    RC4_Receive_PDO_Mapping_Physical_outputs_60FE_01 : UDINT;
    RC4_Transmit_PDO_Mapping_StatusWord_6041_00 : UINT;
    RC4_Transmit_PDO_Mapping_Position_actual_value_6064_00 : DINT;
    RC4_Transmit_PDO_Mapping_Mode_of_operation_display_6061_00 : SINT;
    RC4_Transmit_PDO_Mapping_Following_error_actual_valu_60F4_00 : DINT;
    RC4_Transmit_PDO_Mapping_Torque_actual_value_6077_00 : INT;
    RC4_Transmit_PDO_Mapping_Digital_inputs_60FD_00 : UDINT;
    RC4_Transmit_PDO_Mapping_Error_code_603F_00 : UINT;
    RC5_Receive_PDO_Mapping_ControlWord_6040_00 : UINT;
    RC5_Receive_PDO_Mapping_Target_Position_607A_00 : DINT;
    RC5_Receive_PDO_Mapping_Mode_of_operation_6060_00 : SINT;
    RC5_Receive_PDO_Mapping_Profile_velocity_6081_00 : UDINT;
    RC5_Receive_PDO_Mapping_Profile_acceleration_6083_00 : UDINT;
    RC5_Receive_PDO_Mapping_Profile_deceleration_6084_00 : UDINT;
    RC5_Receive_PDO_Mapping_Physical_outputs_60FE_01 : UDINT;
    RC5_Transmit_PDO_Mapping_StatusWord_6041_00 : UINT;
    RC5_Transmit_PDO_Mapping_Position_actual_value_6064_00 : DINT;
    RC5_Transmit_PDO_Mapping_Mode_of_operation_display_6061_00 : SINT;
    RC5_Transmit_PDO_Mapping_Following_error_actual_valu_60F4_00 : DINT;
    RC5_Transmit_PDO_Mapping_Torque_actual_value_6077_00 : INT;
    RC5_Transmit_PDO_Mapping_Digital_inputs_60FD_00 : UDINT;
    RC5_Transmit_PDO_Mapping_Error_code_603F_00 : UINT;
    RC6_Receive_PDO_Mapping_ControlWord_6040_00 : UINT;
    RC6_Receive_PDO_Mapping_ControlWord_6040_00_1 : UINT;
    RC6_Receive_PDO_Mapping_Target_Position_607A_00 : DINT;
    RC6_Receive_PDO_Mapping_Mode_of_operation_6060_00 : SINT;
    RC6_Receive_PDO_Mapping_Profile_velocity_6081_00 : UDINT;
    RC6_Receive_PDO_Mapping_Profile_acceleration_6083_00 : UDINT;
    RC6_Receive_PDO_Mapping_Profile_deceleration_6084_00 : UDINT;
    RC6_Receive_PDO_Mapping_Physical_outputs_60FE_01 : UDINT;
    RC6_Transmit_PDO_Mapping_StatusWord_6041_00 : UINT;
    RC6_Transmit_PDO_Mapping_Position_actual_value_6064_00 : DINT;
    RC6_Transmit_PDO_Mapping_Mode_of_operation_display_6061_00 : SINT;
    RC6_Transmit_PDO_Mapping_Following_error_actual_valu_60F4_00 : DINT;
    RC6_Transmit_PDO_Mapping_Torque_actual_value_6077_00 : INT;
    RC6_Transmit_PDO_Mapping_Digital_inputs_60FD_00 : UDINT;
    RC6_Transmit_PDO_Mapping_Error_code_603F_00 : UINT;
    RCON1_OUT : ARRAY[1..6] OF ST_RCON_Direct_OUT_Axis;  (* RCON1 6軸分 PLC→RCON 指令（内部変数・通信変換は別途） *)
    RCON1_IN : ARRAY[1..6] OF ST_RCON_Direct_IN_Axis;  (* RCON1 6軸分 RCON→PLC 取得値・状態（内部変数・通信変換は別途） *)
    RCON1_SpeedUnit_mm_s : LREAL;  (* RCON1 速度の1カウント量mm/s。実機設定1.0または0.1を確認。未確認・0では使用しない。 *)
    RCON1_OUT_GwControl0Raw : UINT;  (* RCON1 PLC→RCON 【OUT00】共通 ゲートウェイ制御信号0（MON等）（未割付・直接数値指定の設計用） *)
    RCON1_OUT_GwControl1ReservedRaw : UINT;  (* RCON1 PLC→RCON 【OUT01】共通 ゲートウェイ制御信号1（予約・使用禁止）（未割付・直接数値指定の設計用） *)
    RCON1_OUT_ReservedOut02Raw : UINT;  (* RCON1 PLC→RCON 【OUT02】共通 共通予約領域（使用禁止・占有あり）（未割付・直接数値指定の設計用） *)
    RCON1_OUT_ReservedOut03Raw : UINT;  (* RCON1 PLC→RCON 【OUT03】共通 共通予約領域（使用禁止・占有あり）（未割付・直接数値指定の設計用） *)
    RCON1_OUT_ReservedOut04Raw : UINT;  (* RCON1 PLC→RCON 【OUT04】共通 共通予約領域（使用禁止・占有あり）（未割付・直接数値指定の設計用） *)
    RCON1_OUT_ReservedOut05Raw : UINT;  (* RCON1 PLC→RCON 【OUT05】共通 共通予約領域（使用禁止・占有あり）（未割付・直接数値指定の設計用） *)
    RCON1_OUT_ReservedOut06Raw : UINT;  (* RCON1 PLC→RCON 【OUT06】共通 共通予約領域（使用禁止・占有あり）（未割付・直接数値指定の設計用） *)
    RCON1_OUT_ReservedOut07Raw : UINT;  (* RCON1 PLC→RCON 【OUT07】共通 共通予約領域（使用禁止・占有あり）（未割付・直接数値指定の設計用） *)
    RCON1_OUT_Axis1_TargetPosLoRaw : UINT;  (* RCON1 PLC→RCON 【OUT08】1軸目（No.0） 目標位置 下位ワード（未割付・直接数値指定の設計用） *)
    RCON1_OUT_Axis1_TargetPosHiRaw : UINT;  (* RCON1 PLC→RCON 【OUT09】1軸目（No.0） 目標位置 上位ワード（未割付・直接数値指定の設計用） *)
    RCON1_OUT_Axis1_PositionBandLoRaw : UINT;  (* RCON1 PLC→RCON 【OUT10】1軸目（No.0） 位置決め幅 下位ワード（未割付・直接数値指定の設計用） *)
    RCON1_OUT_Axis1_PositionBandHiRaw : UINT;  (* RCON1 PLC→RCON 【OUT11】1軸目（No.0） 位置決め幅 上位ワード（未割付・直接数値指定の設計用） *)
    RCON1_OUT_Axis1_SpeedRaw : UINT;  (* RCON1 PLC→RCON 【OUT12】1軸目（No.0） 速度指令（未割付・直接数値指定の設計用） *)
    RCON1_OUT_Axis1_AccDecRaw : UINT;  (* RCON1 PLC→RCON 【OUT13】1軸目（No.0） 加減速度指令（加速・減速共通）（未割付・直接数値指定の設計用） *)
    RCON1_OUT_Axis1_PushLimitRaw : UINT;  (* RCON1 PLC→RCON 【OUT14】1軸目（No.0） 押付け電流制限値（未割付・直接数値指定の設計用） *)
    RCON1_OUT_Axis1_ControlRaw : UINT;  (* RCON1 PLC→RCON 【OUT15】1軸目（No.0） 軸制御信号（DSTR・SON等）（未割付・直接数値指定の設計用） *)
    RCON1_OUT_Axis2_TargetPosLoRaw : UINT;  (* RCON1 PLC→RCON 【OUT16】2軸目（No.1） 目標位置 下位ワード（未割付・直接数値指定の設計用） *)
    RCON1_OUT_Axis2_TargetPosHiRaw : UINT;  (* RCON1 PLC→RCON 【OUT17】2軸目（No.1） 目標位置 上位ワード（未割付・直接数値指定の設計用） *)
    RCON1_OUT_Axis2_PositionBandLoRaw : UINT;  (* RCON1 PLC→RCON 【OUT18】2軸目（No.1） 位置決め幅 下位ワード（未割付・直接数値指定の設計用） *)
    RCON1_OUT_Axis2_PositionBandHiRaw : UINT;  (* RCON1 PLC→RCON 【OUT19】2軸目（No.1） 位置決め幅 上位ワード（未割付・直接数値指定の設計用） *)
    RCON1_OUT_Axis2_SpeedRaw : UINT;  (* RCON1 PLC→RCON 【OUT20】2軸目（No.1） 速度指令（未割付・直接数値指定の設計用） *)
    RCON1_OUT_Axis2_AccDecRaw : UINT;  (* RCON1 PLC→RCON 【OUT21】2軸目（No.1） 加減速度指令（加速・減速共通）（未割付・直接数値指定の設計用） *)
    RCON1_OUT_Axis2_PushLimitRaw : UINT;  (* RCON1 PLC→RCON 【OUT22】2軸目（No.1） 押付け電流制限値（未割付・直接数値指定の設計用） *)
    RCON1_OUT_Axis2_ControlRaw : UINT;  (* RCON1 PLC→RCON 【OUT23】2軸目（No.1） 軸制御信号（DSTR・SON等）（未割付・直接数値指定の設計用） *)
    RCON1_OUT_Axis3_TargetPosLoRaw : UINT;  (* RCON1 PLC→RCON 【OUT24】3軸目（No.2） 目標位置 下位ワード（未割付・直接数値指定の設計用） *)
    RCON1_OUT_Axis3_TargetPosHiRaw : UINT;  (* RCON1 PLC→RCON 【OUT25】3軸目（No.2） 目標位置 上位ワード（未割付・直接数値指定の設計用） *)
    RCON1_OUT_Axis3_PositionBandLoRaw : UINT;  (* RCON1 PLC→RCON 【OUT26】3軸目（No.2） 位置決め幅 下位ワード（未割付・直接数値指定の設計用） *)
    RCON1_OUT_Axis3_PositionBandHiRaw : UINT;  (* RCON1 PLC→RCON 【OUT27】3軸目（No.2） 位置決め幅 上位ワード（未割付・直接数値指定の設計用） *)
    RCON1_OUT_Axis3_SpeedRaw : UINT;  (* RCON1 PLC→RCON 【OUT28】3軸目（No.2） 速度指令（未割付・直接数値指定の設計用） *)
    RCON1_OUT_Axis3_AccDecRaw : UINT;  (* RCON1 PLC→RCON 【OUT29】3軸目（No.2） 加減速度指令（加速・減速共通）（未割付・直接数値指定の設計用） *)
    RCON1_OUT_Axis3_PushLimitRaw : UINT;  (* RCON1 PLC→RCON 【OUT30】3軸目（No.2） 押付け電流制限値（未割付・直接数値指定の設計用） *)
    RCON1_OUT_Axis3_ControlRaw : UINT;  (* RCON1 PLC→RCON 【OUT31】3軸目（No.2） 軸制御信号（DSTR・SON等）（未割付・直接数値指定の設計用） *)
    RCON1_OUT_Axis4_TargetPosLoRaw : UINT;  (* RCON1 PLC→RCON 【OUT32】4軸目（No.3） 目標位置 下位ワード（未割付・直接数値指定の設計用） *)
    RCON1_OUT_Axis4_TargetPosHiRaw : UINT;  (* RCON1 PLC→RCON 【OUT33】4軸目（No.3） 目標位置 上位ワード（未割付・直接数値指定の設計用） *)
    RCON1_OUT_Axis4_PositionBandLoRaw : UINT;  (* RCON1 PLC→RCON 【OUT34】4軸目（No.3） 位置決め幅 下位ワード（未割付・直接数値指定の設計用） *)
    RCON1_OUT_Axis4_PositionBandHiRaw : UINT;  (* RCON1 PLC→RCON 【OUT35】4軸目（No.3） 位置決め幅 上位ワード（未割付・直接数値指定の設計用） *)
    RCON1_OUT_Axis4_SpeedRaw : UINT;  (* RCON1 PLC→RCON 【OUT36】4軸目（No.3） 速度指令（未割付・直接数値指定の設計用） *)
    RCON1_OUT_Axis4_AccDecRaw : UINT;  (* RCON1 PLC→RCON 【OUT37】4軸目（No.3） 加減速度指令（加速・減速共通）（未割付・直接数値指定の設計用） *)
    RCON1_OUT_Axis4_PushLimitRaw : UINT;  (* RCON1 PLC→RCON 【OUT38】4軸目（No.3） 押付け電流制限値（未割付・直接数値指定の設計用） *)
    RCON1_OUT_Axis4_ControlRaw : UINT;  (* RCON1 PLC→RCON 【OUT39】4軸目（No.3） 軸制御信号（DSTR・SON等）（未割付・直接数値指定の設計用） *)
    RCON1_OUT_Axis5_TargetPosLoRaw : UINT;  (* RCON1 PLC→RCON 【OUT40】5軸目（No.4） 目標位置 下位ワード（未割付・直接数値指定の設計用） *)
    RCON1_OUT_Axis5_TargetPosHiRaw : UINT;  (* RCON1 PLC→RCON 【OUT41】5軸目（No.4） 目標位置 上位ワード（未割付・直接数値指定の設計用） *)
    RCON1_OUT_Axis5_PositionBandLoRaw : UINT;  (* RCON1 PLC→RCON 【OUT42】5軸目（No.4） 位置決め幅 下位ワード（未割付・直接数値指定の設計用） *)
    RCON1_OUT_Axis5_PositionBandHiRaw : UINT;  (* RCON1 PLC→RCON 【OUT43】5軸目（No.4） 位置決め幅 上位ワード（未割付・直接数値指定の設計用） *)
    RCON1_OUT_Axis5_SpeedRaw : UINT;  (* RCON1 PLC→RCON 【OUT44】5軸目（No.4） 速度指令（未割付・直接数値指定の設計用） *)
    RCON1_OUT_Axis5_AccDecRaw : UINT;  (* RCON1 PLC→RCON 【OUT45】5軸目（No.4） 加減速度指令（加速・減速共通）（未割付・直接数値指定の設計用） *)
    RCON1_OUT_Axis5_PushLimitRaw : UINT;  (* RCON1 PLC→RCON 【OUT46】5軸目（No.4） 押付け電流制限値（未割付・直接数値指定の設計用） *)
    RCON1_OUT_Axis5_ControlRaw : UINT;  (* RCON1 PLC→RCON 【OUT47】5軸目（No.4） 軸制御信号（DSTR・SON等）（未割付・直接数値指定の設計用） *)
    RCON1_OUT_Axis6_TargetPosLoRaw : UINT;  (* RCON1 PLC→RCON 【OUT48】6軸目（No.5） 目標位置 下位ワード（未割付・直接数値指定の設計用） *)
    RCON1_OUT_Axis6_TargetPosHiRaw : UINT;  (* RCON1 PLC→RCON 【OUT49】6軸目（No.5） 目標位置 上位ワード（未割付・直接数値指定の設計用） *)
    RCON1_OUT_Axis6_PositionBandLoRaw : UINT;  (* RCON1 PLC→RCON 【OUT50】6軸目（No.5） 位置決め幅 下位ワード（未割付・直接数値指定の設計用） *)
    RCON1_OUT_Axis6_PositionBandHiRaw : UINT;  (* RCON1 PLC→RCON 【OUT51】6軸目（No.5） 位置決め幅 上位ワード（未割付・直接数値指定の設計用） *)
    RCON1_OUT_Axis6_SpeedRaw : UINT;  (* RCON1 PLC→RCON 【OUT52】6軸目（No.5） 速度指令（未割付・直接数値指定の設計用） *)
    RCON1_OUT_Axis6_AccDecRaw : UINT;  (* RCON1 PLC→RCON 【OUT53】6軸目（No.5） 加減速度指令（加速・減速共通）（未割付・直接数値指定の設計用） *)
    RCON1_OUT_Axis6_PushLimitRaw : UINT;  (* RCON1 PLC→RCON 【OUT54】6軸目（No.5） 押付け電流制限値（未割付・直接数値指定の設計用） *)
    RCON1_OUT_Axis6_ControlRaw : UINT;  (* RCON1 PLC→RCON 【OUT55】6軸目（No.5） 軸制御信号（DSTR・SON等）（未割付・直接数値指定の設計用） *)
    RCON1_IN_GwStatus0Raw : UINT;  (* RCON1 RCON→PLC 【IN00】共通 ゲートウェイ状態信号0（未割付・直接数値指定の設計用） *)
    RCON1_IN_AxisLinkStatusRaw : UINT;  (* RCON1 RCON→PLC 【IN01】共通 ゲートウェイ状態信号1（軸No.0～15リンク状態）（未割付・直接数値指定の設計用） *)
    RCON1_IN_PowerStatus0Raw : UINT;  (* RCON1 RCON→PLC 【IN02】共通 電源ユニット状態信号0（未割付・直接数値指定の設計用） *)
    RCON1_IN_PowerStatus1Raw : UINT;  (* RCON1 RCON→PLC 【IN03】共通 電源ユニット状態信号1（未割付・直接数値指定の設計用） *)
    RCON1_IN_PowerStatus2Raw : UINT;  (* RCON1 RCON→PLC 【IN04】共通 電源ユニット状態信号2（未割付・直接数値指定の設計用） *)
    RCON1_IN_PowerStatus3Raw : UINT;  (* RCON1 RCON→PLC 【IN05】共通 電源ユニット状態信号3（未割付・直接数値指定の設計用） *)
    RCON1_IN_PowerStatus4MaintenanceRaw : UINT;  (* RCON1 RCON→PLC 【IN06】共通 電源ユニット状態信号4／軽故障メンテナンス（設定依存）（未割付・直接数値指定の設計用） *)
    RCON1_IN_ReservedIn07Raw : UINT;  (* RCON1 RCON→PLC 【IN07】共通 共通予約領域（使用禁止・占有あり）（未割付・直接数値指定の設計用） *)
    RCON1_IN_Axis1_ActualPosLoRaw : UINT;  (* RCON1 RCON→PLC 【IN08】1軸目（No.0） 現在位置 下位ワード（未割付・直接数値指定の設計用） *)
    RCON1_IN_Axis1_ActualPosHiRaw : UINT;  (* RCON1 RCON→PLC 【IN09】1軸目（No.0） 現在位置 上位ワード（未割付・直接数値指定の設計用） *)
    RCON1_IN_Axis1_CurrentLoRaw : UINT;  (* RCON1 RCON→PLC 【IN10】1軸目（No.0） 現在電流 下位ワード（PCは指令電流）（未割付・直接数値指定の設計用） *)
    RCON1_IN_Axis1_CurrentHiRaw : UINT;  (* RCON1 RCON→PLC 【IN11】1軸目（No.0） 現在電流 上位ワード（PCは指令電流）（未割付・直接数値指定の設計用） *)
    RCON1_IN_Axis1_ActualSpeedRaw : UINT;  (* RCON1 RCON→PLC 【IN12】1軸目（No.0） 現在速度（負方向は2の補数）（未割付・直接数値指定の設計用） *)
    RCON1_IN_Axis1_ReservedInRaw : UINT;  (* RCON1 RCON→PLC 【IN13】1軸目（No.0） 予約領域（使用禁止）（未割付・直接数値指定の設計用） *)
    RCON1_IN_Axis1_AlarmCodeRaw : UINT;  (* RCON1 RCON→PLC 【IN14】1軸目（No.0） アラームコード（簡易コードではない）（未割付・直接数値指定の設計用） *)
    RCON1_IN_Axis1_StatusRaw : UINT;  (* RCON1 RCON→PLC 【IN15】1軸目（No.0） 軸状態信号（PEND・SV等）（未割付・直接数値指定の設計用） *)
    RCON1_IN_Axis2_ActualPosLoRaw : UINT;  (* RCON1 RCON→PLC 【IN16】2軸目（No.1） 現在位置 下位ワード（未割付・直接数値指定の設計用） *)
    RCON1_IN_Axis2_ActualPosHiRaw : UINT;  (* RCON1 RCON→PLC 【IN17】2軸目（No.1） 現在位置 上位ワード（未割付・直接数値指定の設計用） *)
    RCON1_IN_Axis2_CurrentLoRaw : UINT;  (* RCON1 RCON→PLC 【IN18】2軸目（No.1） 現在電流 下位ワード（PCは指令電流）（未割付・直接数値指定の設計用） *)
    RCON1_IN_Axis2_CurrentHiRaw : UINT;  (* RCON1 RCON→PLC 【IN19】2軸目（No.1） 現在電流 上位ワード（PCは指令電流）（未割付・直接数値指定の設計用） *)
    RCON1_IN_Axis2_ActualSpeedRaw : UINT;  (* RCON1 RCON→PLC 【IN20】2軸目（No.1） 現在速度（負方向は2の補数）（未割付・直接数値指定の設計用） *)
    RCON1_IN_Axis2_ReservedInRaw : UINT;  (* RCON1 RCON→PLC 【IN21】2軸目（No.1） 予約領域（使用禁止）（未割付・直接数値指定の設計用） *)
    RCON1_IN_Axis2_AlarmCodeRaw : UINT;  (* RCON1 RCON→PLC 【IN22】2軸目（No.1） アラームコード（簡易コードではない）（未割付・直接数値指定の設計用） *)
    RCON1_IN_Axis2_StatusRaw : UINT;  (* RCON1 RCON→PLC 【IN23】2軸目（No.1） 軸状態信号（PEND・SV等）（未割付・直接数値指定の設計用） *)
    RCON1_IN_Axis3_ActualPosLoRaw : UINT;  (* RCON1 RCON→PLC 【IN24】3軸目（No.2） 現在位置 下位ワード（未割付・直接数値指定の設計用） *)
    RCON1_IN_Axis3_ActualPosHiRaw : UINT;  (* RCON1 RCON→PLC 【IN25】3軸目（No.2） 現在位置 上位ワード（未割付・直接数値指定の設計用） *)
    RCON1_IN_Axis3_CurrentLoRaw : UINT;  (* RCON1 RCON→PLC 【IN26】3軸目（No.2） 現在電流 下位ワード（PCは指令電流）（未割付・直接数値指定の設計用） *)
    RCON1_IN_Axis3_CurrentHiRaw : UINT;  (* RCON1 RCON→PLC 【IN27】3軸目（No.2） 現在電流 上位ワード（PCは指令電流）（未割付・直接数値指定の設計用） *)
    RCON1_IN_Axis3_ActualSpeedRaw : UINT;  (* RCON1 RCON→PLC 【IN28】3軸目（No.2） 現在速度（負方向は2の補数）（未割付・直接数値指定の設計用） *)
    RCON1_IN_Axis3_ReservedInRaw : UINT;  (* RCON1 RCON→PLC 【IN29】3軸目（No.2） 予約領域（使用禁止）（未割付・直接数値指定の設計用） *)
    RCON1_IN_Axis3_AlarmCodeRaw : UINT;  (* RCON1 RCON→PLC 【IN30】3軸目（No.2） アラームコード（簡易コードではない）（未割付・直接数値指定の設計用） *)
    RCON1_IN_Axis3_StatusRaw : UINT;  (* RCON1 RCON→PLC 【IN31】3軸目（No.2） 軸状態信号（PEND・SV等）（未割付・直接数値指定の設計用） *)
    RCON1_IN_Axis4_ActualPosLoRaw : UINT;  (* RCON1 RCON→PLC 【IN32】4軸目（No.3） 現在位置 下位ワード（未割付・直接数値指定の設計用） *)
    RCON1_IN_Axis4_ActualPosHiRaw : UINT;  (* RCON1 RCON→PLC 【IN33】4軸目（No.3） 現在位置 上位ワード（未割付・直接数値指定の設計用） *)
    RCON1_IN_Axis4_CurrentLoRaw : UINT;  (* RCON1 RCON→PLC 【IN34】4軸目（No.3） 現在電流 下位ワード（PCは指令電流）（未割付・直接数値指定の設計用） *)
    RCON1_IN_Axis4_CurrentHiRaw : UINT;  (* RCON1 RCON→PLC 【IN35】4軸目（No.3） 現在電流 上位ワード（PCは指令電流）（未割付・直接数値指定の設計用） *)
    RCON1_IN_Axis4_ActualSpeedRaw : UINT;  (* RCON1 RCON→PLC 【IN36】4軸目（No.3） 現在速度（負方向は2の補数）（未割付・直接数値指定の設計用） *)
    RCON1_IN_Axis4_ReservedInRaw : UINT;  (* RCON1 RCON→PLC 【IN37】4軸目（No.3） 予約領域（使用禁止）（未割付・直接数値指定の設計用） *)
    RCON1_IN_Axis4_AlarmCodeRaw : UINT;  (* RCON1 RCON→PLC 【IN38】4軸目（No.3） アラームコード（簡易コードではない）（未割付・直接数値指定の設計用） *)
    RCON1_IN_Axis4_StatusRaw : UINT;  (* RCON1 RCON→PLC 【IN39】4軸目（No.3） 軸状態信号（PEND・SV等）（未割付・直接数値指定の設計用） *)
    RCON1_IN_Axis5_ActualPosLoRaw : UINT;  (* RCON1 RCON→PLC 【IN40】5軸目（No.4） 現在位置 下位ワード（未割付・直接数値指定の設計用） *)
    RCON1_IN_Axis5_ActualPosHiRaw : UINT;  (* RCON1 RCON→PLC 【IN41】5軸目（No.4） 現在位置 上位ワード（未割付・直接数値指定の設計用） *)
    RCON1_IN_Axis5_CurrentLoRaw : UINT;  (* RCON1 RCON→PLC 【IN42】5軸目（No.4） 現在電流 下位ワード（PCは指令電流）（未割付・直接数値指定の設計用） *)
    RCON1_IN_Axis5_CurrentHiRaw : UINT;  (* RCON1 RCON→PLC 【IN43】5軸目（No.4） 現在電流 上位ワード（PCは指令電流）（未割付・直接数値指定の設計用） *)
    RCON1_IN_Axis5_ActualSpeedRaw : UINT;  (* RCON1 RCON→PLC 【IN44】5軸目（No.4） 現在速度（負方向は2の補数）（未割付・直接数値指定の設計用） *)
    RCON1_IN_Axis5_ReservedInRaw : UINT;  (* RCON1 RCON→PLC 【IN45】5軸目（No.4） 予約領域（使用禁止）（未割付・直接数値指定の設計用） *)
    RCON1_IN_Axis5_AlarmCodeRaw : UINT;  (* RCON1 RCON→PLC 【IN46】5軸目（No.4） アラームコード（簡易コードではない）（未割付・直接数値指定の設計用） *)
    RCON1_IN_Axis5_StatusRaw : UINT;  (* RCON1 RCON→PLC 【IN47】5軸目（No.4） 軸状態信号（PEND・SV等）（未割付・直接数値指定の設計用） *)
    RCON1_IN_Axis6_ActualPosLoRaw : UINT;  (* RCON1 RCON→PLC 【IN48】6軸目（No.5） 現在位置 下位ワード（未割付・直接数値指定の設計用） *)
    RCON1_IN_Axis6_ActualPosHiRaw : UINT;  (* RCON1 RCON→PLC 【IN49】6軸目（No.5） 現在位置 上位ワード（未割付・直接数値指定の設計用） *)
    RCON1_IN_Axis6_CurrentLoRaw : UINT;  (* RCON1 RCON→PLC 【IN50】6軸目（No.5） 現在電流 下位ワード（PCは指令電流）（未割付・直接数値指定の設計用） *)
    RCON1_IN_Axis6_CurrentHiRaw : UINT;  (* RCON1 RCON→PLC 【IN51】6軸目（No.5） 現在電流 上位ワード（PCは指令電流）（未割付・直接数値指定の設計用） *)
    RCON1_IN_Axis6_ActualSpeedRaw : UINT;  (* RCON1 RCON→PLC 【IN52】6軸目（No.5） 現在速度（負方向は2の補数）（未割付・直接数値指定の設計用） *)
    RCON1_IN_Axis6_ReservedInRaw : UINT;  (* RCON1 RCON→PLC 【IN53】6軸目（No.5） 予約領域（使用禁止）（未割付・直接数値指定の設計用） *)
    RCON1_IN_Axis6_AlarmCodeRaw : UINT;  (* RCON1 RCON→PLC 【IN54】6軸目（No.5） アラームコード（簡易コードではない）（未割付・直接数値指定の設計用） *)
    RCON1_IN_Axis6_StatusRaw : UINT;  (* RCON1 RCON→PLC 【IN55】6軸目（No.5） 軸状態信号（PEND・SV等）（未割付・直接数値指定の設計用） *)
    RCON2_OUT : ARRAY[1..5] OF ST_RCON_Direct_OUT_Axis;  (* RCON2 5軸分 PLC→RCON 指令（内部変数・通信変換は別途） *)
    RCON2_IN : ARRAY[1..5] OF ST_RCON_Direct_IN_Axis;  (* RCON2 5軸分 RCON→PLC 取得値・状態（内部変数・通信変換は別途） *)
    RCON2_SpeedUnit_mm_s : LREAL;  (* RCON2 速度の1カウント量mm/s。実機設定1.0または0.1を確認。未確認・0では使用しない。 *)
    RCON2_OUT_GwControl0Raw : UINT;  (* RCON2 PLC→RCON 【OUT00】共通 ゲートウェイ制御信号0（MON等）（未割付・直接数値指定の設計用） *)
    RCON2_OUT_GwControl1ReservedRaw : UINT;  (* RCON2 PLC→RCON 【OUT01】共通 ゲートウェイ制御信号1（予約・使用禁止）（未割付・直接数値指定の設計用） *)
    RCON2_OUT_ReservedOut02Raw : UINT;  (* RCON2 PLC→RCON 【OUT02】共通 共通予約領域（使用禁止・占有あり）（未割付・直接数値指定の設計用） *)
    RCON2_OUT_ReservedOut03Raw : UINT;  (* RCON2 PLC→RCON 【OUT03】共通 共通予約領域（使用禁止・占有あり）（未割付・直接数値指定の設計用） *)
    RCON2_OUT_ReservedOut04Raw : UINT;  (* RCON2 PLC→RCON 【OUT04】共通 共通予約領域（使用禁止・占有あり）（未割付・直接数値指定の設計用） *)
    RCON2_OUT_ReservedOut05Raw : UINT;  (* RCON2 PLC→RCON 【OUT05】共通 共通予約領域（使用禁止・占有あり）（未割付・直接数値指定の設計用） *)
    RCON2_OUT_ReservedOut06Raw : UINT;  (* RCON2 PLC→RCON 【OUT06】共通 共通予約領域（使用禁止・占有あり）（未割付・直接数値指定の設計用） *)
    RCON2_OUT_ReservedOut07Raw : UINT;  (* RCON2 PLC→RCON 【OUT07】共通 共通予約領域（使用禁止・占有あり）（未割付・直接数値指定の設計用） *)
    RCON2_OUT_Axis1_TargetPosLoRaw : UINT;  (* RCON2 PLC→RCON 【OUT08】1軸目（No.0） 目標位置 下位ワード（未割付・直接数値指定の設計用） *)
    RCON2_OUT_Axis1_TargetPosHiRaw : UINT;  (* RCON2 PLC→RCON 【OUT09】1軸目（No.0） 目標位置 上位ワード（未割付・直接数値指定の設計用） *)
    RCON2_OUT_Axis1_PositionBandLoRaw : UINT;  (* RCON2 PLC→RCON 【OUT10】1軸目（No.0） 位置決め幅 下位ワード（未割付・直接数値指定の設計用） *)
    RCON2_OUT_Axis1_PositionBandHiRaw : UINT;  (* RCON2 PLC→RCON 【OUT11】1軸目（No.0） 位置決め幅 上位ワード（未割付・直接数値指定の設計用） *)
    RCON2_OUT_Axis1_SpeedRaw : UINT;  (* RCON2 PLC→RCON 【OUT12】1軸目（No.0） 速度指令（未割付・直接数値指定の設計用） *)
    RCON2_OUT_Axis1_AccDecRaw : UINT;  (* RCON2 PLC→RCON 【OUT13】1軸目（No.0） 加減速度指令（加速・減速共通）（未割付・直接数値指定の設計用） *)
    RCON2_OUT_Axis1_PushLimitRaw : UINT;  (* RCON2 PLC→RCON 【OUT14】1軸目（No.0） 押付け電流制限値（未割付・直接数値指定の設計用） *)
    RCON2_OUT_Axis1_ControlRaw : UINT;  (* RCON2 PLC→RCON 【OUT15】1軸目（No.0） 軸制御信号（DSTR・SON等）（未割付・直接数値指定の設計用） *)
    RCON2_OUT_Axis2_TargetPosLoRaw : UINT;  (* RCON2 PLC→RCON 【OUT16】2軸目（No.1） 目標位置 下位ワード（未割付・直接数値指定の設計用） *)
    RCON2_OUT_Axis2_TargetPosHiRaw : UINT;  (* RCON2 PLC→RCON 【OUT17】2軸目（No.1） 目標位置 上位ワード（未割付・直接数値指定の設計用） *)
    RCON2_OUT_Axis2_PositionBandLoRaw : UINT;  (* RCON2 PLC→RCON 【OUT18】2軸目（No.1） 位置決め幅 下位ワード（未割付・直接数値指定の設計用） *)
    RCON2_OUT_Axis2_PositionBandHiRaw : UINT;  (* RCON2 PLC→RCON 【OUT19】2軸目（No.1） 位置決め幅 上位ワード（未割付・直接数値指定の設計用） *)
    RCON2_OUT_Axis2_SpeedRaw : UINT;  (* RCON2 PLC→RCON 【OUT20】2軸目（No.1） 速度指令（未割付・直接数値指定の設計用） *)
    RCON2_OUT_Axis2_AccDecRaw : UINT;  (* RCON2 PLC→RCON 【OUT21】2軸目（No.1） 加減速度指令（加速・減速共通）（未割付・直接数値指定の設計用） *)
    RCON2_OUT_Axis2_PushLimitRaw : UINT;  (* RCON2 PLC→RCON 【OUT22】2軸目（No.1） 押付け電流制限値（未割付・直接数値指定の設計用） *)
    RCON2_OUT_Axis2_ControlRaw : UINT;  (* RCON2 PLC→RCON 【OUT23】2軸目（No.1） 軸制御信号（DSTR・SON等）（未割付・直接数値指定の設計用） *)
    RCON2_OUT_Axis3_TargetPosLoRaw : UINT;  (* RCON2 PLC→RCON 【OUT24】3軸目（No.2） 目標位置 下位ワード（未割付・直接数値指定の設計用） *)
    RCON2_OUT_Axis3_TargetPosHiRaw : UINT;  (* RCON2 PLC→RCON 【OUT25】3軸目（No.2） 目標位置 上位ワード（未割付・直接数値指定の設計用） *)
    RCON2_OUT_Axis3_PositionBandLoRaw : UINT;  (* RCON2 PLC→RCON 【OUT26】3軸目（No.2） 位置決め幅 下位ワード（未割付・直接数値指定の設計用） *)
    RCON2_OUT_Axis3_PositionBandHiRaw : UINT;  (* RCON2 PLC→RCON 【OUT27】3軸目（No.2） 位置決め幅 上位ワード（未割付・直接数値指定の設計用） *)
    RCON2_OUT_Axis3_SpeedRaw : UINT;  (* RCON2 PLC→RCON 【OUT28】3軸目（No.2） 速度指令（未割付・直接数値指定の設計用） *)
    RCON2_OUT_Axis3_AccDecRaw : UINT;  (* RCON2 PLC→RCON 【OUT29】3軸目（No.2） 加減速度指令（加速・減速共通）（未割付・直接数値指定の設計用） *)
    RCON2_OUT_Axis3_PushLimitRaw : UINT;  (* RCON2 PLC→RCON 【OUT30】3軸目（No.2） 押付け電流制限値（未割付・直接数値指定の設計用） *)
    RCON2_OUT_Axis3_ControlRaw : UINT;  (* RCON2 PLC→RCON 【OUT31】3軸目（No.2） 軸制御信号（DSTR・SON等）（未割付・直接数値指定の設計用） *)
    RCON2_OUT_Axis4_TargetPosLoRaw : UINT;  (* RCON2 PLC→RCON 【OUT32】4軸目（No.3） 目標位置 下位ワード（未割付・直接数値指定の設計用） *)
    RCON2_OUT_Axis4_TargetPosHiRaw : UINT;  (* RCON2 PLC→RCON 【OUT33】4軸目（No.3） 目標位置 上位ワード（未割付・直接数値指定の設計用） *)
    RCON2_OUT_Axis4_PositionBandLoRaw : UINT;  (* RCON2 PLC→RCON 【OUT34】4軸目（No.3） 位置決め幅 下位ワード（未割付・直接数値指定の設計用） *)
    RCON2_OUT_Axis4_PositionBandHiRaw : UINT;  (* RCON2 PLC→RCON 【OUT35】4軸目（No.3） 位置決め幅 上位ワード（未割付・直接数値指定の設計用） *)
    RCON2_OUT_Axis4_SpeedRaw : UINT;  (* RCON2 PLC→RCON 【OUT36】4軸目（No.3） 速度指令（未割付・直接数値指定の設計用） *)
    RCON2_OUT_Axis4_AccDecRaw : UINT;  (* RCON2 PLC→RCON 【OUT37】4軸目（No.3） 加減速度指令（加速・減速共通）（未割付・直接数値指定の設計用） *)
    RCON2_OUT_Axis4_PushLimitRaw : UINT;  (* RCON2 PLC→RCON 【OUT38】4軸目（No.3） 押付け電流制限値（未割付・直接数値指定の設計用） *)
    RCON2_OUT_Axis4_ControlRaw : UINT;  (* RCON2 PLC→RCON 【OUT39】4軸目（No.3） 軸制御信号（DSTR・SON等）（未割付・直接数値指定の設計用） *)
    RCON2_OUT_Axis5_TargetPosLoRaw : UINT;  (* RCON2 PLC→RCON 【OUT40】5軸目（No.4） 目標位置 下位ワード（未割付・直接数値指定の設計用） *)
    RCON2_OUT_Axis5_TargetPosHiRaw : UINT;  (* RCON2 PLC→RCON 【OUT41】5軸目（No.4） 目標位置 上位ワード（未割付・直接数値指定の設計用） *)
    RCON2_OUT_Axis5_PositionBandLoRaw : UINT;  (* RCON2 PLC→RCON 【OUT42】5軸目（No.4） 位置決め幅 下位ワード（未割付・直接数値指定の設計用） *)
    RCON2_OUT_Axis5_PositionBandHiRaw : UINT;  (* RCON2 PLC→RCON 【OUT43】5軸目（No.4） 位置決め幅 上位ワード（未割付・直接数値指定の設計用） *)
    RCON2_OUT_Axis5_SpeedRaw : UINT;  (* RCON2 PLC→RCON 【OUT44】5軸目（No.4） 速度指令（未割付・直接数値指定の設計用） *)
    RCON2_OUT_Axis5_AccDecRaw : UINT;  (* RCON2 PLC→RCON 【OUT45】5軸目（No.4） 加減速度指令（加速・減速共通）（未割付・直接数値指定の設計用） *)
    RCON2_OUT_Axis5_PushLimitRaw : UINT;  (* RCON2 PLC→RCON 【OUT46】5軸目（No.4） 押付け電流制限値（未割付・直接数値指定の設計用） *)
    RCON2_OUT_Axis5_ControlRaw : UINT;  (* RCON2 PLC→RCON 【OUT47】5軸目（No.4） 軸制御信号（DSTR・SON等）（未割付・直接数値指定の設計用） *)
    RCON2_IN_GwStatus0Raw : UINT;  (* RCON2 RCON→PLC 【IN00】共通 ゲートウェイ状態信号0（未割付・直接数値指定の設計用） *)
    RCON2_IN_AxisLinkStatusRaw : UINT;  (* RCON2 RCON→PLC 【IN01】共通 ゲートウェイ状態信号1（軸No.0～15リンク状態）（未割付・直接数値指定の設計用） *)
    RCON2_IN_PowerStatus0Raw : UINT;  (* RCON2 RCON→PLC 【IN02】共通 電源ユニット状態信号0（未割付・直接数値指定の設計用） *)
    RCON2_IN_PowerStatus1Raw : UINT;  (* RCON2 RCON→PLC 【IN03】共通 電源ユニット状態信号1（未割付・直接数値指定の設計用） *)
    RCON2_IN_PowerStatus2Raw : UINT;  (* RCON2 RCON→PLC 【IN04】共通 電源ユニット状態信号2（未割付・直接数値指定の設計用） *)
    RCON2_IN_PowerStatus3Raw : UINT;  (* RCON2 RCON→PLC 【IN05】共通 電源ユニット状態信号3（未割付・直接数値指定の設計用） *)
    RCON2_IN_PowerStatus4MaintenanceRaw : UINT;  (* RCON2 RCON→PLC 【IN06】共通 電源ユニット状態信号4／軽故障メンテナンス（設定依存）（未割付・直接数値指定の設計用） *)
    RCON2_IN_ReservedIn07Raw : UINT;  (* RCON2 RCON→PLC 【IN07】共通 共通予約領域（使用禁止・占有あり）（未割付・直接数値指定の設計用） *)
    RCON2_IN_Axis1_ActualPosLoRaw : UINT;  (* RCON2 RCON→PLC 【IN08】1軸目（No.0） 現在位置 下位ワード（未割付・直接数値指定の設計用） *)
    RCON2_IN_Axis1_ActualPosHiRaw : UINT;  (* RCON2 RCON→PLC 【IN09】1軸目（No.0） 現在位置 上位ワード（未割付・直接数値指定の設計用） *)
    RCON2_IN_Axis1_CurrentLoRaw : UINT;  (* RCON2 RCON→PLC 【IN10】1軸目（No.0） 現在電流 下位ワード（PCは指令電流）（未割付・直接数値指定の設計用） *)
    RCON2_IN_Axis1_CurrentHiRaw : UINT;  (* RCON2 RCON→PLC 【IN11】1軸目（No.0） 現在電流 上位ワード（PCは指令電流）（未割付・直接数値指定の設計用） *)
    RCON2_IN_Axis1_ActualSpeedRaw : UINT;  (* RCON2 RCON→PLC 【IN12】1軸目（No.0） 現在速度（負方向は2の補数）（未割付・直接数値指定の設計用） *)
    RCON2_IN_Axis1_ReservedInRaw : UINT;  (* RCON2 RCON→PLC 【IN13】1軸目（No.0） 予約領域（使用禁止）（未割付・直接数値指定の設計用） *)
    RCON2_IN_Axis1_AlarmCodeRaw : UINT;  (* RCON2 RCON→PLC 【IN14】1軸目（No.0） アラームコード（簡易コードではない）（未割付・直接数値指定の設計用） *)
    RCON2_IN_Axis1_StatusRaw : UINT;  (* RCON2 RCON→PLC 【IN15】1軸目（No.0） 軸状態信号（PEND・SV等）（未割付・直接数値指定の設計用） *)
    RCON2_IN_Axis2_ActualPosLoRaw : UINT;  (* RCON2 RCON→PLC 【IN16】2軸目（No.1） 現在位置 下位ワード（未割付・直接数値指定の設計用） *)
    RCON2_IN_Axis2_ActualPosHiRaw : UINT;  (* RCON2 RCON→PLC 【IN17】2軸目（No.1） 現在位置 上位ワード（未割付・直接数値指定の設計用） *)
    RCON2_IN_Axis2_CurrentLoRaw : UINT;  (* RCON2 RCON→PLC 【IN18】2軸目（No.1） 現在電流 下位ワード（PCは指令電流）（未割付・直接数値指定の設計用） *)
    RCON2_IN_Axis2_CurrentHiRaw : UINT;  (* RCON2 RCON→PLC 【IN19】2軸目（No.1） 現在電流 上位ワード（PCは指令電流）（未割付・直接数値指定の設計用） *)
    RCON2_IN_Axis2_ActualSpeedRaw : UINT;  (* RCON2 RCON→PLC 【IN20】2軸目（No.1） 現在速度（負方向は2の補数）（未割付・直接数値指定の設計用） *)
    RCON2_IN_Axis2_ReservedInRaw : UINT;  (* RCON2 RCON→PLC 【IN21】2軸目（No.1） 予約領域（使用禁止）（未割付・直接数値指定の設計用） *)
    RCON2_IN_Axis2_AlarmCodeRaw : UINT;  (* RCON2 RCON→PLC 【IN22】2軸目（No.1） アラームコード（簡易コードではない）（未割付・直接数値指定の設計用） *)
    RCON2_IN_Axis2_StatusRaw : UINT;  (* RCON2 RCON→PLC 【IN23】2軸目（No.1） 軸状態信号（PEND・SV等）（未割付・直接数値指定の設計用） *)
    RCON2_IN_Axis3_ActualPosLoRaw : UINT;  (* RCON2 RCON→PLC 【IN24】3軸目（No.2） 現在位置 下位ワード（未割付・直接数値指定の設計用） *)
    RCON2_IN_Axis3_ActualPosHiRaw : UINT;  (* RCON2 RCON→PLC 【IN25】3軸目（No.2） 現在位置 上位ワード（未割付・直接数値指定の設計用） *)
    RCON2_IN_Axis3_CurrentLoRaw : UINT;  (* RCON2 RCON→PLC 【IN26】3軸目（No.2） 現在電流 下位ワード（PCは指令電流）（未割付・直接数値指定の設計用） *)
    RCON2_IN_Axis3_CurrentHiRaw : UINT;  (* RCON2 RCON→PLC 【IN27】3軸目（No.2） 現在電流 上位ワード（PCは指令電流）（未割付・直接数値指定の設計用） *)
    RCON2_IN_Axis3_ActualSpeedRaw : UINT;  (* RCON2 RCON→PLC 【IN28】3軸目（No.2） 現在速度（負方向は2の補数）（未割付・直接数値指定の設計用） *)
    RCON2_IN_Axis3_ReservedInRaw : UINT;  (* RCON2 RCON→PLC 【IN29】3軸目（No.2） 予約領域（使用禁止）（未割付・直接数値指定の設計用） *)
    RCON2_IN_Axis3_AlarmCodeRaw : UINT;  (* RCON2 RCON→PLC 【IN30】3軸目（No.2） アラームコード（簡易コードではない）（未割付・直接数値指定の設計用） *)
    RCON2_IN_Axis3_StatusRaw : UINT;  (* RCON2 RCON→PLC 【IN31】3軸目（No.2） 軸状態信号（PEND・SV等）（未割付・直接数値指定の設計用） *)
    RCON2_IN_Axis4_ActualPosLoRaw : UINT;  (* RCON2 RCON→PLC 【IN32】4軸目（No.3） 現在位置 下位ワード（未割付・直接数値指定の設計用） *)
    RCON2_IN_Axis4_ActualPosHiRaw : UINT;  (* RCON2 RCON→PLC 【IN33】4軸目（No.3） 現在位置 上位ワード（未割付・直接数値指定の設計用） *)
    RCON2_IN_Axis4_CurrentLoRaw : UINT;  (* RCON2 RCON→PLC 【IN34】4軸目（No.3） 現在電流 下位ワード（PCは指令電流）（未割付・直接数値指定の設計用） *)
    RCON2_IN_Axis4_CurrentHiRaw : UINT;  (* RCON2 RCON→PLC 【IN35】4軸目（No.3） 現在電流 上位ワード（PCは指令電流）（未割付・直接数値指定の設計用） *)
    RCON2_IN_Axis4_ActualSpeedRaw : UINT;  (* RCON2 RCON→PLC 【IN36】4軸目（No.3） 現在速度（負方向は2の補数）（未割付・直接数値指定の設計用） *)
    RCON2_IN_Axis4_ReservedInRaw : UINT;  (* RCON2 RCON→PLC 【IN37】4軸目（No.3） 予約領域（使用禁止）（未割付・直接数値指定の設計用） *)
    RCON2_IN_Axis4_AlarmCodeRaw : UINT;  (* RCON2 RCON→PLC 【IN38】4軸目（No.3） アラームコード（簡易コードではない）（未割付・直接数値指定の設計用） *)
    RCON2_IN_Axis4_StatusRaw : UINT;  (* RCON2 RCON→PLC 【IN39】4軸目（No.3） 軸状態信号（PEND・SV等）（未割付・直接数値指定の設計用） *)
    RCON2_IN_Axis5_ActualPosLoRaw : UINT;  (* RCON2 RCON→PLC 【IN40】5軸目（No.4） 現在位置 下位ワード（未割付・直接数値指定の設計用） *)
    RCON2_IN_Axis5_ActualPosHiRaw : UINT;  (* RCON2 RCON→PLC 【IN41】5軸目（No.4） 現在位置 上位ワード（未割付・直接数値指定の設計用） *)
    RCON2_IN_Axis5_CurrentLoRaw : UINT;  (* RCON2 RCON→PLC 【IN42】5軸目（No.4） 現在電流 下位ワード（PCは指令電流）（未割付・直接数値指定の設計用） *)
    RCON2_IN_Axis5_CurrentHiRaw : UINT;  (* RCON2 RCON→PLC 【IN43】5軸目（No.4） 現在電流 上位ワード（PCは指令電流）（未割付・直接数値指定の設計用） *)
    RCON2_IN_Axis5_ActualSpeedRaw : UINT;  (* RCON2 RCON→PLC 【IN44】5軸目（No.4） 現在速度（負方向は2の補数）（未割付・直接数値指定の設計用） *)
    RCON2_IN_Axis5_ReservedInRaw : UINT;  (* RCON2 RCON→PLC 【IN45】5軸目（No.4） 予約領域（使用禁止）（未割付・直接数値指定の設計用） *)
    RCON2_IN_Axis5_AlarmCodeRaw : UINT;  (* RCON2 RCON→PLC 【IN46】5軸目（No.4） アラームコード（簡易コードではない）（未割付・直接数値指定の設計用） *)
    RCON2_IN_Axis5_StatusRaw : UINT;  (* RCON2 RCON→PLC 【IN47】5軸目（No.4） 軸状態信号（PEND・SV等）（未割付・直接数値指定の設計用） *)
    E005_Out_OUT00_2003_01 : UINT;
    E005_Out_OUT01_2003_02 : UINT;
    E005_Out_OUT02_2003_03 : UINT;
    E005_Out_OUT03_2003_04 : UINT;
    E005_Out_OUT04_2003_05 : UINT;
    E005_Out_OUT05_2003_06 : UINT;
    E005_Out_OUT06_2003_07 : UINT;
    E005_Out_OUT07_2003_08 : UINT;
    E005_Out_OUT08_2003_09 : UINT;
    E005_Out_OUT09_2003_0A : UINT;
    E005_Out_OUT10_2003_0B : UINT;
    E005_Out_OUT11_2003_0C : UINT;
    E005_Out_OUT12_2003_0D : UINT;
    E005_Out_OUT13_2003_0E : UINT;
    E005_Out_OUT14_2003_0F : UINT;
    E005_Out_OUT15_2003_10 : UINT;
    E005_Out_OUT16_2003_11 : UINT;
    E005_Out_OUT17_2003_12 : UINT;
    E005_Out_OUT18_2003_13 : UINT;
    E005_Out_OUT19_2003_14 : UINT;
    E005_Out_OUT20_2003_15 : UINT;
    E005_Out_OUT21_2003_16 : UINT;
    E005_Out_OUT22_2003_17 : UINT;
    E005_Out_OUT23_2003_18 : UINT;
    E005_Out_OUT24_2003_19 : UINT;
    E005_Out_OUT25_2003_1A : UINT;
    E005_Out_OUT26_2003_1B : UINT;
    E005_Out_OUT27_2003_1C : UINT;
    E005_Out_OUT28_2003_1D : UINT;
    E005_Out_OUT29_2003_1E : UINT;
    E005_Out_OUT30_2003_1F : UINT;
    E005_Out_OUT31_2003_20 : UINT;
    E005_Out_OUT32_2003_21 : UINT;
    E005_Out_OUT33_2003_22 : UINT;
    E005_Out_OUT34_2003_23 : UINT;
    E005_Out_OUT35_2003_24 : UINT;
    E005_Out_OUT36_2003_25 : UINT;
    E005_Out_OUT37_2003_26 : UINT;
    E005_Out_OUT38_2003_27 : UINT;
    E005_Out_OUT39_2003_28 : UINT;
    E005_Out_OUT40_2003_29 : UINT;
    E005_Out_OUT41_2003_2A : UINT;
    E005_Out_OUT42_2003_2B : UINT;
    E005_Out_OUT43_2003_2C : UINT;
    E005_Out_OUT44_2003_2D : UINT;
    E005_Out_OUT45_2003_2E : UINT;
    E005_Out_OUT46_2003_2F : UINT;
    E005_Out_OUT47_2003_30 : UINT;
    E005_Out_OUT48_2003_31 : UINT;
    E005_Out_OUT49_2003_32 : UINT;
    E005_Out_OUT50_2003_33 : UINT;
    E005_Out_OUT51_2003_34 : UINT;
    E005_Out_OUT52_2003_35 : UINT;
    E005_Out_OUT53_2003_36 : UINT;
    E005_Out_OUT54_2003_37 : UINT;
    E005_Out_OUT55_2003_38 : UINT;
    E005_Out_OUT56_2003_39 : UINT;
    E005_Out_OUT57_2003_3A : UINT;
    E005_Out_OUT58_2003_3B : UINT;
    E005_Out_OUT59_2003_3C : UINT;
    E005_Out_OUT60_2003_3D : UINT;
    E005_Out_OUT61_2003_3E : UINT;
    E005_Out_OUT62_2003_3F : UINT;
    E005_Out_OUT63_2003_40 : UINT;
    E005_Out_OUT64_2003_41 : UINT;
    E005_Out_OUT65_2003_42 : UINT;
    E005_Out_OUT66_2003_43 : UINT;
    E005_Out_OUT67_2003_44 : UINT;
    E005_Out_OUT68_2003_45 : UINT;
    E005_Out_OUT69_2003_46 : UINT;
    E005_Out_OUT70_2003_47 : UINT;
    E005_Out_OUT71_2003_48 : UINT;
    E005_In_IN00_2004_01 : UINT;
    E005_In_IN01_2004_02 : UINT;
    E005_In_IN02_2004_03 : UINT;
    E005_In_IN03_2004_04 : UINT;
    E005_In_IN04_2004_05 : UINT;
    E005_In_IN05_2004_06 : UINT;
    E005_In_IN06_2004_07 : UINT;
    E005_In_IN07_2004_08 : UINT;
    E005_In_IN08_2004_09 : UINT;
    E005_In_IN09_2004_0A : UINT;
    E005_In_IN10_2004_0B : UINT;
    E005_In_IN11_2004_0C : UINT;
    E005_In_IN12_2004_0D : UINT;
    E005_In_IN13_2004_0E : UINT;
    E005_In_IN14_2004_0F : UINT;
    E005_In_IN15_2004_10 : UINT;
    E005_In_IN16_2004_11 : UINT;
    E005_In_IN17_2004_12 : UINT;
    E005_In_IN18_2004_13 : UINT;
    E005_In_IN19_2004_14 : UINT;
    E005_In_IN20_2004_15 : UINT;
    E005_In_IN21_2004_16 : UINT;
    E005_In_IN22_2004_17 : UINT;
    E005_In_IN23_2004_18 : UINT;
    E005_In_IN24_2004_19 : UINT;
    E005_In_IN25_2004_1A : UINT;
    E005_In_IN26_2004_1B : UINT;
    E005_In_IN27_2004_1C : UINT;
    E005_In_IN28_2004_1D : UINT;
    E005_In_IN29_2004_1E : UINT;
    E005_In_IN30_2004_1F : UINT;
    E005_In_IN31_2004_20 : UINT;
    E005_In_IN32_2004_21 : UINT;
    E005_In_IN33_2004_22 : UINT;
    E005_In_IN34_2004_23 : UINT;
    E005_In_IN35_2004_24 : UINT;
    E005_In_IN36_2004_25 : UINT;
    E005_In_IN37_2004_26 : UINT;
    E005_In_IN38_2004_27 : UINT;
    E005_In_IN39_2004_28 : UINT;
    E005_In_IN40_2004_29 : UINT;
    E005_In_IN41_2004_2A : UINT;
    E005_In_IN42_2004_2B : UINT;
    E005_In_IN43_2004_2C : UINT;
    E005_In_IN44_2004_2D : UINT;
    E005_In_IN45_2004_2E : UINT;
    E005_In_IN46_2004_2F : UINT;
    E005_In_IN47_2004_30 : UINT;
    E005_In_IN48_2004_31 : UINT;
    E005_In_IN49_2004_32 : UINT;
    E005_In_IN50_2004_33 : UINT;
    E005_In_IN51_2004_34 : UINT;
    E005_In_IN52_2004_35 : UINT;
    E005_In_IN53_2004_36 : UINT;
    E005_In_IN54_2004_37 : UINT;
    E005_In_IN55_2004_38 : UINT;
    E005_In_IN56_2004_39 : UINT;
    E005_In_IN57_2004_3A : UINT;
    E005_In_IN58_2004_3B : UINT;
    E005_In_IN59_2004_3C : UINT;
    E005_In_IN60_2004_3D : UINT;
    E005_In_IN61_2004_3E : UINT;
    E005_In_IN62_2004_3F : UINT;
    E005_In_IN63_2004_40 : UINT;
    E005_In_IN64_2004_41 : UINT;
    E005_In_IN65_2004_42 : UINT;
    E005_In_IN66_2004_43 : UINT;
    E005_In_IN67_2004_44 : UINT;
    E005_In_IN68_2004_45 : UINT;
    E005_In_IN69_2004_46 : UINT;
    E005_In_IN70_2004_47 : UINT;
    E005_In_IN71_2004_48 : UINT;
    E005_Out_OUT00_2003_01_1 : UINT;  (* RCON2（Node5） PLC→RCON 【OUT00】共通 ゲートウェイ制御信号0（MON等）; at ECAT://node#5/Out_OUT00_2003_01 *)
    E005_Out_OUT01_2003_02_1 : UINT;  (* RCON2（Node5） PLC→RCON 【OUT01】共通 ゲートウェイ制御信号1（予約・使用禁止）／今回書込まない; at ECAT://node#5/Out_OUT01_2003_02 *)
    E005_Out_OUT02_2003_03_1 : UINT;  (* RCON2（Node5） PLC→RCON 【OUT02】共通 共通予約領域（使用禁止・占有あり）／今回書込まない; at ECAT://node#5/Out_OUT02_2003_03 *)
    E005_Out_OUT03_2003_04_1 : UINT;  (* RCON2（Node5） PLC→RCON 【OUT03】共通 共通予約領域（使用禁止・占有あり）／今回書込まない; at ECAT://node#5/Out_OUT03_2003_04 *)
    E005_Out_OUT04_2003_05_1 : UINT;  (* RCON2（Node5） PLC→RCON 【OUT04】共通 共通予約領域（使用禁止・占有あり）／今回書込まない; at ECAT://node#5/Out_OUT04_2003_05 *)
    E005_Out_OUT05_2003_06_1 : UINT;  (* RCON2（Node5） PLC→RCON 【OUT05】共通 共通予約領域（使用禁止・占有あり）／今回書込まない; at ECAT://node#5/Out_OUT05_2003_06 *)
    E005_Out_OUT06_2003_07_1 : UINT;  (* RCON2（Node5） PLC→RCON 【OUT06】共通 共通予約領域（使用禁止・占有あり）／今回書込まない; at ECAT://node#5/Out_OUT06_2003_07 *)
    E005_Out_OUT07_2003_08_1 : UINT;  (* RCON2（Node5） PLC→RCON 【OUT07】共通 共通予約領域（使用禁止・占有あり）／今回書込まない; at ECAT://node#5/Out_OUT07_2003_08 *)
    E005_Out_OUT08_2003_09_1 : UINT;  (* RCON2（Node5） PLC→RCON 【OUT08】1軸目（No.0） 目標位置 下位ワード; at ECAT://node#5/Out_OUT08_2003_09 *)
    E005_Out_OUT09_2003_0A_1 : UINT;  (* RCON2（Node5） PLC→RCON 【OUT09】1軸目（No.0） 目標位置 上位ワード; at ECAT://node#5/Out_OUT09_2003_0A *)
    E005_Out_OUT10_2003_0B_1 : UINT;  (* RCON2（Node5） PLC→RCON 【OUT10】1軸目（No.0） 位置決め幅 下位ワード; at ECAT://node#5/Out_OUT10_2003_0B *)
    E005_Out_OUT11_2003_0C_1 : UINT;  (* RCON2（Node5） PLC→RCON 【OUT11】1軸目（No.0） 位置決め幅 上位ワード; at ECAT://node#5/Out_OUT11_2003_0C *)
    E005_Out_OUT12_2003_0D_1 : UINT;  (* RCON2（Node5） PLC→RCON 【OUT12】1軸目（No.0） 速度指令; at ECAT://node#5/Out_OUT12_2003_0D *)
    E005_Out_OUT13_2003_0E_1 : UINT;  (* RCON2（Node5） PLC→RCON 【OUT13】1軸目（No.0） 加減速度指令（加速・減速共通）; at ECAT://node#5/Out_OUT13_2003_0E *)
    E005_Out_OUT14_2003_0F_1 : UINT;  (* RCON2（Node5） PLC→RCON 【OUT14】1軸目（No.0） 押付け電流制限値; at ECAT://node#5/Out_OUT14_2003_0F *)
    E005_Out_OUT15_2003_10_1 : UINT;  (* RCON2（Node5） PLC→RCON 【OUT15】1軸目（No.0） 軸制御信号（DSTR・SON等）; at ECAT://node#5/Out_OUT15_2003_10 *)
    E005_Out_OUT16_2003_11_1 : UINT;  (* RCON2（Node5） PLC→RCON 【OUT16】2軸目（No.1） 目標位置 下位ワード; at ECAT://node#5/Out_OUT16_2003_11 *)
    E005_Out_OUT17_2003_12_1 : UINT;  (* RCON2（Node5） PLC→RCON 【OUT17】2軸目（No.1） 目標位置 上位ワード; at ECAT://node#5/Out_OUT17_2003_12 *)
    E005_Out_OUT18_2003_13_1 : UINT;  (* RCON2（Node5） PLC→RCON 【OUT18】2軸目（No.1） 位置決め幅 下位ワード; at ECAT://node#5/Out_OUT18_2003_13 *)
    E005_Out_OUT19_2003_14_1 : UINT;  (* RCON2（Node5） PLC→RCON 【OUT19】2軸目（No.1） 位置決め幅 上位ワード; at ECAT://node#5/Out_OUT19_2003_14 *)
    E005_Out_OUT20_2003_15_1 : UINT;  (* RCON2（Node5） PLC→RCON 【OUT20】2軸目（No.1） 速度指令; at ECAT://node#5/Out_OUT20_2003_15 *)
    E005_Out_OUT21_2003_16_1 : UINT;  (* RCON2（Node5） PLC→RCON 【OUT21】2軸目（No.1） 加減速度指令（加速・減速共通）; at ECAT://node#5/Out_OUT21_2003_16 *)
    E005_Out_OUT22_2003_17_1 : UINT;  (* RCON2（Node5） PLC→RCON 【OUT22】2軸目（No.1） 押付け電流制限値; at ECAT://node#5/Out_OUT22_2003_17 *)
    E005_Out_OUT23_2003_18_1 : UINT;  (* RCON2（Node5） PLC→RCON 【OUT23】2軸目（No.1） 軸制御信号（DSTR・SON等）; at ECAT://node#5/Out_OUT23_2003_18 *)
    E005_Out_OUT24_2003_19_1 : UINT;  (* RCON2（Node5） PLC→RCON 【OUT24】3軸目（No.2） 目標位置 下位ワード; at ECAT://node#5/Out_OUT24_2003_19 *)
    E005_Out_OUT25_2003_1A_1 : UINT;  (* RCON2（Node5） PLC→RCON 【OUT25】3軸目（No.2） 目標位置 上位ワード; at ECAT://node#5/Out_OUT25_2003_1A *)
    E005_Out_OUT26_2003_1B_1 : UINT;  (* RCON2（Node5） PLC→RCON 【OUT26】3軸目（No.2） 位置決め幅 下位ワード; at ECAT://node#5/Out_OUT26_2003_1B *)
    E005_Out_OUT27_2003_1C_1 : UINT;  (* RCON2（Node5） PLC→RCON 【OUT27】3軸目（No.2） 位置決め幅 上位ワード; at ECAT://node#5/Out_OUT27_2003_1C *)
    E005_Out_OUT28_2003_1D_1 : UINT;  (* RCON2（Node5） PLC→RCON 【OUT28】3軸目（No.2） 速度指令; at ECAT://node#5/Out_OUT28_2003_1D *)
    E005_Out_OUT29_2003_1E_1 : UINT;  (* RCON2（Node5） PLC→RCON 【OUT29】3軸目（No.2） 加減速度指令（加速・減速共通）; at ECAT://node#5/Out_OUT29_2003_1E *)
    E005_Out_OUT30_2003_1F_1 : UINT;  (* RCON2（Node5） PLC→RCON 【OUT30】3軸目（No.2） 押付け電流制限値; at ECAT://node#5/Out_OUT30_2003_1F *)
    E005_Out_OUT31_2003_20_1 : UINT;  (* RCON2（Node5） PLC→RCON 【OUT31】3軸目（No.2） 軸制御信号（DSTR・SON等）; at ECAT://node#5/Out_OUT31_2003_20 *)
    E005_Out_OUT32_2003_21_1 : UINT;  (* RCON2（Node5） PLC→RCON 【OUT32】4軸目（No.3） 目標位置 下位ワード; at ECAT://node#5/Out_OUT32_2003_21 *)
    E005_Out_OUT33_2003_22_1 : UINT;  (* RCON2（Node5） PLC→RCON 【OUT33】4軸目（No.3） 目標位置 上位ワード; at ECAT://node#5/Out_OUT33_2003_22 *)
    E005_Out_OUT34_2003_23_1 : UINT;  (* RCON2（Node5） PLC→RCON 【OUT34】4軸目（No.3） 位置決め幅 下位ワード; at ECAT://node#5/Out_OUT34_2003_23 *)
    E005_Out_OUT35_2003_24_1 : UINT;  (* RCON2（Node5） PLC→RCON 【OUT35】4軸目（No.3） 位置決め幅 上位ワード; at ECAT://node#5/Out_OUT35_2003_24 *)
    E005_Out_OUT36_2003_25_1 : UINT;  (* RCON2（Node5） PLC→RCON 【OUT36】4軸目（No.3） 速度指令; at ECAT://node#5/Out_OUT36_2003_25 *)
    E005_Out_OUT37_2003_26_1 : UINT;  (* RCON2（Node5） PLC→RCON 【OUT37】4軸目（No.3） 加減速度指令（加速・減速共通）; at ECAT://node#5/Out_OUT37_2003_26 *)
    E005_Out_OUT38_2003_27_1 : UINT;  (* RCON2（Node5） PLC→RCON 【OUT38】4軸目（No.3） 押付け電流制限値; at ECAT://node#5/Out_OUT38_2003_27 *)
    E005_Out_OUT39_2003_28_1 : UINT;  (* RCON2（Node5） PLC→RCON 【OUT39】4軸目（No.3） 軸制御信号（DSTR・SON等）; at ECAT://node#5/Out_OUT39_2003_28 *)
    E005_Out_OUT40_2003_29_1 : UINT;  (* RCON2（Node5） PLC→RCON 【OUT40】5軸目（No.4） 目標位置 下位ワード; at ECAT://node#5/Out_OUT40_2003_29 *)
    E005_Out_OUT41_2003_2A_1 : UINT;  (* RCON2（Node5） PLC→RCON 【OUT41】5軸目（No.4） 目標位置 上位ワード; at ECAT://node#5/Out_OUT41_2003_2A *)
    E005_Out_OUT42_2003_2B_1 : UINT;  (* RCON2（Node5） PLC→RCON 【OUT42】5軸目（No.4） 位置決め幅 下位ワード; at ECAT://node#5/Out_OUT42_2003_2B *)
    E005_Out_OUT43_2003_2C_1 : UINT;  (* RCON2（Node5） PLC→RCON 【OUT43】5軸目（No.4） 位置決め幅 上位ワード; at ECAT://node#5/Out_OUT43_2003_2C *)
    E005_Out_OUT44_2003_2D_1 : UINT;  (* RCON2（Node5） PLC→RCON 【OUT44】5軸目（No.4） 速度指令; at ECAT://node#5/Out_OUT44_2003_2D *)
    E005_Out_OUT45_2003_2E_1 : UINT;  (* RCON2（Node5） PLC→RCON 【OUT45】5軸目（No.4） 加減速度指令（加速・減速共通）; at ECAT://node#5/Out_OUT45_2003_2E *)
    E005_Out_OUT46_2003_2F_1 : UINT;  (* RCON2（Node5） PLC→RCON 【OUT46】5軸目（No.4） 押付け電流制限値; at ECAT://node#5/Out_OUT46_2003_2F *)
    E005_Out_OUT47_2003_30_1 : UINT;  (* RCON2（Node5） PLC→RCON 【OUT47】5軸目（No.4） 軸制御信号（DSTR・SON等）; at ECAT://node#5/Out_OUT47_2003_30 *)
    E005_Out_OUT48_2003_31_1 : UINT;  (* RCON2（Node5） 【OUT48】用途未確認領域。今回の軸データ変換では未使用。／今回書込まない; at ECAT://node#5/Out_OUT48_2003_31 *)
    E005_Out_OUT49_2003_32_1 : UINT;  (* RCON2（Node5） 【OUT49】用途未確認領域。今回の軸データ変換では未使用。／今回書込まない; at ECAT://node#5/Out_OUT49_2003_32 *)
    E005_Out_OUT50_2003_33_1 : UINT;  (* RCON2（Node5） 【OUT50】用途未確認領域。今回の軸データ変換では未使用。／今回書込まない; at ECAT://node#5/Out_OUT50_2003_33 *)
    E005_Out_OUT51_2003_34_1 : UINT;  (* RCON2（Node5） 【OUT51】用途未確認領域。今回の軸データ変換では未使用。／今回書込まない; at ECAT://node#5/Out_OUT51_2003_34 *)
    E005_Out_OUT52_2003_35_1 : UINT;  (* RCON2（Node5） 【OUT52】用途未確認領域。今回の軸データ変換では未使用。／今回書込まない; at ECAT://node#5/Out_OUT52_2003_35 *)
    E005_Out_OUT53_2003_36_1 : UINT;  (* RCON2（Node5） 【OUT53】用途未確認領域。今回の軸データ変換では未使用。／今回書込まない; at ECAT://node#5/Out_OUT53_2003_36 *)
    E005_Out_OUT54_2003_37_1 : UINT;  (* RCON2（Node5） 【OUT54】用途未確認領域。今回の軸データ変換では未使用。／今回書込まない; at ECAT://node#5/Out_OUT54_2003_37 *)
    E005_Out_OUT55_2003_38_1 : UINT;  (* RCON2（Node5） 【OUT55】用途未確認領域。今回の軸データ変換では未使用。／今回書込まない; at ECAT://node#5/Out_OUT55_2003_38 *)
    E005_In_IN00_2004_01_1 : UINT;  (* RCON2（Node5） RCON→PLC 【IN00】共通 ゲートウェイ状態信号0; at ECAT://node#5/In_IN00_2004_01 *)
    E005_In_IN01_2004_02_1 : UINT;  (* RCON2（Node5） RCON→PLC 【IN01】共通 ゲートウェイ状態信号1（軸No.0～15リンク状態）; at ECAT://node#5/In_IN01_2004_02 *)
    E005_In_IN02_2004_03_1 : UINT;  (* RCON2（Node5） RCON→PLC 【IN02】共通 電源ユニット状態信号0; at ECAT://node#5/In_IN02_2004_03 *)
    E005_In_IN03_2004_04_1 : UINT;  (* RCON2（Node5） RCON→PLC 【IN03】共通 電源ユニット状態信号1; at ECAT://node#5/In_IN03_2004_04 *)
    E005_In_IN04_2004_05_1 : UINT;  (* RCON2（Node5） RCON→PLC 【IN04】共通 電源ユニット状態信号2; at ECAT://node#5/In_IN04_2004_05 *)
    E005_In_IN05_2004_06_1 : UINT;  (* RCON2（Node5） RCON→PLC 【IN05】共通 電源ユニット状態信号3; at ECAT://node#5/In_IN05_2004_06 *)
    E005_In_IN06_2004_07_1 : UINT;  (* RCON2（Node5） RCON→PLC 【IN06】共通 電源ユニット状態信号4／軽故障メンテナンス（設定依存）; at ECAT://node#5/In_IN06_2004_07 *)
    E005_In_IN07_2004_08_1 : UINT;  (* RCON2（Node5） RCON→PLC 【IN07】共通 共通予約領域（使用禁止・占有あり）; at ECAT://node#5/In_IN07_2004_08 *)
    E005_In_IN08_2004_09_1 : UINT;  (* RCON2（Node5） RCON→PLC 【IN08】1軸目（No.0） 現在位置 下位ワード; at ECAT://node#5/In_IN08_2004_09 *)
    E005_In_IN09_2004_0A_1 : UINT;  (* RCON2（Node5） RCON→PLC 【IN09】1軸目（No.0） 現在位置 上位ワード; at ECAT://node#5/In_IN09_2004_0A *)
    E005_In_IN10_2004_0B_1 : UINT;  (* RCON2（Node5） RCON→PLC 【IN10】1軸目（No.0） 現在電流 下位ワード（PCは指令電流）; at ECAT://node#5/In_IN10_2004_0B *)
    E005_In_IN11_2004_0C_1 : UINT;  (* RCON2（Node5） RCON→PLC 【IN11】1軸目（No.0） 現在電流 上位ワード（PCは指令電流）; at ECAT://node#5/In_IN11_2004_0C *)
    E005_In_IN12_2004_0D_1 : UINT;  (* RCON2（Node5） RCON→PLC 【IN12】1軸目（No.0） 現在速度（負方向は2の補数）; at ECAT://node#5/In_IN12_2004_0D *)
    E005_In_IN13_2004_0E_1 : UINT;  (* RCON2（Node5） RCON→PLC 【IN13】1軸目（No.0） 予約領域（使用禁止）; at ECAT://node#5/In_IN13_2004_0E *)
    E005_In_IN14_2004_0F_1 : UINT;  (* RCON2（Node5） RCON→PLC 【IN14】1軸目（No.0） アラームコード（簡易コードではない）; at ECAT://node#5/In_IN14_2004_0F *)
    E005_In_IN15_2004_10_1 : UINT;  (* RCON2（Node5） RCON→PLC 【IN15】1軸目（No.0） 軸状態信号（PEND・SV等）; at ECAT://node#5/In_IN15_2004_10 *)
    E005_In_IN16_2004_11_1 : UINT;  (* RCON2（Node5） RCON→PLC 【IN16】2軸目（No.1） 現在位置 下位ワード; at ECAT://node#5/In_IN16_2004_11 *)
    E005_In_IN17_2004_12_1 : UINT;  (* RCON2（Node5） RCON→PLC 【IN17】2軸目（No.1） 現在位置 上位ワード; at ECAT://node#5/In_IN17_2004_12 *)
    E005_In_IN18_2004_13_1 : UINT;  (* RCON2（Node5） RCON→PLC 【IN18】2軸目（No.1） 現在電流 下位ワード（PCは指令電流）; at ECAT://node#5/In_IN18_2004_13 *)
    E005_In_IN19_2004_14_1 : UINT;  (* RCON2（Node5） RCON→PLC 【IN19】2軸目（No.1） 現在電流 上位ワード（PCは指令電流）; at ECAT://node#5/In_IN19_2004_14 *)
    E005_In_IN20_2004_15_1 : UINT;  (* RCON2（Node5） RCON→PLC 【IN20】2軸目（No.1） 現在速度（負方向は2の補数）; at ECAT://node#5/In_IN20_2004_15 *)
    E005_In_IN21_2004_16_1 : UINT;  (* RCON2（Node5） RCON→PLC 【IN21】2軸目（No.1） 予約領域（使用禁止）; at ECAT://node#5/In_IN21_2004_16 *)
    E005_In_IN22_2004_17_1 : UINT;  (* RCON2（Node5） RCON→PLC 【IN22】2軸目（No.1） アラームコード（簡易コードではない）; at ECAT://node#5/In_IN22_2004_17 *)
    E005_In_IN23_2004_18_1 : UINT;  (* RCON2（Node5） RCON→PLC 【IN23】2軸目（No.1） 軸状態信号（PEND・SV等）; at ECAT://node#5/In_IN23_2004_18 *)
    E005_In_IN24_2004_19_1 : UINT;  (* RCON2（Node5） RCON→PLC 【IN24】3軸目（No.2） 現在位置 下位ワード; at ECAT://node#5/In_IN24_2004_19 *)
    E005_In_IN25_2004_1A_1 : UINT;  (* RCON2（Node5） RCON→PLC 【IN25】3軸目（No.2） 現在位置 上位ワード; at ECAT://node#5/In_IN25_2004_1A *)
    E005_In_IN26_2004_1B_1 : UINT;  (* RCON2（Node5） RCON→PLC 【IN26】3軸目（No.2） 現在電流 下位ワード（PCは指令電流）; at ECAT://node#5/In_IN26_2004_1B *)
    E005_In_IN27_2004_1C_1 : UINT;  (* RCON2（Node5） RCON→PLC 【IN27】3軸目（No.2） 現在電流 上位ワード（PCは指令電流）; at ECAT://node#5/In_IN27_2004_1C *)
    E005_In_IN28_2004_1D_1 : UINT;  (* RCON2（Node5） RCON→PLC 【IN28】3軸目（No.2） 現在速度（負方向は2の補数）; at ECAT://node#5/In_IN28_2004_1D *)
    E005_In_IN29_2004_1E_1 : UINT;  (* RCON2（Node5） RCON→PLC 【IN29】3軸目（No.2） 予約領域（使用禁止）; at ECAT://node#5/In_IN29_2004_1E *)
    E005_In_IN30_2004_1F_1 : UINT;  (* RCON2（Node5） RCON→PLC 【IN30】3軸目（No.2） アラームコード（簡易コードではない）; at ECAT://node#5/In_IN30_2004_1F *)
    E005_In_IN31_2004_20_1 : UINT;  (* RCON2（Node5） RCON→PLC 【IN31】3軸目（No.2） 軸状態信号（PEND・SV等）; at ECAT://node#5/In_IN31_2004_20 *)
    E005_In_IN32_2004_21_1 : UINT;  (* RCON2（Node5） RCON→PLC 【IN32】4軸目（No.3） 現在位置 下位ワード; at ECAT://node#5/In_IN32_2004_21 *)
    E005_In_IN33_2004_22_1 : UINT;  (* RCON2（Node5） RCON→PLC 【IN33】4軸目（No.3） 現在位置 上位ワード; at ECAT://node#5/In_IN33_2004_22 *)
    E005_In_IN34_2004_23_1 : UINT;  (* RCON2（Node5） RCON→PLC 【IN34】4軸目（No.3） 現在電流 下位ワード（PCは指令電流）; at ECAT://node#5/In_IN34_2004_23 *)
    E005_In_IN35_2004_24_1 : UINT;  (* RCON2（Node5） RCON→PLC 【IN35】4軸目（No.3） 現在電流 上位ワード（PCは指令電流）; at ECAT://node#5/In_IN35_2004_24 *)
    E005_In_IN36_2004_25_1 : UINT;  (* RCON2（Node5） RCON→PLC 【IN36】4軸目（No.3） 現在速度（負方向は2の補数）; at ECAT://node#5/In_IN36_2004_25 *)
    E005_In_IN37_2004_26_1 : UINT;  (* RCON2（Node5） RCON→PLC 【IN37】4軸目（No.3） 予約領域（使用禁止）; at ECAT://node#5/In_IN37_2004_26 *)
    E005_In_IN38_2004_27_1 : UINT;  (* RCON2（Node5） RCON→PLC 【IN38】4軸目（No.3） アラームコード（簡易コードではない）; at ECAT://node#5/In_IN38_2004_27 *)
    E005_In_IN39_2004_28_1 : UINT;  (* RCON2（Node5） RCON→PLC 【IN39】4軸目（No.3） 軸状態信号（PEND・SV等）; at ECAT://node#5/In_IN39_2004_28 *)
    E005_In_IN40_2004_29_1 : UINT;  (* RCON2（Node5） RCON→PLC 【IN40】5軸目（No.4） 現在位置 下位ワード; at ECAT://node#5/In_IN40_2004_29 *)
    E005_In_IN41_2004_2A_1 : UINT;  (* RCON2（Node5） RCON→PLC 【IN41】5軸目（No.4） 現在位置 上位ワード; at ECAT://node#5/In_IN41_2004_2A *)
    E005_In_IN42_2004_2B_1 : UINT;  (* RCON2（Node5） RCON→PLC 【IN42】5軸目（No.4） 現在電流 下位ワード（PCは指令電流）; at ECAT://node#5/In_IN42_2004_2B *)
    E005_In_IN43_2004_2C_1 : UINT;  (* RCON2（Node5） RCON→PLC 【IN43】5軸目（No.4） 現在電流 上位ワード（PCは指令電流）; at ECAT://node#5/In_IN43_2004_2C *)
    E005_In_IN44_2004_2D_1 : UINT;  (* RCON2（Node5） RCON→PLC 【IN44】5軸目（No.4） 現在速度（負方向は2の補数）; at ECAT://node#5/In_IN44_2004_2D *)
    E005_In_IN45_2004_2E_1 : UINT;  (* RCON2（Node5） RCON→PLC 【IN45】5軸目（No.4） 予約領域（使用禁止）; at ECAT://node#5/In_IN45_2004_2E *)
    E005_In_IN46_2004_2F_1 : UINT;  (* RCON2（Node5） RCON→PLC 【IN46】5軸目（No.4） アラームコード（簡易コードではない）; at ECAT://node#5/In_IN46_2004_2F *)
    E005_In_IN47_2004_30_1 : UINT;  (* RCON2（Node5） RCON→PLC 【IN47】5軸目（No.4） 軸状態信号（PEND・SV等）; at ECAT://node#5/In_IN47_2004_30 *)
    E005_In_IN48_2004_31_1 : UINT;  (* RCON2（Node5） 【IN48】用途未確認領域。今回の軸データ変換では未使用。; at ECAT://node#5/In_IN48_2004_31 *)
    E005_In_IN49_2004_32_1 : UINT;  (* RCON2（Node5） 【IN49】用途未確認領域。今回の軸データ変換では未使用。; at ECAT://node#5/In_IN49_2004_32 *)
    E005_In_IN50_2004_33_1 : UINT;  (* RCON2（Node5） 【IN50】用途未確認領域。今回の軸データ変換では未使用。; at ECAT://node#5/In_IN50_2004_33 *)
    E005_In_IN51_2004_34_1 : UINT;  (* RCON2（Node5） 【IN51】用途未確認領域。今回の軸データ変換では未使用。; at ECAT://node#5/In_IN51_2004_34 *)
    E005_In_IN52_2004_35_1 : UINT;  (* RCON2（Node5） 【IN52】用途未確認領域。今回の軸データ変換では未使用。; at ECAT://node#5/In_IN52_2004_35 *)
    E005_In_IN53_2004_36_1 : UINT;  (* RCON2（Node5） 【IN53】用途未確認領域。今回の軸データ変換では未使用。; at ECAT://node#5/In_IN53_2004_36 *)
    E005_In_IN54_2004_37_1 : UINT;  (* RCON2（Node5） 【IN54】用途未確認領域。今回の軸データ変換では未使用。; at ECAT://node#5/In_IN54_2004_37 *)
    E005_In_IN55_2004_38_1 : UINT;  (* RCON2（Node5） 【IN55】用途未確認領域。今回の軸データ変換では未使用。; at ECAT://node#5/In_IN55_2004_38 *)
    E001_Out_OUT00_2003_01 : UINT;  (* RCON1（Node1） PLC→RCON 【OUT00】共通 ゲートウェイ制御信号0（MON等）; at ECAT://node#1/Out_OUT00_2003_01 *)
    E001_Out_OUT01_2003_02 : UINT;  (* RCON1（Node1） PLC→RCON 【OUT01】共通 ゲートウェイ制御信号1（予約・使用禁止）／今回書込まない; at ECAT://node#1/Out_OUT01_2003_02 *)
    E001_Out_OUT02_2003_03 : UINT;  (* RCON1（Node1） PLC→RCON 【OUT02】共通 共通予約領域（使用禁止・占有あり）／今回書込まない; at ECAT://node#1/Out_OUT02_2003_03 *)
    E001_Out_OUT03_2003_04 : UINT;  (* RCON1（Node1） PLC→RCON 【OUT03】共通 共通予約領域（使用禁止・占有あり）／今回書込まない; at ECAT://node#1/Out_OUT03_2003_04 *)
    E001_Out_OUT04_2003_05 : UINT;  (* RCON1（Node1） PLC→RCON 【OUT04】共通 共通予約領域（使用禁止・占有あり）／今回書込まない; at ECAT://node#1/Out_OUT04_2003_05 *)
    E001_Out_OUT05_2003_06 : UINT;  (* RCON1（Node1） PLC→RCON 【OUT05】共通 共通予約領域（使用禁止・占有あり）／今回書込まない; at ECAT://node#1/Out_OUT05_2003_06 *)
    E001_Out_OUT06_2003_07 : UINT;  (* RCON1（Node1） PLC→RCON 【OUT06】共通 共通予約領域（使用禁止・占有あり）／今回書込まない; at ECAT://node#1/Out_OUT06_2003_07 *)
    E001_Out_OUT07_2003_08 : UINT;  (* RCON1（Node1） PLC→RCON 【OUT07】共通 共通予約領域（使用禁止・占有あり）／今回書込まない; at ECAT://node#1/Out_OUT07_2003_08 *)
    E001_Out_OUT08_2003_09 : UINT;  (* RCON1（Node1） PLC→RCON 【OUT08】1軸目（No.0） 目標位置 下位ワード; at ECAT://node#1/Out_OUT08_2003_09 *)
    E001_Out_OUT09_2003_0A : UINT;  (* RCON1（Node1） PLC→RCON 【OUT09】1軸目（No.0） 目標位置 上位ワード; at ECAT://node#1/Out_OUT09_2003_0A *)
    E001_Out_OUT10_2003_0B : UINT;  (* RCON1（Node1） PLC→RCON 【OUT10】1軸目（No.0） 位置決め幅 下位ワード; at ECAT://node#1/Out_OUT10_2003_0B *)
    E001_Out_OUT11_2003_0C : UINT;  (* RCON1（Node1） PLC→RCON 【OUT11】1軸目（No.0） 位置決め幅 上位ワード; at ECAT://node#1/Out_OUT11_2003_0C *)
    E001_Out_OUT12_2003_0D : UINT;  (* RCON1（Node1） PLC→RCON 【OUT12】1軸目（No.0） 速度指令; at ECAT://node#1/Out_OUT12_2003_0D *)
    E001_Out_OUT13_2003_0E : UINT;  (* RCON1（Node1） PLC→RCON 【OUT13】1軸目（No.0） 加減速度指令（加速・減速共通）; at ECAT://node#1/Out_OUT13_2003_0E *)
    E001_Out_OUT14_2003_0F : UINT;  (* RCON1（Node1） PLC→RCON 【OUT14】1軸目（No.0） 押付け電流制限値; at ECAT://node#1/Out_OUT14_2003_0F *)
    E001_Out_OUT15_2003_10 : UINT;  (* RCON1（Node1） PLC→RCON 【OUT15】1軸目（No.0） 軸制御信号（DSTR・SON等）; at ECAT://node#1/Out_OUT15_2003_10 *)
    E001_Out_OUT16_2003_11 : UINT;  (* RCON1（Node1） PLC→RCON 【OUT16】2軸目（No.1） 目標位置 下位ワード; at ECAT://node#1/Out_OUT16_2003_11 *)
    E001_Out_OUT17_2003_12 : UINT;  (* RCON1（Node1） PLC→RCON 【OUT17】2軸目（No.1） 目標位置 上位ワード; at ECAT://node#1/Out_OUT17_2003_12 *)
    E001_Out_OUT18_2003_13 : UINT;  (* RCON1（Node1） PLC→RCON 【OUT18】2軸目（No.1） 位置決め幅 下位ワード; at ECAT://node#1/Out_OUT18_2003_13 *)
    E001_Out_OUT19_2003_14 : UINT;  (* RCON1（Node1） PLC→RCON 【OUT19】2軸目（No.1） 位置決め幅 上位ワード; at ECAT://node#1/Out_OUT19_2003_14 *)
    E001_Out_OUT20_2003_15 : UINT;  (* RCON1（Node1） PLC→RCON 【OUT20】2軸目（No.1） 速度指令; at ECAT://node#1/Out_OUT20_2003_15 *)
    E001_Out_OUT21_2003_16 : UINT;  (* RCON1（Node1） PLC→RCON 【OUT21】2軸目（No.1） 加減速度指令（加速・減速共通）; at ECAT://node#1/Out_OUT21_2003_16 *)
    E001_Out_OUT22_2003_17 : UINT;  (* RCON1（Node1） PLC→RCON 【OUT22】2軸目（No.1） 押付け電流制限値; at ECAT://node#1/Out_OUT22_2003_17 *)
    E001_Out_OUT23_2003_18 : UINT;  (* RCON1（Node1） PLC→RCON 【OUT23】2軸目（No.1） 軸制御信号（DSTR・SON等）; at ECAT://node#1/Out_OUT23_2003_18 *)
    E001_Out_OUT24_2003_19 : UINT;  (* RCON1（Node1） PLC→RCON 【OUT24】3軸目（No.2） 目標位置 下位ワード; at ECAT://node#1/Out_OUT24_2003_19 *)
    E001_Out_OUT25_2003_1A : UINT;  (* RCON1（Node1） PLC→RCON 【OUT25】3軸目（No.2） 目標位置 上位ワード; at ECAT://node#1/Out_OUT25_2003_1A *)
    E001_Out_OUT26_2003_1B : UINT;  (* RCON1（Node1） PLC→RCON 【OUT26】3軸目（No.2） 位置決め幅 下位ワード; at ECAT://node#1/Out_OUT26_2003_1B *)
    E001_Out_OUT27_2003_1C : UINT;  (* RCON1（Node1） PLC→RCON 【OUT27】3軸目（No.2） 位置決め幅 上位ワード; at ECAT://node#1/Out_OUT27_2003_1C *)
    E001_Out_OUT28_2003_1D : UINT;  (* RCON1（Node1） PLC→RCON 【OUT28】3軸目（No.2） 速度指令; at ECAT://node#1/Out_OUT28_2003_1D *)
    E001_Out_OUT29_2003_1E : UINT;  (* RCON1（Node1） PLC→RCON 【OUT29】3軸目（No.2） 加減速度指令（加速・減速共通）; at ECAT://node#1/Out_OUT29_2003_1E *)
    E001_Out_OUT30_2003_1F : UINT;  (* RCON1（Node1） PLC→RCON 【OUT30】3軸目（No.2） 押付け電流制限値; at ECAT://node#1/Out_OUT30_2003_1F *)
    E001_Out_OUT31_2003_20 : UINT;  (* RCON1（Node1） PLC→RCON 【OUT31】3軸目（No.2） 軸制御信号（DSTR・SON等）; at ECAT://node#1/Out_OUT31_2003_20 *)
    E001_Out_OUT32_2003_21 : UINT;  (* RCON1（Node1） PLC→RCON 【OUT32】4軸目（No.3） 目標位置 下位ワード; at ECAT://node#1/Out_OUT32_2003_21 *)
    E001_Out_OUT33_2003_22 : UINT;  (* RCON1（Node1） PLC→RCON 【OUT33】4軸目（No.3） 目標位置 上位ワード; at ECAT://node#1/Out_OUT33_2003_22 *)
    E001_Out_OUT34_2003_23 : UINT;  (* RCON1（Node1） PLC→RCON 【OUT34】4軸目（No.3） 位置決め幅 下位ワード; at ECAT://node#1/Out_OUT34_2003_23 *)
    E001_Out_OUT35_2003_24 : UINT;  (* RCON1（Node1） PLC→RCON 【OUT35】4軸目（No.3） 位置決め幅 上位ワード; at ECAT://node#1/Out_OUT35_2003_24 *)
    E001_Out_OUT36_2003_25 : UINT;  (* RCON1（Node1） PLC→RCON 【OUT36】4軸目（No.3） 速度指令; at ECAT://node#1/Out_OUT36_2003_25 *)
    E001_Out_OUT37_2003_26 : UINT;  (* RCON1（Node1） PLC→RCON 【OUT37】4軸目（No.3） 加減速度指令（加速・減速共通）; at ECAT://node#1/Out_OUT37_2003_26 *)
    E001_Out_OUT38_2003_27 : UINT;  (* RCON1（Node1） PLC→RCON 【OUT38】4軸目（No.3） 押付け電流制限値; at ECAT://node#1/Out_OUT38_2003_27 *)
    E001_Out_OUT39_2003_28 : UINT;  (* RCON1（Node1） PLC→RCON 【OUT39】4軸目（No.3） 軸制御信号（DSTR・SON等）; at ECAT://node#1/Out_OUT39_2003_28 *)
    E001_Out_OUT40_2003_29 : UINT;  (* RCON1（Node1） PLC→RCON 【OUT40】5軸目（No.4） 目標位置 下位ワード; at ECAT://node#1/Out_OUT40_2003_29 *)
    E001_Out_OUT41_2003_2A : UINT;  (* RCON1（Node1） PLC→RCON 【OUT41】5軸目（No.4） 目標位置 上位ワード; at ECAT://node#1/Out_OUT41_2003_2A *)
    E001_Out_OUT42_2003_2B : UINT;  (* RCON1（Node1） PLC→RCON 【OUT42】5軸目（No.4） 位置決め幅 下位ワード; at ECAT://node#1/Out_OUT42_2003_2B *)
    E001_Out_OUT43_2003_2C : UINT;  (* RCON1（Node1） PLC→RCON 【OUT43】5軸目（No.4） 位置決め幅 上位ワード; at ECAT://node#1/Out_OUT43_2003_2C *)
    E001_Out_OUT44_2003_2D : UINT;  (* RCON1（Node1） PLC→RCON 【OUT44】5軸目（No.4） 速度指令; at ECAT://node#1/Out_OUT44_2003_2D *)
    E001_Out_OUT45_2003_2E : UINT;  (* RCON1（Node1） PLC→RCON 【OUT45】5軸目（No.4） 加減速度指令（加速・減速共通）; at ECAT://node#1/Out_OUT45_2003_2E *)
    E001_Out_OUT46_2003_2F : UINT;  (* RCON1（Node1） PLC→RCON 【OUT46】5軸目（No.4） 押付け電流制限値; at ECAT://node#1/Out_OUT46_2003_2F *)
    E001_Out_OUT47_2003_30 : UINT;  (* RCON1（Node1） PLC→RCON 【OUT47】5軸目（No.4） 軸制御信号（DSTR・SON等）; at ECAT://node#1/Out_OUT47_2003_30 *)
    E001_Out_OUT48_2003_31 : UINT;  (* RCON1（Node1） PLC→RCON 【OUT48】6軸目（No.5） 目標位置 下位ワード; at ECAT://node#1/Out_OUT48_2003_31 *)
    E001_Out_OUT49_2003_32 : UINT;  (* RCON1（Node1） PLC→RCON 【OUT49】6軸目（No.5） 目標位置 上位ワード; at ECAT://node#1/Out_OUT49_2003_32 *)
    E001_Out_OUT50_2003_33 : UINT;  (* RCON1（Node1） PLC→RCON 【OUT50】6軸目（No.5） 位置決め幅 下位ワード; at ECAT://node#1/Out_OUT50_2003_33 *)
    E001_Out_OUT51_2003_34 : UINT;  (* RCON1（Node1） PLC→RCON 【OUT51】6軸目（No.5） 位置決め幅 上位ワード; at ECAT://node#1/Out_OUT51_2003_34 *)
    E001_Out_OUT52_2003_35 : UINT;  (* RCON1（Node1） PLC→RCON 【OUT52】6軸目（No.5） 速度指令; at ECAT://node#1/Out_OUT52_2003_35 *)
    E001_Out_OUT53_2003_36 : UINT;  (* RCON1（Node1） PLC→RCON 【OUT53】6軸目（No.5） 加減速度指令（加速・減速共通）; at ECAT://node#1/Out_OUT53_2003_36 *)
    E001_Out_OUT54_2003_37 : UINT;  (* RCON1（Node1） PLC→RCON 【OUT54】6軸目（No.5） 押付け電流制限値; at ECAT://node#1/Out_OUT54_2003_37 *)
    E001_Out_OUT55_2003_38 : UINT;  (* RCON1（Node1） PLC→RCON 【OUT55】6軸目（No.5） 軸制御信号（DSTR・SON等）; at ECAT://node#1/Out_OUT55_2003_38 *)
    E001_Out_OUT56_2003_39 : UINT;  (* RCON1（Node1） 【OUT56】用途未確認領域。今回の軸データ変換では未使用。／今回書込まない; at ECAT://node#1/Out_OUT56_2003_39 *)
    E001_Out_OUT57_2003_3A : UINT;  (* RCON1（Node1） 【OUT57】用途未確認領域。今回の軸データ変換では未使用。／今回書込まない; at ECAT://node#1/Out_OUT57_2003_3A *)
    E001_Out_OUT58_2003_3B : UINT;  (* RCON1（Node1） 【OUT58】用途未確認領域。今回の軸データ変換では未使用。／今回書込まない; at ECAT://node#1/Out_OUT58_2003_3B *)
    E001_Out_OUT59_2003_3C : UINT;  (* RCON1（Node1） 【OUT59】用途未確認領域。今回の軸データ変換では未使用。／今回書込まない; at ECAT://node#1/Out_OUT59_2003_3C *)
    E001_Out_OUT60_2003_3D : UINT;  (* RCON1（Node1） 【OUT60】用途未確認領域。今回の軸データ変換では未使用。／今回書込まない; at ECAT://node#1/Out_OUT60_2003_3D *)
    E001_Out_OUT61_2003_3E : UINT;  (* RCON1（Node1） 【OUT61】用途未確認領域。今回の軸データ変換では未使用。／今回書込まない; at ECAT://node#1/Out_OUT61_2003_3E *)
    E001_Out_OUT62_2003_3F : UINT;  (* RCON1（Node1） 【OUT62】用途未確認領域。今回の軸データ変換では未使用。／今回書込まない; at ECAT://node#1/Out_OUT62_2003_3F *)
    E001_Out_OUT63_2003_40 : UINT;  (* RCON1（Node1） 【OUT63】用途未確認領域。今回の軸データ変換では未使用。／今回書込まない; at ECAT://node#1/Out_OUT63_2003_40 *)
    E001_Out_OUT64_2003_41 : UINT;  (* RCON1（Node1） 【OUT64】用途未確認領域。今回の軸データ変換では未使用。／今回書込まない; at ECAT://node#1/Out_OUT64_2003_41 *)
    E001_Out_OUT65_2003_42 : UINT;  (* RCON1（Node1） 【OUT65】用途未確認領域。今回の軸データ変換では未使用。／今回書込まない; at ECAT://node#1/Out_OUT65_2003_42 *)
    E001_Out_OUT66_2003_43 : UINT;  (* RCON1（Node1） 【OUT66】用途未確認領域。今回の軸データ変換では未使用。／今回書込まない; at ECAT://node#1/Out_OUT66_2003_43 *)
    E001_Out_OUT67_2003_44 : UINT;  (* RCON1（Node1） 【OUT67】用途未確認領域。今回の軸データ変換では未使用。／今回書込まない; at ECAT://node#1/Out_OUT67_2003_44 *)
    E001_Out_OUT68_2003_45 : UINT;  (* RCON1（Node1） 【OUT68】用途未確認領域。今回の軸データ変換では未使用。／今回書込まない; at ECAT://node#1/Out_OUT68_2003_45 *)
    E001_Out_OUT69_2003_46 : UINT;  (* RCON1（Node1） 【OUT69】用途未確認領域。今回の軸データ変換では未使用。／今回書込まない; at ECAT://node#1/Out_OUT69_2003_46 *)
    E001_Out_OUT70_2003_47 : UINT;  (* RCON1（Node1） 【OUT70】用途未確認領域。今回の軸データ変換では未使用。／今回書込まない; at ECAT://node#1/Out_OUT70_2003_47 *)
    E001_Out_OUT71_2003_48 : UINT;  (* RCON1（Node1） 【OUT71】用途未確認領域。今回の軸データ変換では未使用。／今回書込まない; at ECAT://node#1/Out_OUT71_2003_48 *)
    E001_In_IN00_2004_01 : UINT;  (* RCON1（Node1） RCON→PLC 【IN00】共通 ゲートウェイ状態信号0; at ECAT://node#1/In_IN00_2004_01 *)
    E001_In_IN01_2004_02 : UINT;  (* RCON1（Node1） RCON→PLC 【IN01】共通 ゲートウェイ状態信号1（軸No.0～15リンク状態）; at ECAT://node#1/In_IN01_2004_02 *)
    E001_In_IN02_2004_03 : UINT;  (* RCON1（Node1） RCON→PLC 【IN02】共通 電源ユニット状態信号0; at ECAT://node#1/In_IN02_2004_03 *)
    E001_In_IN03_2004_04 : UINT;  (* RCON1（Node1） RCON→PLC 【IN03】共通 電源ユニット状態信号1; at ECAT://node#1/In_IN03_2004_04 *)
    E001_In_IN04_2004_05 : UINT;  (* RCON1（Node1） RCON→PLC 【IN04】共通 電源ユニット状態信号2; at ECAT://node#1/In_IN04_2004_05 *)
    E001_In_IN05_2004_06 : UINT;  (* RCON1（Node1） RCON→PLC 【IN05】共通 電源ユニット状態信号3; at ECAT://node#1/In_IN05_2004_06 *)
    E001_In_IN06_2004_07 : UINT;  (* RCON1（Node1） RCON→PLC 【IN06】共通 電源ユニット状態信号4／軽故障メンテナンス（設定依存）; at ECAT://node#1/In_IN06_2004_07 *)
    E001_In_IN07_2004_08 : UINT;  (* RCON1（Node1） RCON→PLC 【IN07】共通 共通予約領域（使用禁止・占有あり）; at ECAT://node#1/In_IN07_2004_08 *)
    E001_In_IN08_2004_09 : UINT;  (* RCON1（Node1） RCON→PLC 【IN08】1軸目（No.0） 現在位置 下位ワード; at ECAT://node#1/In_IN08_2004_09 *)
    E001_In_IN09_2004_0A : UINT;  (* RCON1（Node1） RCON→PLC 【IN09】1軸目（No.0） 現在位置 上位ワード; at ECAT://node#1/In_IN09_2004_0A *)
    E001_In_IN10_2004_0B : UINT;  (* RCON1（Node1） RCON→PLC 【IN10】1軸目（No.0） 現在電流 下位ワード（PCは指令電流）; at ECAT://node#1/In_IN10_2004_0B *)
    E001_In_IN11_2004_0C : UINT;  (* RCON1（Node1） RCON→PLC 【IN11】1軸目（No.0） 現在電流 上位ワード（PCは指令電流）; at ECAT://node#1/In_IN11_2004_0C *)
    E001_In_IN12_2004_0D : UINT;  (* RCON1（Node1） RCON→PLC 【IN12】1軸目（No.0） 現在速度（負方向は2の補数）; at ECAT://node#1/In_IN12_2004_0D *)
    E001_In_IN13_2004_0E : UINT;  (* RCON1（Node1） RCON→PLC 【IN13】1軸目（No.0） 予約領域（使用禁止）; at ECAT://node#1/In_IN13_2004_0E *)
    E001_In_IN14_2004_0F : UINT;  (* RCON1（Node1） RCON→PLC 【IN14】1軸目（No.0） アラームコード（簡易コードではない）; at ECAT://node#1/In_IN14_2004_0F *)
    E001_In_IN15_2004_10 : UINT;  (* RCON1（Node1） RCON→PLC 【IN15】1軸目（No.0） 軸状態信号（PEND・SV等）; at ECAT://node#1/In_IN15_2004_10 *)
    E001_In_IN16_2004_11 : UINT;  (* RCON1（Node1） RCON→PLC 【IN16】2軸目（No.1） 現在位置 下位ワード; at ECAT://node#1/In_IN16_2004_11 *)
    E001_In_IN17_2004_12 : UINT;  (* RCON1（Node1） RCON→PLC 【IN17】2軸目（No.1） 現在位置 上位ワード; at ECAT://node#1/In_IN17_2004_12 *)
    E001_In_IN18_2004_13 : UINT;  (* RCON1（Node1） RCON→PLC 【IN18】2軸目（No.1） 現在電流 下位ワード（PCは指令電流）; at ECAT://node#1/In_IN18_2004_13 *)
    E001_In_IN19_2004_14 : UINT;  (* RCON1（Node1） RCON→PLC 【IN19】2軸目（No.1） 現在電流 上位ワード（PCは指令電流）; at ECAT://node#1/In_IN19_2004_14 *)
    E001_In_IN20_2004_15 : UINT;  (* RCON1（Node1） RCON→PLC 【IN20】2軸目（No.1） 現在速度（負方向は2の補数）; at ECAT://node#1/In_IN20_2004_15 *)
    E001_In_IN21_2004_16 : UINT;  (* RCON1（Node1） RCON→PLC 【IN21】2軸目（No.1） 予約領域（使用禁止）; at ECAT://node#1/In_IN21_2004_16 *)
    E001_In_IN22_2004_17 : UINT;  (* RCON1（Node1） RCON→PLC 【IN22】2軸目（No.1） アラームコード（簡易コードではない）; at ECAT://node#1/In_IN22_2004_17 *)
    E001_In_IN23_2004_18 : UINT;  (* RCON1（Node1） RCON→PLC 【IN23】2軸目（No.1） 軸状態信号（PEND・SV等）; at ECAT://node#1/In_IN23_2004_18 *)
    E001_In_IN24_2004_19 : UINT;  (* RCON1（Node1） RCON→PLC 【IN24】3軸目（No.2） 現在位置 下位ワード; at ECAT://node#1/In_IN24_2004_19 *)
    E001_In_IN25_2004_1A : UINT;  (* RCON1（Node1） RCON→PLC 【IN25】3軸目（No.2） 現在位置 上位ワード; at ECAT://node#1/In_IN25_2004_1A *)
    E001_In_IN26_2004_1B : UINT;  (* RCON1（Node1） RCON→PLC 【IN26】3軸目（No.2） 現在電流 下位ワード（PCは指令電流）; at ECAT://node#1/In_IN26_2004_1B *)
    E001_In_IN27_2004_1C : UINT;  (* RCON1（Node1） RCON→PLC 【IN27】3軸目（No.2） 現在電流 上位ワード（PCは指令電流）; at ECAT://node#1/In_IN27_2004_1C *)
    E001_In_IN28_2004_1D : UINT;  (* RCON1（Node1） RCON→PLC 【IN28】3軸目（No.2） 現在速度（負方向は2の補数）; at ECAT://node#1/In_IN28_2004_1D *)
    E001_In_IN29_2004_1E : UINT;  (* RCON1（Node1） RCON→PLC 【IN29】3軸目（No.2） 予約領域（使用禁止）; at ECAT://node#1/In_IN29_2004_1E *)
    E001_In_IN30_2004_1F : UINT;  (* RCON1（Node1） RCON→PLC 【IN30】3軸目（No.2） アラームコード（簡易コードではない）; at ECAT://node#1/In_IN30_2004_1F *)
    E001_In_IN31_2004_20 : UINT;  (* RCON1（Node1） RCON→PLC 【IN31】3軸目（No.2） 軸状態信号（PEND・SV等）; at ECAT://node#1/In_IN31_2004_20 *)
    E001_In_IN32_2004_21 : UINT;  (* RCON1（Node1） RCON→PLC 【IN32】4軸目（No.3） 現在位置 下位ワード; at ECAT://node#1/In_IN32_2004_21 *)
    E001_In_IN33_2004_22 : UINT;  (* RCON1（Node1） RCON→PLC 【IN33】4軸目（No.3） 現在位置 上位ワード; at ECAT://node#1/In_IN33_2004_22 *)
    E001_In_IN34_2004_23 : UINT;  (* RCON1（Node1） RCON→PLC 【IN34】4軸目（No.3） 現在電流 下位ワード（PCは指令電流）; at ECAT://node#1/In_IN34_2004_23 *)
    E001_In_IN35_2004_24 : UINT;  (* RCON1（Node1） RCON→PLC 【IN35】4軸目（No.3） 現在電流 上位ワード（PCは指令電流）; at ECAT://node#1/In_IN35_2004_24 *)
    E001_In_IN36_2004_25 : UINT;  (* RCON1（Node1） RCON→PLC 【IN36】4軸目（No.3） 現在速度（負方向は2の補数）; at ECAT://node#1/In_IN36_2004_25 *)
    E001_In_IN37_2004_26 : UINT;  (* RCON1（Node1） RCON→PLC 【IN37】4軸目（No.3） 予約領域（使用禁止）; at ECAT://node#1/In_IN37_2004_26 *)
    E001_In_IN38_2004_27 : UINT;  (* RCON1（Node1） RCON→PLC 【IN38】4軸目（No.3） アラームコード（簡易コードではない）; at ECAT://node#1/In_IN38_2004_27 *)
    E001_In_IN39_2004_28 : UINT;  (* RCON1（Node1） RCON→PLC 【IN39】4軸目（No.3） 軸状態信号（PEND・SV等）; at ECAT://node#1/In_IN39_2004_28 *)
    E001_In_IN40_2004_29 : UINT;  (* RCON1（Node1） RCON→PLC 【IN40】5軸目（No.4） 現在位置 下位ワード; at ECAT://node#1/In_IN40_2004_29 *)
    E001_In_IN41_2004_2A : UINT;  (* RCON1（Node1） RCON→PLC 【IN41】5軸目（No.4） 現在位置 上位ワード; at ECAT://node#1/In_IN41_2004_2A *)
    E001_In_IN42_2004_2B : UINT;  (* RCON1（Node1） RCON→PLC 【IN42】5軸目（No.4） 現在電流 下位ワード（PCは指令電流）; at ECAT://node#1/In_IN42_2004_2B *)
    E001_In_IN43_2004_2C : UINT;  (* RCON1（Node1） RCON→PLC 【IN43】5軸目（No.4） 現在電流 上位ワード（PCは指令電流）; at ECAT://node#1/In_IN43_2004_2C *)
    E001_In_IN44_2004_2D : UINT;  (* RCON1（Node1） RCON→PLC 【IN44】5軸目（No.4） 現在速度（負方向は2の補数）; at ECAT://node#1/In_IN44_2004_2D *)
    E001_In_IN45_2004_2E : UINT;  (* RCON1（Node1） RCON→PLC 【IN45】5軸目（No.4） 予約領域（使用禁止）; at ECAT://node#1/In_IN45_2004_2E *)
    E001_In_IN46_2004_2F : UINT;  (* RCON1（Node1） RCON→PLC 【IN46】5軸目（No.4） アラームコード（簡易コードではない）; at ECAT://node#1/In_IN46_2004_2F *)
    E001_In_IN47_2004_30 : UINT;  (* RCON1（Node1） RCON→PLC 【IN47】5軸目（No.4） 軸状態信号（PEND・SV等）; at ECAT://node#1/In_IN47_2004_30 *)
    E001_In_IN48_2004_31 : UINT;  (* RCON1（Node1） RCON→PLC 【IN48】6軸目（No.5） 現在位置 下位ワード; at ECAT://node#1/In_IN48_2004_31 *)
    E001_In_IN49_2004_32 : UINT;  (* RCON1（Node1） RCON→PLC 【IN49】6軸目（No.5） 現在位置 上位ワード; at ECAT://node#1/In_IN49_2004_32 *)
    E001_In_IN50_2004_33 : UINT;  (* RCON1（Node1） RCON→PLC 【IN50】6軸目（No.5） 現在電流 下位ワード（PCは指令電流）; at ECAT://node#1/In_IN50_2004_33 *)
    E001_In_IN51_2004_34 : UINT;  (* RCON1（Node1） RCON→PLC 【IN51】6軸目（No.5） 現在電流 上位ワード（PCは指令電流）; at ECAT://node#1/In_IN51_2004_34 *)
    E001_In_IN52_2004_35 : UINT;  (* RCON1（Node1） RCON→PLC 【IN52】6軸目（No.5） 現在速度（負方向は2の補数）; at ECAT://node#1/In_IN52_2004_35 *)
    E001_In_IN53_2004_36 : UINT;  (* RCON1（Node1） RCON→PLC 【IN53】6軸目（No.5） 予約領域（使用禁止）; at ECAT://node#1/In_IN53_2004_36 *)
    E001_In_IN54_2004_37 : UINT;  (* RCON1（Node1） RCON→PLC 【IN54】6軸目（No.5） アラームコード（簡易コードではない）; at ECAT://node#1/In_IN54_2004_37 *)
    E001_In_IN55_2004_38 : UINT;  (* RCON1（Node1） RCON→PLC 【IN55】6軸目（No.5） 軸状態信号（PEND・SV等）; at ECAT://node#1/In_IN55_2004_38 *)
    E001_In_IN56_2004_39 : UINT;  (* RCON1（Node1） 【IN56】用途未確認領域。今回の軸データ変換では未使用。; at ECAT://node#1/In_IN56_2004_39 *)
    E001_In_IN57_2004_3A : UINT;  (* RCON1（Node1） 【IN57】用途未確認領域。今回の軸データ変換では未使用。; at ECAT://node#1/In_IN57_2004_3A *)
    E001_In_IN58_2004_3B : UINT;  (* RCON1（Node1） 【IN58】用途未確認領域。今回の軸データ変換では未使用。; at ECAT://node#1/In_IN58_2004_3B *)
    E001_In_IN59_2004_3C : UINT;  (* RCON1（Node1） 【IN59】用途未確認領域。今回の軸データ変換では未使用。; at ECAT://node#1/In_IN59_2004_3C *)
    E001_In_IN60_2004_3D : UINT;  (* RCON1（Node1） 【IN60】用途未確認領域。今回の軸データ変換では未使用。; at ECAT://node#1/In_IN60_2004_3D *)
    E001_In_IN61_2004_3E : UINT;  (* RCON1（Node1） 【IN61】用途未確認領域。今回の軸データ変換では未使用。; at ECAT://node#1/In_IN61_2004_3E *)
    E001_In_IN62_2004_3F : UINT;  (* RCON1（Node1） 【IN62】用途未確認領域。今回の軸データ変換では未使用。; at ECAT://node#1/In_IN62_2004_3F *)
    E001_In_IN63_2004_40 : UINT;  (* RCON1（Node1） 【IN63】用途未確認領域。今回の軸データ変換では未使用。; at ECAT://node#1/In_IN63_2004_40 *)
    E001_In_IN64_2004_41 : UINT;  (* RCON1（Node1） 【IN64】用途未確認領域。今回の軸データ変換では未使用。; at ECAT://node#1/In_IN64_2004_41 *)
    E001_In_IN65_2004_42 : UINT;  (* RCON1（Node1） 【IN65】用途未確認領域。今回の軸データ変換では未使用。; at ECAT://node#1/In_IN65_2004_42 *)
    E001_In_IN66_2004_43 : UINT;  (* RCON1（Node1） 【IN66】用途未確認領域。今回の軸データ変換では未使用。; at ECAT://node#1/In_IN66_2004_43 *)
    E001_In_IN67_2004_44 : UINT;  (* RCON1（Node1） 【IN67】用途未確認領域。今回の軸データ変換では未使用。; at ECAT://node#1/In_IN67_2004_44 *)
    E001_In_IN68_2004_45 : UINT;  (* RCON1（Node1） 【IN68】用途未確認領域。今回の軸データ変換では未使用。; at ECAT://node#1/In_IN68_2004_45 *)
    E001_In_IN69_2004_46 : UINT;  (* RCON1（Node1） 【IN69】用途未確認領域。今回の軸データ変換では未使用。; at ECAT://node#1/In_IN69_2004_46 *)
    E001_In_IN70_2004_47 : UINT;  (* RCON1（Node1） 【IN70】用途未確認領域。今回の軸データ変換では未使用。; at ECAT://node#1/In_IN70_2004_47 *)
    E001_In_IN71_2004_48 : UINT;  (* RCON1（Node1） 【IN71】用途未確認領域。今回の軸データ変換では未使用。; at ECAT://node#1/In_IN71_2004_48 *)
    RCON1_RxRaw : ARRAY[0..71] OF UINT;  (* RCON1：E001入力を読取った通信値。書換えない。 *)
    RCON1_RxWord : ARRAY[0..71] OF WORD;  (* RCON1：バイト順を正規化した論理入力ワード。 *)
    RCON1_TxWord : ARRAY[0..55] OF WORD;  (* RCON1：内部値から作成した論理出力ワード。 *)
    RCON1_TxUInt : ARRAY[0..55] OF UINT;  (* RCON1：バイト順を適用した送信候補。実I/Oそのものではない。 *)
    RCON1_LayoutConfirmed : BOOL;  (* RCON1：初期FALSE。全6軸直接数値指定・共通8W・軸順・占有を確認して設定。 *)
    RCON1_ByteOrderConfirmed : BOOL;  (* RCON1：初期FALSE。既知の位置とbitでワード順・バイト順を確認して設定。 *)
    RCON1_SwapBytes : BOOL;  (* RCON1：初期FALSEは仮値。1ワード内のバイト交換が必要か実機で確認。 *)
    RCON1_CommOK : BOOL;  (* RCON1：初期FALSE。CPUの実EtherCAT通信状態から別途作成。TRUE固定禁止。 *)
    RCON1_GwMON_Request : BOOL;  (* RCON1：初期FALSE。ゲートウェイMON要求。論理b15。安全停止ではない。 *)
    RCON1_GwRTE_Request : BOOL;  (* RCON1：初期FALSE。ゲートウェイ通信異常ラッチ解除要求。論理b13。 *)
    RCON1_GwRun : BOOL;  (* RCON1：入力：ゲートウェイ正常動作中RUN。 *)
    RCON1_GwControllerCommLatch : BOOL;  (* RCON1：入力：運転中ERR-C保持LERC。 *)
    RCON1_GwAxisCommError : BOOL;  (* RCON1：入力：ゲートウェイと軸の通信異常ERRT。 *)
    RCON1_GwManual : BOOL;  (* RCON1：入力：MANUスイッチ選択MOD。 *)
    RCON1_GwHeavyAlarm : BOOL;  (* RCON1：入力：再起動が必要なゲートウェイ異常ALMH。 *)
    RCON1_GwLightAlarm : BOOL;  (* RCON1：入力：ゲートウェイ軽微異常ALML。 *)
    RCON1_GwSystemStop : BOOL;  (* RCON1：入力：システムSTOP入力による停止状態SEMG。安全回路の代用不可。 *)
    RCON1_GwAlarmCode : UINT;  (* RCON1：入力：ゲートウェイALMCの下位8bit。軸AlarmCodeとは別。 *)
    RCON1_AxisLinked : ARRAY[1..6] OF BOOL;  (* RCON1：入力：軸No.0～5のリンク状態。 *)
    RCON1_PowerStateRaw : ARRAY[0..4] OF WORD;  (* RCON1：入力IN02～06の正規化済み生ワード。詳細意味は構成依存。 *)
    RCON1_EncodeOK : ARRAY[1..6] OF BOOL;  (* RCON1：通信形式へ数値変換できたか。安全・運転許可ではない。 *)
    RCON1_EncodeError : ARRAY[1..6] OF UINT;  (* RCON1：変換エラー番号。0正常、1単位、2位置、3幅、4速度、5加減速、6押付け、7両方向ジョグ。 *)
    RCON1_WriteEnable : BOOL;  (* RCON1：初期FALSE。実出力への書込みを許可。OFFは出力更新保留であり停止ではない。 *)
    RCON1_GwApply : BOOL;  (* RCON1：初期FALSE。共通MON/RTEワードを書込む。 *)
    RCON1_AxisApply : ARRAY[1..6] OF BOOL;  (* RCON1：初期FALSE。指定軸の8ワードを書込む。OFFは停止ではない。 *)
    RCON1_MotionPermit : ARRAY[1..6] OF BOOL;  (* RCON1：初期FALSE。機械範囲・安全・運転条件から別途作成する運転許可。単純TRUE固定禁止。 *)
    RCON1_GwWritten : BOOL;  (* RCON1：共通出力へ代入したサイクルのみTRUE。RCON受付の意味ではない。 *)
    RCON1_AxisWritten : ARRAY[1..6] OF BOOL;  (* RCON1：各軸出力へ代入したサイクルのみTRUE。RCON受付・完了ではない。 *)
    RCON2_RxRaw : ARRAY[0..47] OF UINT;  (* RCON2：E005（末尾_1）入力を読取った通信値。書換えない。 *)
    RCON2_RxWord : ARRAY[0..47] OF WORD;  (* RCON2：バイト順を正規化した論理入力ワード。 *)
    RCON2_TxWord : ARRAY[0..47] OF WORD;  (* RCON2：内部値から作成した論理出力ワード。 *)
    RCON2_TxUInt : ARRAY[0..47] OF UINT;  (* RCON2：バイト順を適用した送信候補。実I/Oそのものではない。 *)
    RCON2_LayoutConfirmed : BOOL;  (* RCON2：初期FALSE。全5軸直接数値指定・共通8W・軸順・占有を確認して設定。 *)
    RCON2_ByteOrderConfirmed : BOOL;  (* RCON2：初期FALSE。既知の位置とbitでワード順・バイト順を確認して設定。 *)
    RCON2_SwapBytes : BOOL;  (* RCON2：初期FALSEは仮値。1ワード内のバイト交換が必要か実機で確認。 *)
    RCON2_CommOK : BOOL;  (* RCON2：初期FALSE。CPUの実EtherCAT通信状態から別途作成。TRUE固定禁止。 *)
    RCON2_GwMON_Request : BOOL;  (* RCON2：初期FALSE。ゲートウェイMON要求。論理b15。安全停止ではない。 *)
    RCON2_GwRTE_Request : BOOL;  (* RCON2：初期FALSE。ゲートウェイ通信異常ラッチ解除要求。論理b13。 *)
    RCON2_GwRun : BOOL;  (* RCON2：入力：ゲートウェイ正常動作中RUN。 *)
    RCON2_GwControllerCommLatch : BOOL;  (* RCON2：入力：運転中ERR-C保持LERC。 *)
    RCON2_GwAxisCommError : BOOL;  (* RCON2：入力：ゲートウェイと軸の通信異常ERRT。 *)
    RCON2_GwManual : BOOL;  (* RCON2：入力：MANUスイッチ選択MOD。 *)
    RCON2_GwHeavyAlarm : BOOL;  (* RCON2：入力：再起動が必要なゲートウェイ異常ALMH。 *)
    RCON2_GwLightAlarm : BOOL;  (* RCON2：入力：ゲートウェイ軽微異常ALML。 *)
    RCON2_GwSystemStop : BOOL;  (* RCON2：入力：システムSTOP入力による停止状態SEMG。安全回路の代用不可。 *)
    RCON2_GwAlarmCode : UINT;  (* RCON2：入力：ゲートウェイALMCの下位8bit。軸AlarmCodeとは別。 *)
    RCON2_AxisLinked : ARRAY[1..5] OF BOOL;  (* RCON2：入力：軸No.0～4のリンク状態。 *)
    RCON2_PowerStateRaw : ARRAY[0..4] OF WORD;  (* RCON2：入力IN02～06の正規化済み生ワード。詳細意味は構成依存。 *)
    RCON2_EncodeOK : ARRAY[1..5] OF BOOL;  (* RCON2：通信形式へ数値変換できたか。安全・運転許可ではない。 *)
    RCON2_EncodeError : ARRAY[1..5] OF UINT;  (* RCON2：変換エラー番号。0正常、1単位、2位置、3幅、4速度、5加減速、6押付け、7両方向ジョグ。 *)
    RCON2_WriteEnable : BOOL;  (* RCON2：初期FALSE。実出力への書込みを許可。OFFは出力更新保留であり停止ではない。 *)
    RCON2_GwApply : BOOL;  (* RCON2：初期FALSE。共通MON/RTEワードを書込む。 *)
    RCON2_AxisApply : ARRAY[1..5] OF BOOL;  (* RCON2：初期FALSE。指定軸の8ワードを書込む。OFFは停止ではない。 *)
    RCON2_MotionPermit : ARRAY[1..5] OF BOOL;  (* RCON2：初期FALSE。機械範囲・安全・運転条件から別途作成する運転許可。単純TRUE固定禁止。 *)
    RCON2_GwWritten : BOOL;  (* RCON2：共通出力へ代入したサイクルのみTRUE。RCON受付の意味ではない。 *)
    RCON2_AxisWritten : ARRAY[1..5] OF BOOL;  (* RCON2：各軸出力へ代入したサイクルのみTRUE。RCON受付・完了ではない。 *)
END_VAR

PROGRAM ModeManagement_モード管理
VAR
    Setting_M : BOOL;
    Manual_M : BOOL;
    Auto_M : BOOL;
    Dummy_M : BOOL;
    Inital_M : BOOL;
    Output_Error_M : ARRAY[0..99] OF Bool;
    Index_Error_001 : DINT;
    Index_B_001 : DINT;
    Index_Share_001 : DINT;
    Error_TON : ARRAY[0..99] OF TON;
    Error_M : ARRAY[0..99] OF Bool;  (* エラー：; [1] シリンダ; [2] コンベア＆ドアセンサ; [3] FH; [4] A(左側)検査コンベア ワーク不一致 *)
    Error_TOF : ARRAY[0..99] OF TOF;
    AutoMode_A_M : ARRAY[0..99] OF Bool;
END_VAR
VAR_EXTERNAL
    Output_A_Error_M : ARRAY[0..99] OF Bool;
    Output_A_Restart_M : ARRAY[0..99] OF Bool;
    In_Sw_RESET : BOOL;
    In_Sw_START : BOOL;
    ManualMode : BOOL;
    M9999 : BOOL;
    Output_B_Error_M : ARRAY[0..99] OF Bool;  (* B(右側)シリンダエラー *)
    Output_B_Restart_M : ARRAY[0..99] OF Bool;  (* B(右側)シリンダ再開： *)
    Output_Share_Error_M : ARRAY[0..99] OF Bool;
    Output_Share_Restart_M : ARRAY[0..99] OF Bool;
    TimerQ_In_Sen_Accum_CV_A_Full : BOOL;
    Out_TDC_Stop : BOOL;
    In_Sen_Unl_Conv_A_Pass : BOOL;
    In_Sen_Accum_CV_A_Full : BOOL;
    In_Sen_Unl_Conv_B_Pass : BOOL;
    Pause : ARRAY[0..99] OF Bool;
    AutoMode : BOOL;
    In_Sen_DOOR_01 : BOOL;
    In_Sen_DOOR_02 : BOOL;
    In_Sen_DOOR_03 : BOOL;
    In_Sen_DOOR_04 : BOOL;
    In_Sen_DOOR_05 : BOOL;
    In_Sen_DOOR_06 : BOOL;
    In_Sw_EMS1 : BOOL;
    In_Sw_EMS2 : BOOL;
    In_Sw_EMS3 : BOOL;
    In_Sen_AIR１_Pressure_01 : BOOL;
    In_Sen_AIR１_Pressure_02 : BOOL;
    In_Sen_AIR１_Pressure_03 : BOOL;
    TEST_M : ARRAY[0..99] OF Bool;
    ST0_Sup_Start : BOOL;  (* ST0_動作開始 *)
    Out_CYw_Sply_Pick_A_H_Auto : ARRAY[0..10] OF Bool;
    Out_CYw_Sply_Pick_A_H_Done : BOOL;
    Out_CYw_Sply_Slide_A_H_Auto : ARRAY[0..10] OF Bool;
    Out_CYw_Sply_Slide_A_H_Done : BOOL;
    Out_CYw_Sup_Chuck_A_Cl_H_Auto : ARRAY[0..10] OF Bool;
    Out_CYw_Sup_Chuck_A_Cl_H_Done : BOOL;
    In_Sen_Accum_CV_A_Arrival : BOOL;
    In_Sen_Work_A_Pos_00 : BOOL;
    Out_CYw_Sply_Pick_A_F_Auto : ARRAY[0..10] OF Bool;
    Out_CYw_Sply_Pick_A_F_Done : BOOL;
    Out_CYw_Sup_Chuck_A_Cl_F_Auto : ARRAY[0..10] OF Bool;
    Out_CYw_Sup_Chuck_A_Cl_F_Done : BOOL;
    Out_CYw_Sply_Slide_A_F_Auto : ARRAY[0..10] OF Bool;
    Out_CYw_Sply_Slide_A_F_Done : BOOL;
    Ins_A_Cv_Error : BOOL;
    Station_A_Data : ARRAY[0..8] OF sData;
    Ins_A_Cv_M : ARRAY[0..99] OF Bool;
    HMI_MessageNo : ARRAY[0..9] OF UINT;
    FH_5552_10_A_Auto : BOOL;
    In_Sen_Accum_CV_B_Full : BOOL;
    FH_Line3_Error_Status_1 : BOOL;
    FH_Line0_Error_Status_1 : BOOL;
    FH_Line1_Error_Status_1 : BOOL;
    FH_Line2_Error_Status_1 : BOOL;
    FH_Line0_Error_Clear_1 : BOOL;
    FH_Line1_Error_Clear_1 : BOOL;
    FH_Line2_Error_Clear_1 : BOOL;
    FH_Line3_Error_Clear_1 : BOOL;
    Ins_A_Next_Cycle : BOOL;
    OriginDone : BOOL;  (* 原点復帰完了 *)
    DummyDone : BOOL;  (* ダミーチェック完了 *)
    HMI_CurrentPage : STRING[256];
    Ins_A_End : BOOL;
    Auto_A_Start : BOOL;  (* 自動運転 開始 *)
    Auto_Ready : BOOL;  (* 自動運転可能 *)
    ST0_A_Sup_Busy : BOOL;
    ST1_A_Ca1_Busy : BOOL;
END_VAR
VAR
    _e1 : R_TRIG;
    _p2 : BOOL;
    _e3 : R_TRIG;
    _e4 : R_TRIG;
    _e5 : R_TRIG;
    _e6 : R_TRIG;
    _e7 : R_TRIG;
    _e8 : R_TRIG;
    _e9 : R_TRIG;
    _e10 : R_TRIG;
    _e11 : R_TRIG;
    _p12 : BOOL;
    _p13 : BOOL;
    _e14 : R_TRIG;
    _p15 : BOOL;
    _e16 : R_TRIG;
    _e17 : R_TRIG;
    _e18 : R_TRIG;
    _e19 : R_TRIG;
    _e20 : R_TRIG;
    _e21 : R_TRIG;
    _e22 : R_TRIG;
    _p23 : BOOL;
END_VAR

(* Section Initial_初期化処理: ladder, written here as Structured Text *)

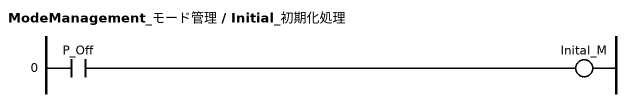
(* Rung 0 *)
Inital_M := P_Off;

(* Section DummyCheck_ダミーチェック: ladder, written here as Structured Text *)

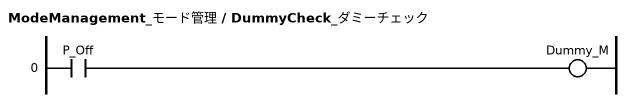
(* Rung 0 *)
Dummy_M := P_Off;

(* Section AutoMode_自動運転: ladder, written here as Structured Text *)

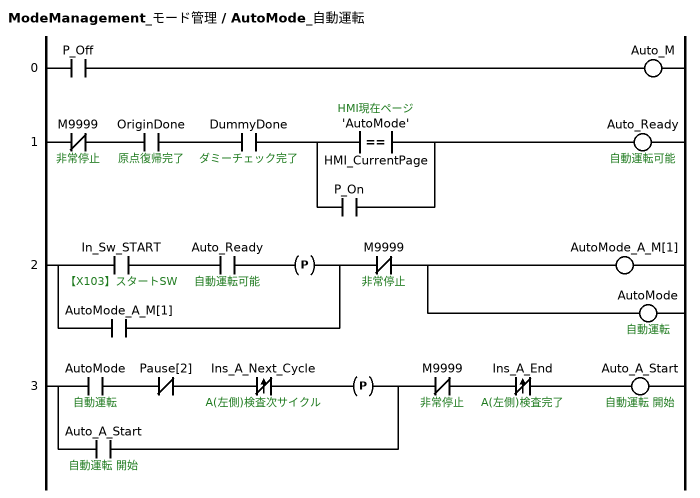
(* Rung 0 *)
Auto_M := P_Off;
(* Rung 1 *)
Auto_Ready := NOT M9999 AND OriginDone AND DummyDone AND (('AutoMode' = HMI_CurrentPage) OR P_On);
(* Rung 2 *)
_e1(CLK := In_Sw_START AND Auto_Ready);
_p2 := (_e1.Q OR AutoMode_A_M[1]) AND NOT M9999;
AutoMode_A_M[1] := _p2;
AutoMode := _p2;
(* Rung 3 *)
_e3(CLK := Ins_A_Next_Cycle);
_e4(CLK := AutoMode AND NOT Pause[2] AND NOT _e3.Q);
_e5(CLK := Ins_A_End);
Auto_A_Start := (_e4.Q OR Auto_A_Start) AND NOT M9999 AND NOT _e5.Q;

(* Section Manual_手動運転: ladder, written here as Structured Text *)

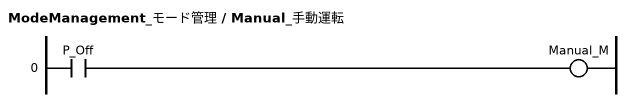
(* Rung 0 *)
Manual_M := P_Off;

(* Section Setting_設定: ladder, written here as Structured Text *)

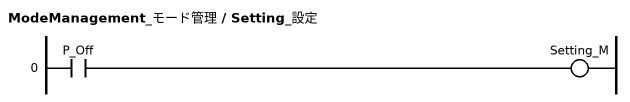
(* Rung 0 *)
Setting_M := P_Off;

(* Section Error_エラー処理: ladder, written here as Structured Text *)

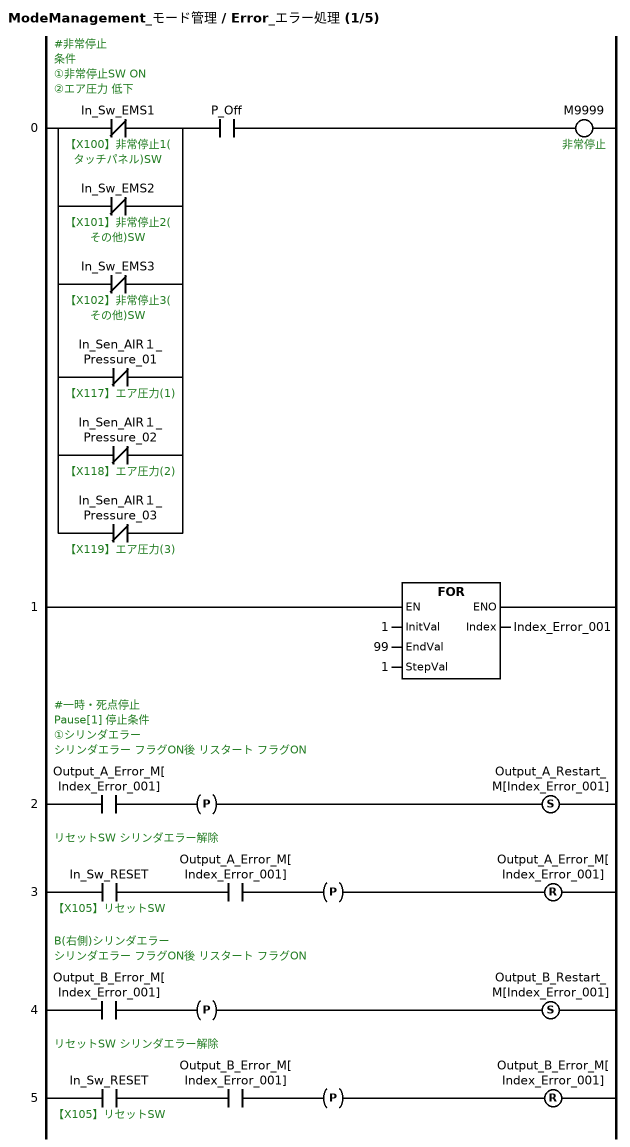
(* Rung 0: #非常停止 / 条件 / ①非常停止SW ON / ②エア圧力 低下 *)
M9999 := (NOT In_Sw_EMS1 OR NOT In_Sw_EMS2 OR NOT In_Sw_EMS3 OR NOT In_Sen_AIR１_Pressure_01 OR NOT In_Sen_AIR１_Pressure_02 OR NOT In_Sen_AIR１_Pressure_03) AND P_Off;
(* Rung 1 *)
Index_Error_001 := FOR(InitVal := 1, EndVal := 99, StepVal := 1);
(* Rung 2: #一時・死点停止 / Pause[1] 停止条件 / ①シリンダエラー / シリンダエラー フラグON後 リスタート フラグON *)
_e6(CLK := Output_A_Error_M[Index_Error_001]);
IF _e6.Q THEN Output_A_Restart_M[Index_Error_001] := TRUE; END_IF;
(* Rung 3: リセットSW シリンダエラー解除 *)
_e7(CLK := In_Sw_RESET AND Output_A_Error_M[Index_Error_001]);
IF _e7.Q THEN Output_A_Error_M[Index_Error_001] := FALSE; END_IF;
(* Rung 4: B(右側)シリンダエラー / シリンダエラー フラグON後 リスタート フラグON *)
_e8(CLK := Output_B_Error_M[Index_Error_001]);
IF _e8.Q THEN Output_B_Restart_M[Index_Error_001] := TRUE; END_IF;
(* Rung 5: リセットSW シリンダエラー解除 *)
_e9(CLK := In_Sw_RESET AND Output_B_Error_M[Index_Error_001]);
IF _e9.Q THEN Output_B_Error_M[Index_Error_001] := FALSE; END_IF;

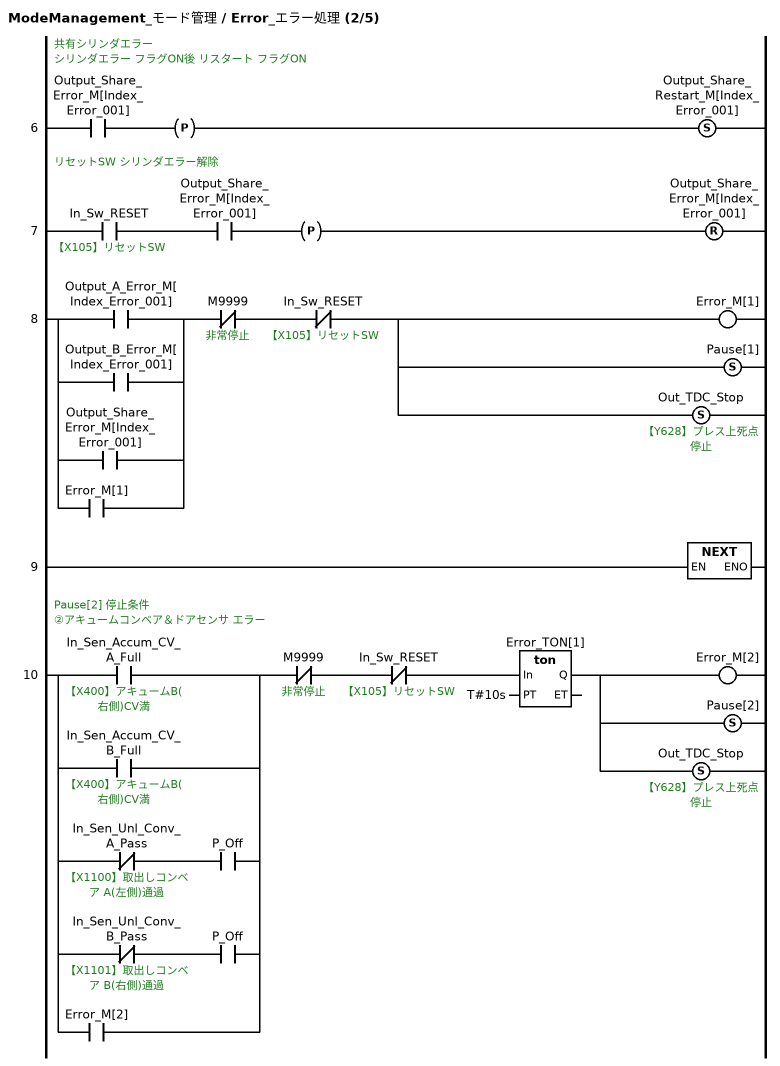
(* Rung 6: 共有シリンダエラー / シリンダエラー フラグON後 リスタート フラグON *)
_e10(CLK := Output_Share_Error_M[Index_Error_001]);
IF _e10.Q THEN Output_Share_Restart_M[Index_Error_001] := TRUE; END_IF;
(* Rung 7: リセットSW シリンダエラー解除 *)
_e11(CLK := In_Sw_RESET AND Output_Share_Error_M[Index_Error_001]);
IF _e11.Q THEN Output_Share_Error_M[Index_Error_001] := FALSE; END_IF;
(* Rung 8 *)
_p12 := (Output_A_Error_M[Index_Error_001] OR Output_B_Error_M[Index_Error_001] OR Output_Share_Error_M[Index_Error_001] OR Error_M[1]) AND NOT M9999 AND NOT In_Sw_RESET;
Error_M[1] := _p12;
IF _p12 THEN
    Pause[1] := TRUE;
    Out_TDC_Stop := TRUE;
END_IF;
(* Rung 9 *)
NEXT();
(* Rung 10: Pause[2] 停止条件 / ②アキュームコンベア＆ドアセンサ エラー *)
Error_TON[1](In := (In_Sen_Accum_CV_A_Full OR In_Sen_Accum_CV_B_Full OR (NOT In_Sen_Unl_Conv_A_Pass AND P_Off) OR (NOT In_Sen_Unl_Conv_B_Pass AND P_Off) OR Error_M[2]) AND NOT M9999 AND NOT In_Sw_RESET, PT := T#10s);
Error_M[2] := Error_TON[1].Q;
IF Error_TON[1].Q THEN
    Pause[2] := TRUE;
    Out_TDC_Stop := TRUE;
END_IF;

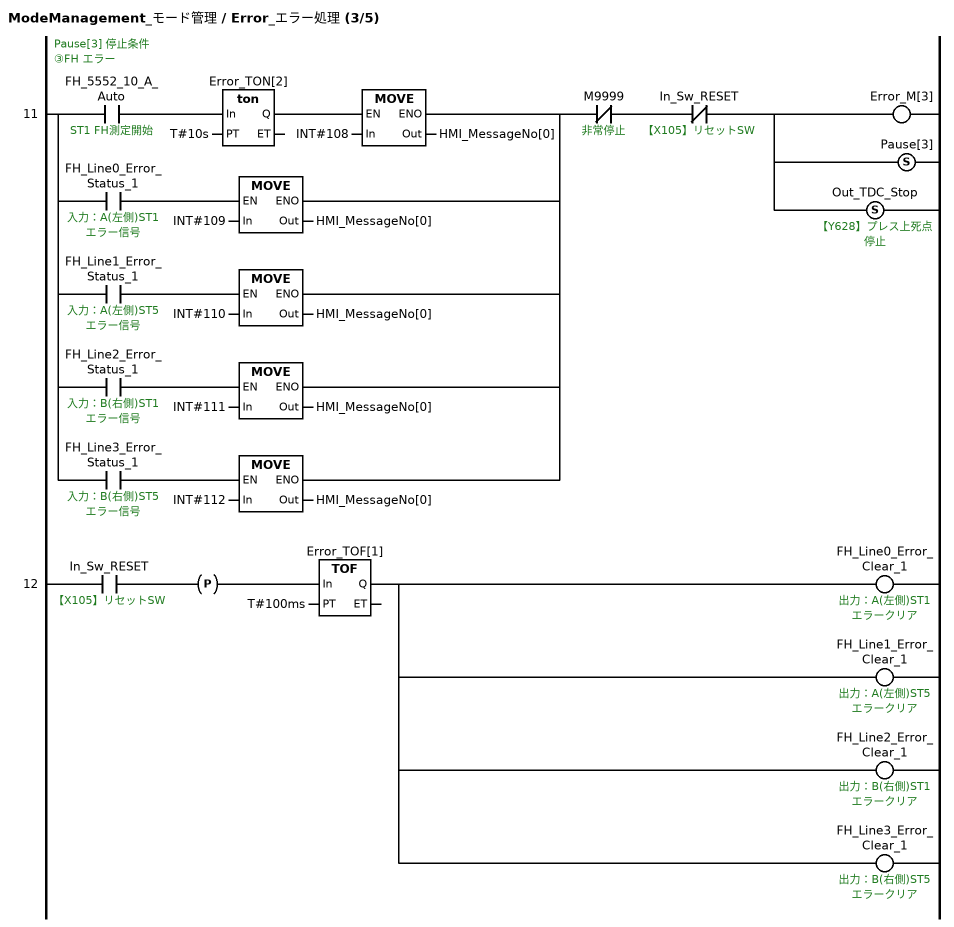
(* Rung 11: Pause[3] 停止条件 / ③FH エラー *)
Error_TON[2](In := FH_5552_10_A_Auto, PT := T#10s);
IF Error_TON[2].Q THEN HMI_MessageNo[0] := INT#108; END_IF;
IF FH_Line0_Error_Status_1 THEN HMI_MessageNo[0] := INT#109; END_IF;
IF FH_Line1_Error_Status_1 THEN HMI_MessageNo[0] := INT#110; END_IF;
IF FH_Line2_Error_Status_1 THEN HMI_MessageNo[0] := INT#111; END_IF;
IF FH_Line3_Error_Status_1 THEN HMI_MessageNo[0] := INT#112; END_IF;
_p13 := (Error_TON[2].Q OR FH_Line0_Error_Status_1 OR FH_Line1_Error_Status_1 OR FH_Line2_Error_Status_1 OR FH_Line3_Error_Status_1) AND NOT M9999 AND NOT In_Sw_RESET;
Error_M[3] := _p13;
IF _p13 THEN
    Pause[3] := TRUE;
    Out_TDC_Stop := TRUE;
END_IF;
(* Rung 12 *)
_e14(CLK := In_Sw_RESET);
Error_TOF[1](In := _e14.Q, PT := T#100ms);
FH_Line0_Error_Clear_1 := Error_TOF[1].Q;
FH_Line1_Error_Clear_1 := Error_TOF[1].Q;
FH_Line2_Error_Clear_1 := Error_TOF[1].Q;
FH_Line3_Error_Clear_1 := Error_TOF[1].Q;

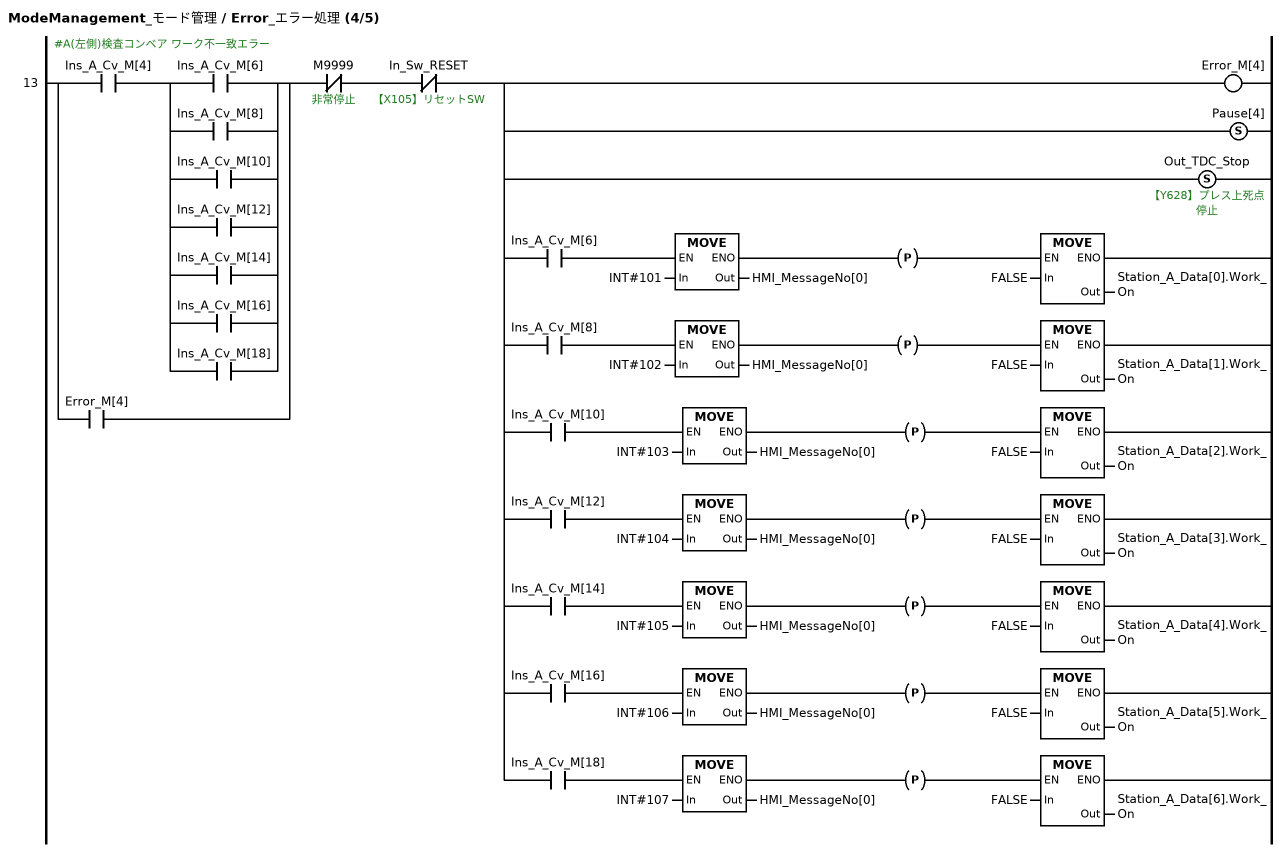
(* Rung 13: #A(左側)検査コンベア ワーク不一致エラー *)
_p15 := ((Ins_A_Cv_M[4] AND (Ins_A_Cv_M[6] OR Ins_A_Cv_M[8] OR Ins_A_Cv_M[10] OR Ins_A_Cv_M[12] OR Ins_A_Cv_M[14] OR Ins_A_Cv_M[16] OR Ins_A_Cv_M[18])) OR Error_M[4]) AND NOT M9999 AND NOT In_Sw_RESET;
Error_M[4] := _p15;
IF _p15 THEN
    Pause[4] := TRUE;
    Out_TDC_Stop := TRUE;
END_IF;
IF _p15 AND Ins_A_Cv_M[6] THEN HMI_MessageNo[0] := INT#101; END_IF;
_e16(CLK := _p15 AND Ins_A_Cv_M[6]);
IF _e16.Q THEN Station_A_Data[0].Work_On := FALSE; END_IF;
IF _p15 AND Ins_A_Cv_M[8] THEN HMI_MessageNo[0] := INT#102; END_IF;
_e17(CLK := _p15 AND Ins_A_Cv_M[8]);
IF _e17.Q THEN Station_A_Data[1].Work_On := FALSE; END_IF;
IF _p15 AND Ins_A_Cv_M[10] THEN HMI_MessageNo[0] := INT#103; END_IF;
_e18(CLK := _p15 AND Ins_A_Cv_M[10]);
IF _e18.Q THEN Station_A_Data[2].Work_On := FALSE; END_IF;
IF _p15 AND Ins_A_Cv_M[12] THEN HMI_MessageNo[0] := INT#104; END_IF;
_e19(CLK := _p15 AND Ins_A_Cv_M[12]);
IF _e19.Q THEN Station_A_Data[3].Work_On := FALSE; END_IF;
IF _p15 AND Ins_A_Cv_M[14] THEN HMI_MessageNo[0] := INT#105; END_IF;
_e20(CLK := _p15 AND Ins_A_Cv_M[14]);
IF _e20.Q THEN Station_A_Data[4].Work_On := FALSE; END_IF;
IF _p15 AND Ins_A_Cv_M[16] THEN HMI_MessageNo[0] := INT#106; END_IF;
_e21(CLK := _p15 AND Ins_A_Cv_M[16]);
IF _e21.Q THEN Station_A_Data[5].Work_On := FALSE; END_IF;
IF _p15 AND Ins_A_Cv_M[18] THEN HMI_MessageNo[0] := INT#107; END_IF;
_e22(CLK := _p15 AND Ins_A_Cv_M[18]);
IF _e22.Q THEN Station_A_Data[6].Work_On := FALSE; END_IF;

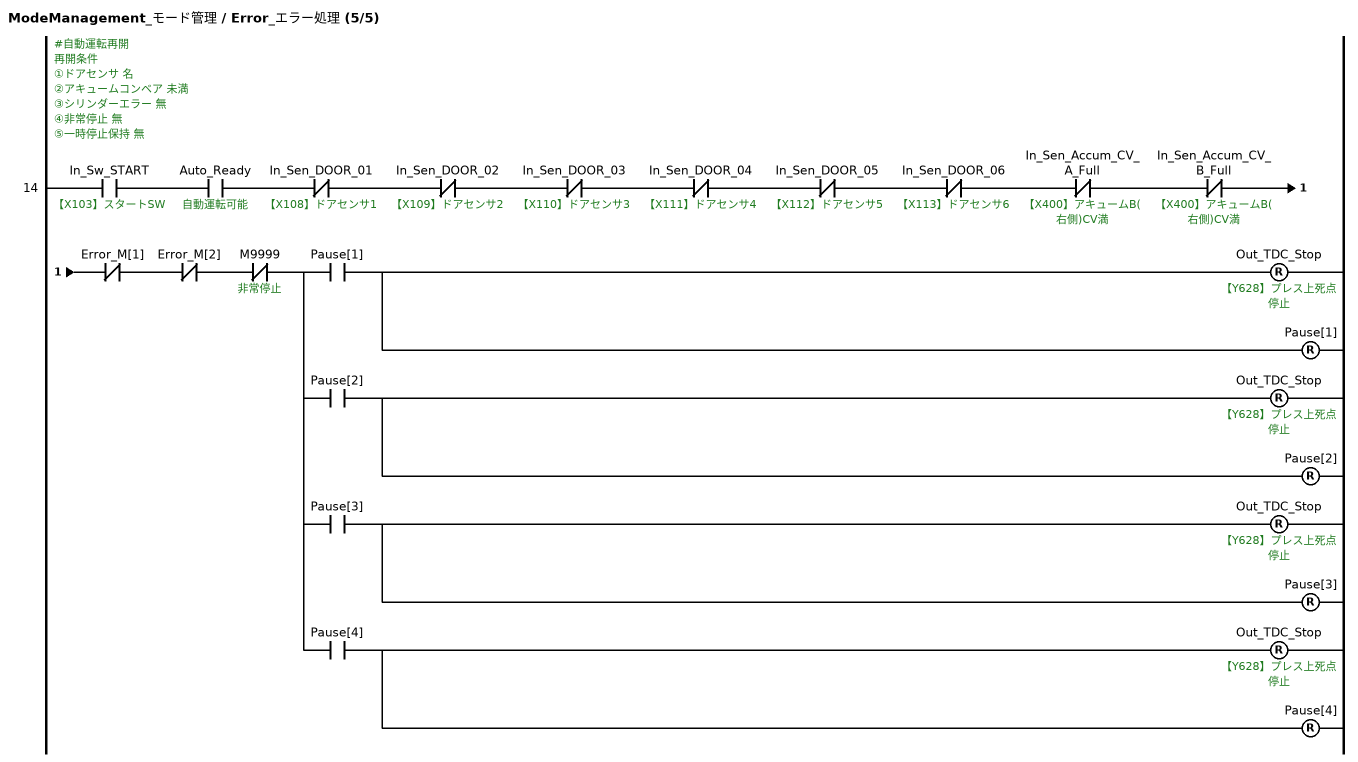
(* Rung 14: #自動運転再開 / 再開条件 / ①ドアセンサ 名 / ②アキュームコンベア 未満 / ③シリンダーエラー 無 / ④非常停止 無 / ⑤一時停止保持 無 *)
_p23 := In_Sw_START AND Auto_Ready AND NOT In_Sen_DOOR_01 AND NOT In_Sen_DOOR_02 AND NOT In_Sen_DOOR_03 AND NOT In_Sen_DOOR_04 AND NOT In_Sen_DOOR_05 AND NOT In_Sen_DOOR_06 AND NOT In_Sen_Accum_CV_A_Full AND NOT In_Sen_Accum_CV_B_Full AND NOT Error_M[1] AND NOT Error_M[2] AND NOT M9999;
IF _p23 AND Pause[1] THEN
    Out_TDC_Stop := FALSE;
    Pause[1] := FALSE;
END_IF;
IF _p23 AND Pause[2] THEN
    Out_TDC_Stop := FALSE;
    Pause[2] := FALSE;
END_IF;
IF _p23 AND Pause[3] THEN
    Out_TDC_Stop := FALSE;
    Pause[3] := FALSE;
END_IF;
IF _p23 AND Pause[4] THEN
    Out_TDC_Stop := FALSE;
    Pause[4] := FALSE;
END_IF;
END_PROGRAM

PROGRAM Movements_動作
VAR
    Mo_M : BOOL;
    ST0_A_Sup_M : ARRAY[0..99] OF Bool;  (* [4] 原点位置移動完了 *)
    ST1_Ins_Cv_Rdy : BOOL;
    ST2_Ins_Cv_Rdy : BOOL;
    ST3_Ins_Cv_Rdy : BOOL;
    ST4_Ins_Cv_Rdy : BOOL;
    ST5_Ins_Cv_Rdy : BOOL;
    ST6_Ins_Cv_Rdy : BOOL;
    ST7_Ins_Cv_Rdy : BOOL;
    Ins_A_Cv_T : ARRAY[0..99] OF TON;
    ST1_A_Ca1_Rdy : BOOL;
    ST1_A_Ca1_M : ARRAY[0..99] OF Bool;  (* [6] ST1 FH測定開始; [3] ワーク有無 判定; [1] ST1 A カメラ1 検査開始; [4] ST1 A ワーク有; [5] ST1 A ワーク無; [2] 【Y720】位置1A(左側)ストッパー 戻 *)
    ST2_A_Hgt_M : ARRAY[0..99] OF Bool;  (* [4] 【Y721】位置2A(左側)ストッパー戻; [6] ST1 A ワーク有; [7] ST1 A ワーク無; [5] ワーク有無 判定; [8] 【Y703】高さ検査A(左側)持上行; [9] 【Y701】高さ検査A(左側)押え行; [10] 高さ検査A(左側)OK判定; [11] 高さ検査A(左側)NG判定; [2] 【Y701】高さ検査A(左側)押え行 *)
    ST3_A_Dis1_M : ARRAY[0..99] OF Bool;
    GT2_A_Inspection_GetTime : DATE_AND_TIME;
    GT2_A_Inspection_GetTime_ST : STRING[256];
    GT2_A_Inspection_GetTime_ST_Del : STRING[20];
END_VAR
VAR_EXTERNAL
    ST0_Sup_Start : BOOL;  (* ST0_動作開始 *)
    M9999 : BOOL;
    Out_CYw_Sply_Pick_A_H_Auto : ARRAY[0..10] OF Bool;
    Out_CYw_Sply_Pick_A_H_Done : BOOL;
    Out_CYw_Sply_Slide_A_H_Auto : ARRAY[0..10] OF Bool;
    Out_CYw_Sply_Slide_A_H_Done : BOOL;
    Out_CYw_Sup_Chuck_A_Cl_H_Auto : ARRAY[0..10] OF Bool;
    Out_CYw_Sup_Chuck_A_Cl_H_Done : BOOL;
    In_Sen_Accum_CV_A_Arrival : BOOL;
    In_Sen_Work_A_Pos_00 : BOOL;
    Out_CYw_Sply_Pick_A_F_Auto : ARRAY[0..10] OF Bool;
    Out_CYw_Sply_Pick_A_F_Done : BOOL;
    Out_CYw_Sup_Chuck_A_Cl_F_Auto : ARRAY[0..10] OF Bool;
    Out_CYw_Sup_Chuck_A_Cl_F_Done : BOOL;
    Out_CYw_Sply_Slide_A_F_Auto : ARRAY[0..10] OF Bool;
    Out_CYw_Sply_Slide_A_F_Done : BOOL;
    Station_A_Data : ARRAY[0..8] OF sData;
    Cv_A_Data : ARRAY[0..8] OF sData;
    ST0_A_Sup_End : BOOL;  (* ST0 検査コンベア運転可 *)
    Out_CYS_Pos_01_Stopper_B_H_Auto : ARRAY[0..10] OF Bool;
    Out_CYS_Pos_02_Stopper_B_H_Auto : ARRAY[0..10] OF Bool;
    Out_CYS_Pos_03_Stopper_B_H_Auto : ARRAY[0..10] OF Bool;
    Out_CYS_Pos_04_Stopper_B_H_Auto : ARRAY[0..10] OF Bool;
    Out_CYS_Pos_05_Stopper_B_H_Auto : ARRAY[0..10] OF Bool;
    Out_CYS_Pos_06_Stopper_B_H_Auto : ARRAY[0..10] OF Bool;
    TimerQ_In_SenCY_Pos_01_Stopper_A_H : BOOL;
    TimerQ_In_SenCY_Pos_02_Stopper_A_H : BOOL;
    TimerQ_In_SenCY_Pos_03_Stopper_A_H : BOOL;
    TimerQ_In_SenCY_Pos_04_Stopper_A_H : BOOL;
    TimerQ_In_SenCY_Pos_05_Stopper_A_H : BOOL;
    TimerQ_In_SenCY_Pos_06_Stopper_A_H : BOOL;
    Out_Insp_Cv_A_Run_Auto : ARRAY[0..10] OF Bool;
    TimerQ_In_Sen_Work_A_Pos_01 : BOOL;
    TimerQ_In_Sen_Work_A_Pos_02 : BOOL;
    Pause : ARRAY[0..99] OF Bool;
    TimerQ_In_Sen_Work_A_Pos_03 : BOOL;
    TimerQ_In_Sen_Work_A_Pos_04 : BOOL;
    TimerQ_In_Sen_Work_A_Pos_05 : BOOL;
    TimerQ_In_Sen_Work_A_Pos_06 : BOOL;
    TimerQ_In_Sen_Work_A_Pos_07 : BOOL;
    Out_CYS_Pos_01_Stopper_A_H_Auto : ARRAY[0..10] OF Bool;
    Out_CYS_Pos_02_Stopper_A_H_Auto : ARRAY[0..10] OF Bool;
    Out_CYS_Pos_03_Stopper_A_H_Auto : ARRAY[0..10] OF Bool;
    Out_CYS_Pos_04_Stopper_A_H_Auto : ARRAY[0..10] OF Bool;
    Out_CYS_Pos_05_Stopper_A_H_Auto : ARRAY[0..10] OF Bool;
    Out_CYS_Pos_06_Stopper_A_H_Auto : ARRAY[0..10] OF Bool;
    Ins_A_Cv_M : ARRAY[0..99] OF Bool;
    Ins_A_Cv_Error : BOOL;  (* 検査コンベア ワーク不一致エラー *)
    TimerQ_In_Sen_Work_A_Pos_00 : BOOL;
    Out_CYS_Pos_01_Stopper_A_F_Auto : ARRAY[0..10] OF Bool;
    Out_CYS_Pos_02_Stopper_A_F_Auto : ARRAY[0..10] OF Bool;
    Out_CYS_Pos_03_Stopper_A_F_Auto : ARRAY[0..10] OF Bool;
    Out_CYS_Pos_04_Stopper_A_F_Auto : ARRAY[0..10] OF Bool;
    Out_CYS_Pos_05_Stopper_A_F_Auto : ARRAY[0..10] OF Bool;
    Out_CYS_Pos_06_Stopper_A_F_Auto : ARRAY[0..10] OF Bool;
    Ins_A_Next_Cycle : BOOL;  (* A(左側)検査コンベア 動作完了 *)
    ST0_A_Sup_Busy : BOOL;  (* ST0 稼働中 *)
    Ins_A_End : BOOL;  (* 検査完了 コンベア運転可能 *)
    Auto_A_Start : BOOL;
    Out_CYS_Pos_01_Stopper_A_H_Done : BOOL;
    FH_5552_10_A_Auto : BOOL;
    FH_A_ST1_Done : BOOL;
    ST1_A_Ca1_Busy : BOOL;  (* ST1 A検査中 *)
    ST1_A_Ca1_End : BOOL;  (* ST1 A 動作完了 *)
    ST2_A_Hgt_Busy : BOOL;  (* ST2 A 動作中 *)
    Out_CYw_HgtInsp_Clp_A_H_Auto : ARRAY[0..10] OF Bool;
    Out_CYw_HgtInsp_Clp_A_H_Done : BOOL;
    Out_CYw_HgtInsp_Lf_A_H_Auto : ARRAY[0..10] OF Bool;
    Out_CYw_HgtInsp_Lf_A_H_Done : BOOL;
    Out_CYS_Pos_02_Stopper_A_H_Done : BOOL;
    Out_CYw_HgtInsp_Clp_A_F_Auto : ARRAY[0..10] OF Bool;
    Out_CYw_HgtInsp_Clp_A_F_Done : BOOL;
    Out_CYw_HgtInsp_Lf_A_F_Auto : ARRAY[0..10] OF Bool;
    Out_CYw_HgtInsp_Lf_A_F_Done : BOOL;
    DLEP1_GT2_A_Auto : BOOL;
    Hgt_A_ComputedValueData : LREAL;
    Hight_LowerLimit : LREAL;  (* 高さ検査 下限値 *)
    Hight_UpperLimit : LREAL;  (* 高さ検査 上限値 *)
    ST2_A_Hgt_End : BOOL;  (* 高さ検査完了 *)
    ST3_A_Dis1_Busy : BOOL;  (* ST3 A 動作中 *)
    Out_CYw_NG1_Srt_A_H_Auto : ARRAY[0..10] OF Bool;
    Out_CYw_NG1_Srt_A_H_Done : BOOL;
    Out_CYw_Swv_01_Pick_A_H_Auto : ARRAY[0..10] OF Bool;
    Out_CYw_Swv_01_Pick_A_H_Done : BOOL;
    Out_CYw_NG1_Pick_A_H_Auto : ARRAY[0..10] OF Bool;
    Out_CYw_NG1_Pick_A_H_Done : BOOL;
    Out_CYw_NG1_Chk_A_H_Auto : ARRAY[0..10] OF Bool;
    Out_CYw_NG1_Chk_A_H_Done : BOOL;
END_VAR
VAR
    _e1 : R_TRIG;
    _p2 : BOOL;
    _e3 : R_TRIG;
    _e4 : R_TRIG;
    _p5 : BOOL;
    _e6 : R_TRIG;
    _e7 : R_TRIG;
    _p8 : BOOL;
    _p9 : BOOL;
    _p10 : BOOL;
    _p11 : BOOL;
    _p12 : BOOL;
    _p13 : BOOL;
    _p14 : BOOL;
    _p15 : BOOL;
    _e16 : R_TRIG;
    _p17 : BOOL;
    _p18 : BOOL;
    _p19 : BOOL;
    _p20 : BOOL;
    _p21 : BOOL;
    _p22 : BOOL;
    _p23 : BOOL;
    _p24 : BOOL;
    _p25 : BOOL;
    _p26 : BOOL;
    _p27 : BOOL;
    _p28 : BOOL;
    _e29 : R_TRIG;
    _p30 : BOOL;
    _p31 : BOOL;
    _p32 : BOOL;
    _p33 : BOOL;
    _p34 : BOOL;
    _p35 : BOOL;
    _p36 : BOOL;
    _p37 : BOOL;
    _p38 : BOOL;
    _p39 : BOOL;
    _p40 : BOOL;
    _p41 : BOOL;
    _p42 : BOOL;
END_VAR

(* Section Ins_A_Cv_左検査Cv: ladder, written here as Structured Text *)

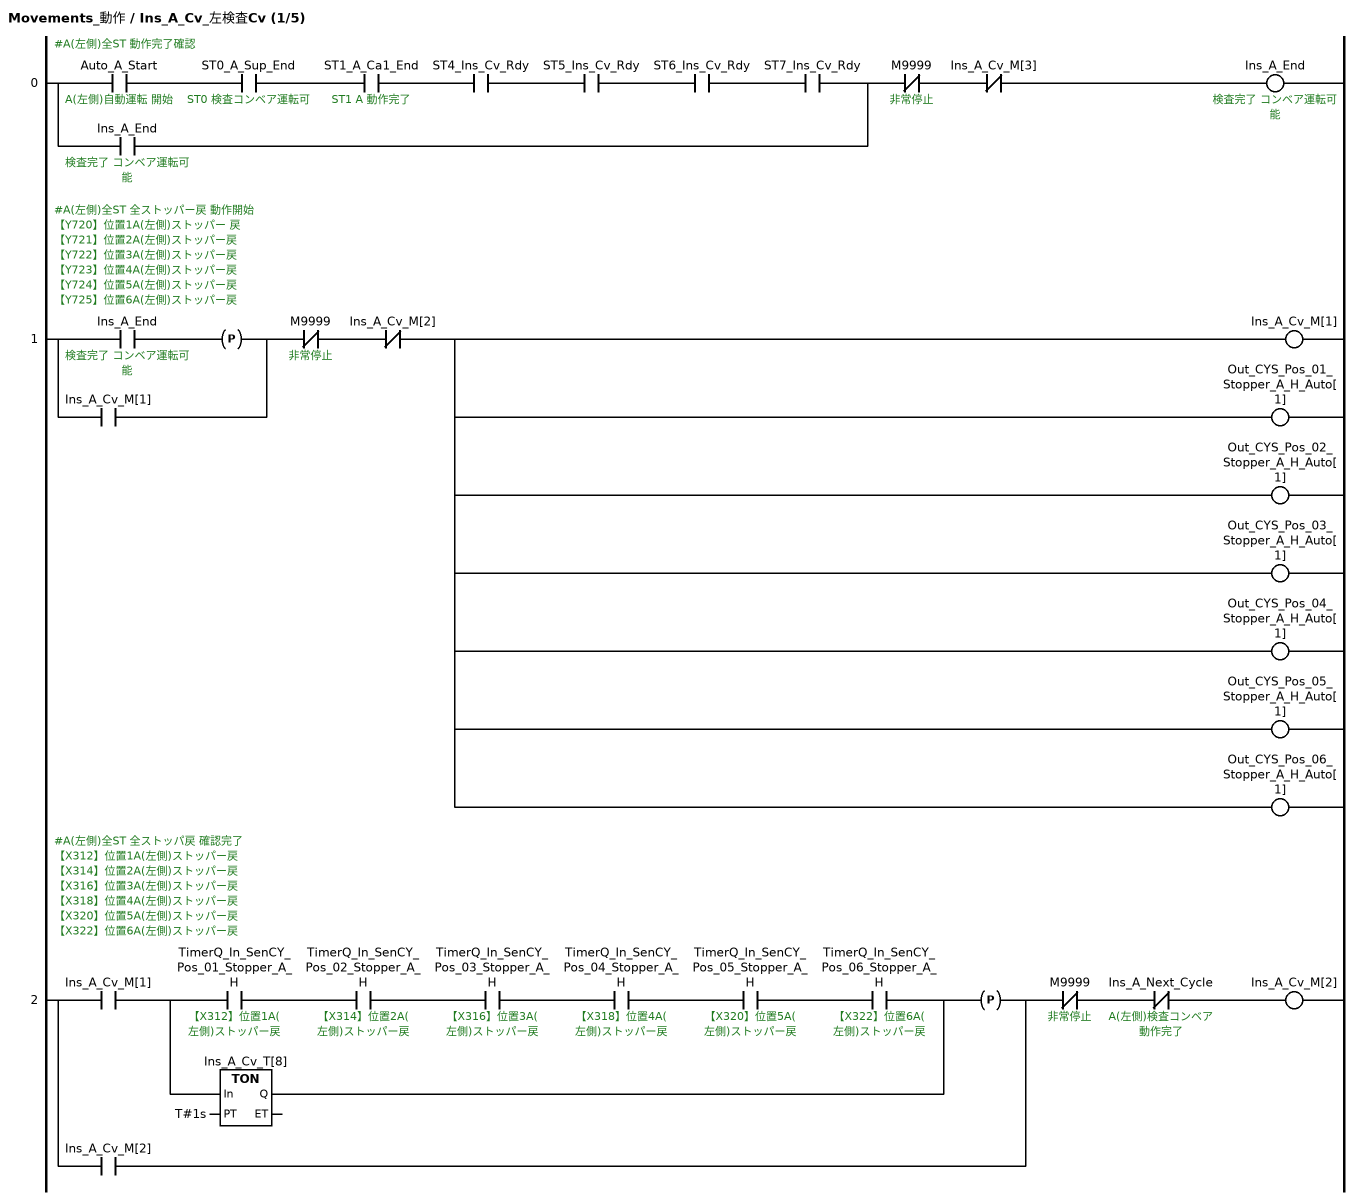
(* Rung 0: #A(左側)全ST 動作完了確認 *)
Ins_A_End := ((Auto_A_Start AND ST0_A_Sup_End AND ST1_A_Ca1_End AND ST4_Ins_Cv_Rdy AND ST5_Ins_Cv_Rdy AND ST6_Ins_Cv_Rdy AND ST7_Ins_Cv_Rdy) OR Ins_A_End) AND NOT M9999 AND NOT Ins_A_Cv_M[3];
(* Rung 1: #A(左側)全ST 全ストッパー戻 動作開始 / 【Y720】位置1A(左側)ストッパー 戻 / 【Y721】位置2A(左側)ストッパー戻 / 【Y722】位置3A(左側)ストッパー戻 / 【Y723】位置4A(左側)ストッパー戻 / 【Y724】位置5A(左側)ストッパー戻 / 【Y725】位置6A(左側)ストッパー戻 *)
_e1(CLK := Ins_A_End);
_p2 := (_e1.Q OR Ins_A_Cv_M[1]) AND NOT M9999 AND NOT Ins_A_Cv_M[2];
Ins_A_Cv_M[1] := _p2;
Out_CYS_Pos_01_Stopper_A_H_Auto[1] := _p2;
Out_CYS_Pos_02_Stopper_A_H_Auto[1] := _p2;
Out_CYS_Pos_03_Stopper_A_H_Auto[1] := _p2;
Out_CYS_Pos_04_Stopper_A_H_Auto[1] := _p2;
Out_CYS_Pos_05_Stopper_A_H_Auto[1] := _p2;
Out_CYS_Pos_06_Stopper_A_H_Auto[1] := _p2;
(* Rung 2: #A(左側)全ST 全ストッパ戻 確認完了 / 【X312】位置1A(左側)ストッパー戻 / 【X314】位置2A(左側)ストッパー戻 / 【X316】位置3A(左側)ストッパー戻 / 【X318】位置4A(左側)ストッパー戻 / 【X320】位置5A(左側)ストッパー戻 / 【X322】位置6A(左側)ストッパー戻 *)
Ins_A_Cv_T[8](In := Ins_A_Cv_M[1], PT := T#1s);
_e3(CLK := (Ins_A_Cv_M[1] AND TimerQ_In_SenCY_Pos_01_Stopper_A_H AND TimerQ_In_SenCY_Pos_02_Stopper_A_H AND TimerQ_In_SenCY_Pos_03_Stopper_A_H AND TimerQ_In_SenCY_Pos_04_Stopper_A_H AND TimerQ_In_SenCY_Pos_05_Stopper_A_H AND TimerQ_In_SenCY_Pos_06_Stopper_A_H) OR Ins_A_Cv_T[8].Q);
Ins_A_Cv_M[2] := (_e3.Q OR Ins_A_Cv_M[2]) AND NOT M9999 AND NOT Ins_A_Next_Cycle;

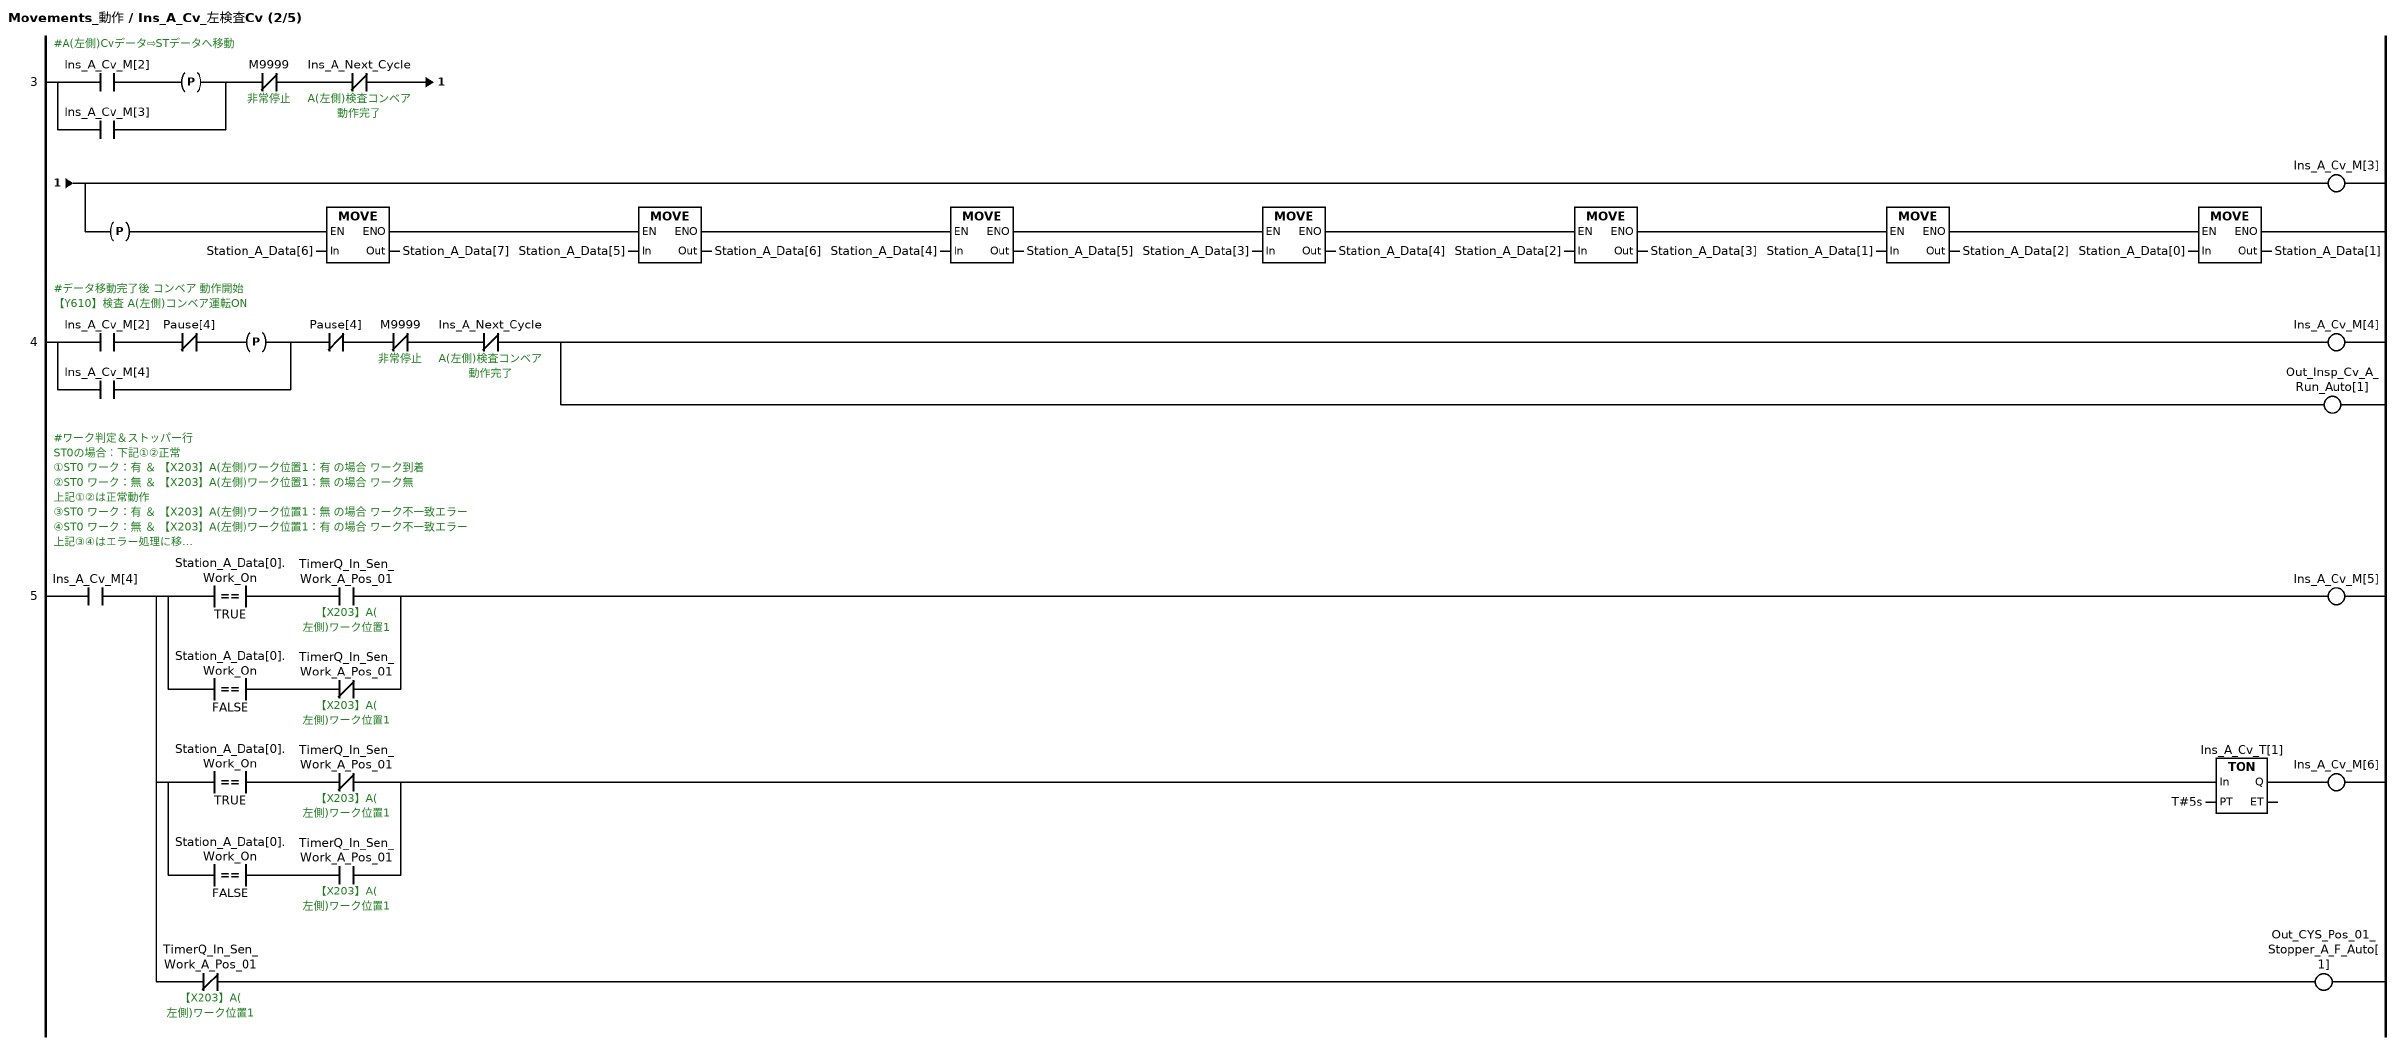
(* Rung 3: #A(左側)Cvデータ⇨STデータへ移動 *)
_e4(CLK := Ins_A_Cv_M[2]);
_p5 := (_e4.Q OR Ins_A_Cv_M[3]) AND NOT M9999 AND NOT Ins_A_Next_Cycle;
Ins_A_Cv_M[3] := _p5;
_e6(CLK := _p5);
IF _e6.Q THEN
    Station_A_Data[7] := Station_A_Data[6];
    Station_A_Data[6] := Station_A_Data[5];
    Station_A_Data[5] := Station_A_Data[4];
    Station_A_Data[4] := Station_A_Data[3];
    Station_A_Data[3] := Station_A_Data[2];
    Station_A_Data[2] := Station_A_Data[1];
    Station_A_Data[1] := Station_A_Data[0];
END_IF;
(* Rung 4: #データ移動完了後 コンベア 動作開始 / 【Y610】検査 A(左側)コンベア運転ON *)
_e7(CLK := Ins_A_Cv_M[2] AND NOT Pause[4]);
_p8 := (_e7.Q OR Ins_A_Cv_M[4]) AND NOT Pause[4] AND NOT M9999 AND NOT Ins_A_Next_Cycle;
Ins_A_Cv_M[4] := _p8;
Out_Insp_Cv_A_Run_Auto[1] := _p8;
(* Rung 5: #ワーク判定＆ストッパー行 / ST0の場合：下記①②正常 / ①ST0 ワーク：有 ＆ 【X203】A(左側)ワーク位置1：有 の場合 ワーク到着 / ②ST0 ワーク：無 ＆ 【X203】A(左側)ワーク位置1：無 の場合 ワーク無 / 上記①②は正常動作 / ③ST0 ワーク：有 ＆ 【X203】A(左側)ワーク位置1：無 の場合 ワーク不一致エラー / ④ST0 ワーク：無 ＆ 【X203】A(左側)ワーク位置1：有 の場合 ワーク不一致エラー / 上記③④はエラー処理に移動 / ⑤【X203】A(左側)ワーク位置1：無 の場合 / 【Y720】位置1A(左側)ストッパー 行 *)
_p9 := Ins_A_Cv_M[4];
Ins_A_Cv_M[5] := Ins_A_Cv_M[4] AND (((Station_A_Data[0].Work_On = TRUE) AND TimerQ_In_Sen_Work_A_Pos_01) OR ((Station_A_Data[0].Work_On = FALSE) AND NOT TimerQ_In_Sen_Work_A_Pos_01));
Ins_A_Cv_T[1](In := _p9 AND (((Station_A_Data[0].Work_On = TRUE) AND NOT TimerQ_In_Sen_Work_A_Pos_01) OR ((Station_A_Data[0].Work_On = FALSE) AND TimerQ_In_Sen_Work_A_Pos_01)), PT := T#5s);
Ins_A_Cv_M[6] := Ins_A_Cv_T[1].Q;
Out_CYS_Pos_01_Stopper_A_F_Auto[1] := _p9 AND NOT TimerQ_In_Sen_Work_A_Pos_01;

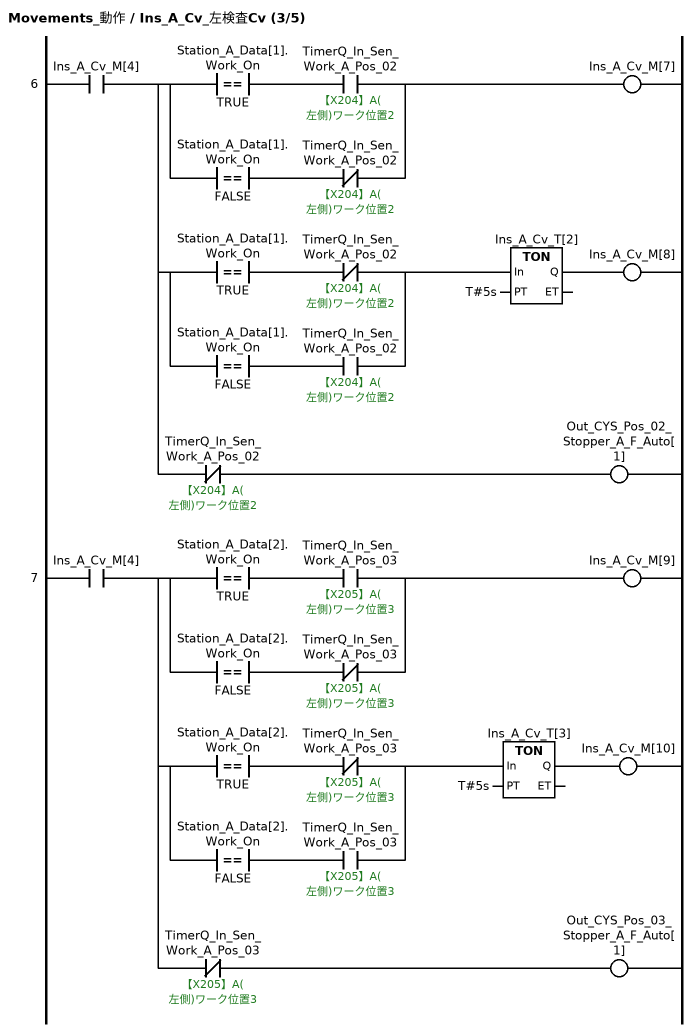
(* Rung 6 *)
_p10 := Ins_A_Cv_M[4];
Ins_A_Cv_M[7] := Ins_A_Cv_M[4] AND (((Station_A_Data[1].Work_On = TRUE) AND TimerQ_In_Sen_Work_A_Pos_02) OR ((Station_A_Data[1].Work_On = FALSE) AND NOT TimerQ_In_Sen_Work_A_Pos_02));
Ins_A_Cv_T[2](In := _p10 AND (((Station_A_Data[1].Work_On = TRUE) AND NOT TimerQ_In_Sen_Work_A_Pos_02) OR ((Station_A_Data[1].Work_On = FALSE) AND TimerQ_In_Sen_Work_A_Pos_02)), PT := T#5s);
Ins_A_Cv_M[8] := Ins_A_Cv_T[2].Q;
Out_CYS_Pos_02_Stopper_A_F_Auto[1] := _p10 AND NOT TimerQ_In_Sen_Work_A_Pos_02;
(* Rung 7 *)
_p11 := Ins_A_Cv_M[4];
Ins_A_Cv_M[9] := Ins_A_Cv_M[4] AND (((Station_A_Data[2].Work_On = TRUE) AND TimerQ_In_Sen_Work_A_Pos_03) OR ((Station_A_Data[2].Work_On = FALSE) AND NOT TimerQ_In_Sen_Work_A_Pos_03));
Ins_A_Cv_T[3](In := _p11 AND (((Station_A_Data[2].Work_On = TRUE) AND NOT TimerQ_In_Sen_Work_A_Pos_03) OR ((Station_A_Data[2].Work_On = FALSE) AND TimerQ_In_Sen_Work_A_Pos_03)), PT := T#5s);
Ins_A_Cv_M[10] := Ins_A_Cv_T[3].Q;
Out_CYS_Pos_03_Stopper_A_F_Auto[1] := _p11 AND NOT TimerQ_In_Sen_Work_A_Pos_03;

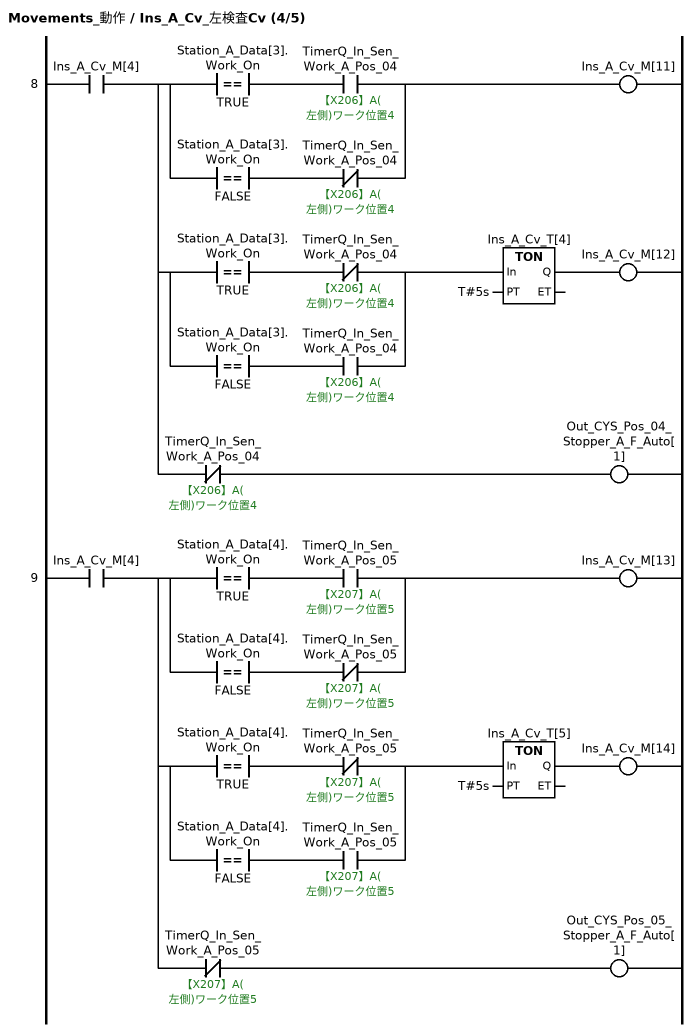
(* Rung 8 *)
_p12 := Ins_A_Cv_M[4];
Ins_A_Cv_M[11] := Ins_A_Cv_M[4] AND (((Station_A_Data[3].Work_On = TRUE) AND TimerQ_In_Sen_Work_A_Pos_04) OR ((Station_A_Data[3].Work_On = FALSE) AND NOT TimerQ_In_Sen_Work_A_Pos_04));
Ins_A_Cv_T[4](In := _p12 AND (((Station_A_Data[3].Work_On = TRUE) AND NOT TimerQ_In_Sen_Work_A_Pos_04) OR ((Station_A_Data[3].Work_On = FALSE) AND TimerQ_In_Sen_Work_A_Pos_04)), PT := T#5s);
Ins_A_Cv_M[12] := Ins_A_Cv_T[4].Q;
Out_CYS_Pos_04_Stopper_A_F_Auto[1] := _p12 AND NOT TimerQ_In_Sen_Work_A_Pos_04;
(* Rung 9 *)
_p13 := Ins_A_Cv_M[4];
Ins_A_Cv_M[13] := Ins_A_Cv_M[4] AND (((Station_A_Data[4].Work_On = TRUE) AND TimerQ_In_Sen_Work_A_Pos_05) OR ((Station_A_Data[4].Work_On = FALSE) AND NOT TimerQ_In_Sen_Work_A_Pos_05));
Ins_A_Cv_T[5](In := _p13 AND (((Station_A_Data[4].Work_On = TRUE) AND NOT TimerQ_In_Sen_Work_A_Pos_05) OR ((Station_A_Data[4].Work_On = FALSE) AND TimerQ_In_Sen_Work_A_Pos_05)), PT := T#5s);
Ins_A_Cv_M[14] := Ins_A_Cv_T[5].Q;
Out_CYS_Pos_05_Stopper_A_F_Auto[1] := _p13 AND NOT TimerQ_In_Sen_Work_A_Pos_05;

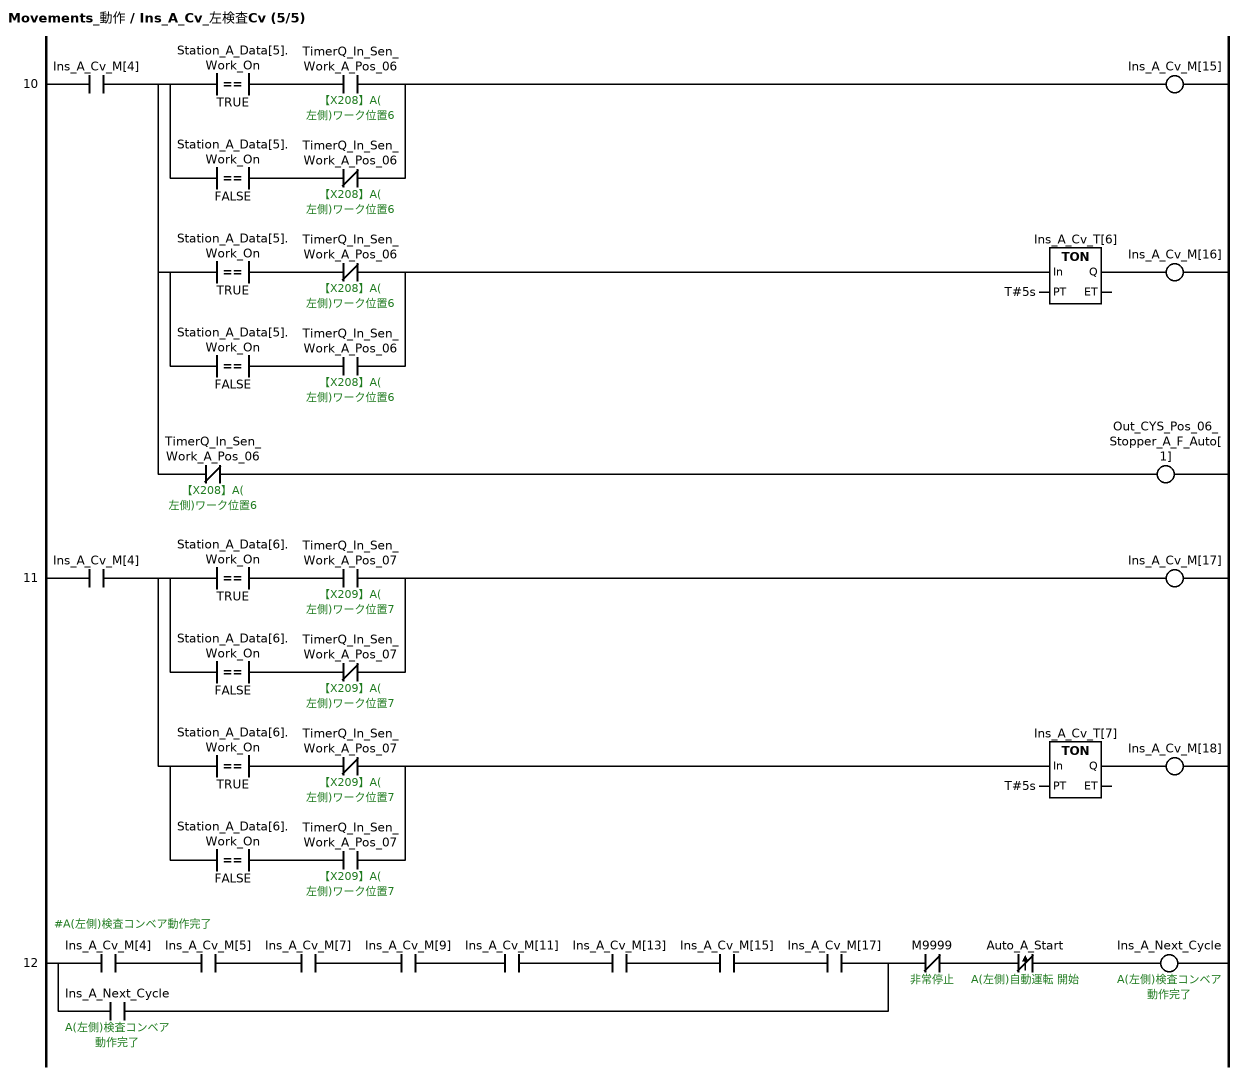
(* Rung 10 *)
_p14 := Ins_A_Cv_M[4];
Ins_A_Cv_M[15] := Ins_A_Cv_M[4] AND (((Station_A_Data[5].Work_On = TRUE) AND TimerQ_In_Sen_Work_A_Pos_06) OR ((Station_A_Data[5].Work_On = FALSE) AND NOT TimerQ_In_Sen_Work_A_Pos_06));
Ins_A_Cv_T[6](In := _p14 AND (((Station_A_Data[5].Work_On = TRUE) AND NOT TimerQ_In_Sen_Work_A_Pos_06) OR ((Station_A_Data[5].Work_On = FALSE) AND TimerQ_In_Sen_Work_A_Pos_06)), PT := T#5s);
Ins_A_Cv_M[16] := Ins_A_Cv_T[6].Q;
Out_CYS_Pos_06_Stopper_A_F_Auto[1] := _p14 AND NOT TimerQ_In_Sen_Work_A_Pos_06;
(* Rung 11 *)
_p15 := Ins_A_Cv_M[4];
Ins_A_Cv_M[17] := Ins_A_Cv_M[4] AND (((Station_A_Data[6].Work_On = TRUE) AND TimerQ_In_Sen_Work_A_Pos_07) OR ((Station_A_Data[6].Work_On = FALSE) AND NOT TimerQ_In_Sen_Work_A_Pos_07));
Ins_A_Cv_T[7](In := _p15 AND (((Station_A_Data[6].Work_On = TRUE) AND NOT TimerQ_In_Sen_Work_A_Pos_07) OR ((Station_A_Data[6].Work_On = FALSE) AND TimerQ_In_Sen_Work_A_Pos_07)), PT := T#5s);
Ins_A_Cv_M[18] := Ins_A_Cv_T[7].Q;
(* Rung 12: #A(左側)検査コンベア動作完了 *)
_e16(CLK := Auto_A_Start);
Ins_A_Next_Cycle := ((Ins_A_Cv_M[4] AND Ins_A_Cv_M[5] AND Ins_A_Cv_M[7] AND Ins_A_Cv_M[9] AND Ins_A_Cv_M[11] AND Ins_A_Cv_M[13] AND Ins_A_Cv_M[15] AND Ins_A_Cv_M[17]) OR Ins_A_Next_Cycle) AND NOT M9999 AND NOT _e16.Q;

(* Section ST0_A_Sup_左供給: ladder, written here as Structured Text *)

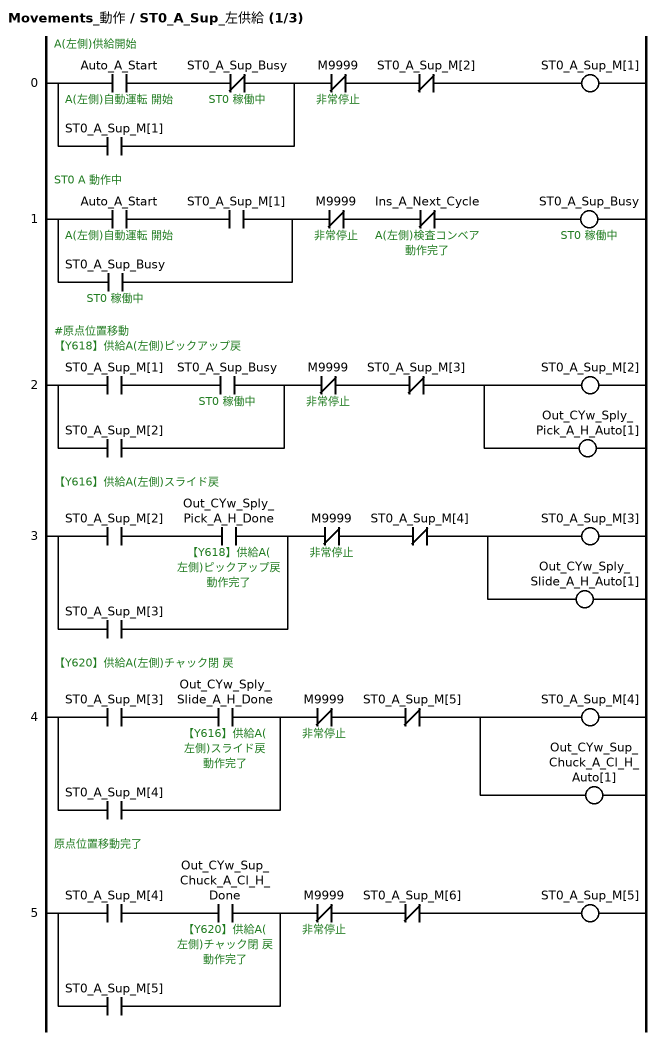
(* Rung 0: A(左側)供給開始 *)
ST0_A_Sup_M[1] := ((Auto_A_Start AND NOT ST0_A_Sup_Busy) OR ST0_A_Sup_M[1]) AND NOT M9999 AND NOT ST0_A_Sup_M[2];
(* Rung 1: ST0 A 動作中 *)
ST0_A_Sup_Busy := ((Auto_A_Start AND ST0_A_Sup_M[1]) OR ST0_A_Sup_Busy) AND NOT M9999 AND NOT Ins_A_Next_Cycle;
(* Rung 2: #原点位置移動 / 【Y618】供給A(左側)ピックアップ戻 *)
_p17 := ((ST0_A_Sup_M[1] AND ST0_A_Sup_Busy) OR ST0_A_Sup_M[2]) AND NOT M9999 AND NOT ST0_A_Sup_M[3];
ST0_A_Sup_M[2] := _p17;
Out_CYw_Sply_Pick_A_H_Auto[1] := _p17;
(* Rung 3: 【Y616】供給A(左側)スライド戻 *)
_p18 := ((ST0_A_Sup_M[2] AND Out_CYw_Sply_Pick_A_H_Done) OR ST0_A_Sup_M[3]) AND NOT M9999 AND NOT ST0_A_Sup_M[4];
ST0_A_Sup_M[3] := _p18;
Out_CYw_Sply_Slide_A_H_Auto[1] := _p18;
(* Rung 4: 【Y620】供給A(左側)チャック閉 戻 *)
_p19 := ((ST0_A_Sup_M[3] AND Out_CYw_Sply_Slide_A_H_Done) OR ST0_A_Sup_M[4]) AND NOT M9999 AND NOT ST0_A_Sup_M[5];
ST0_A_Sup_M[4] := _p19;
Out_CYw_Sup_Chuck_A_Cl_H_Auto[1] := _p19;
(* Rung 5: 原点位置移動完了 *)
ST0_A_Sup_M[5] := ((ST0_A_Sup_M[4] AND Out_CYw_Sup_Chuck_A_Cl_H_Done) OR ST0_A_Sup_M[5]) AND NOT M9999 AND NOT ST0_A_Sup_M[6];

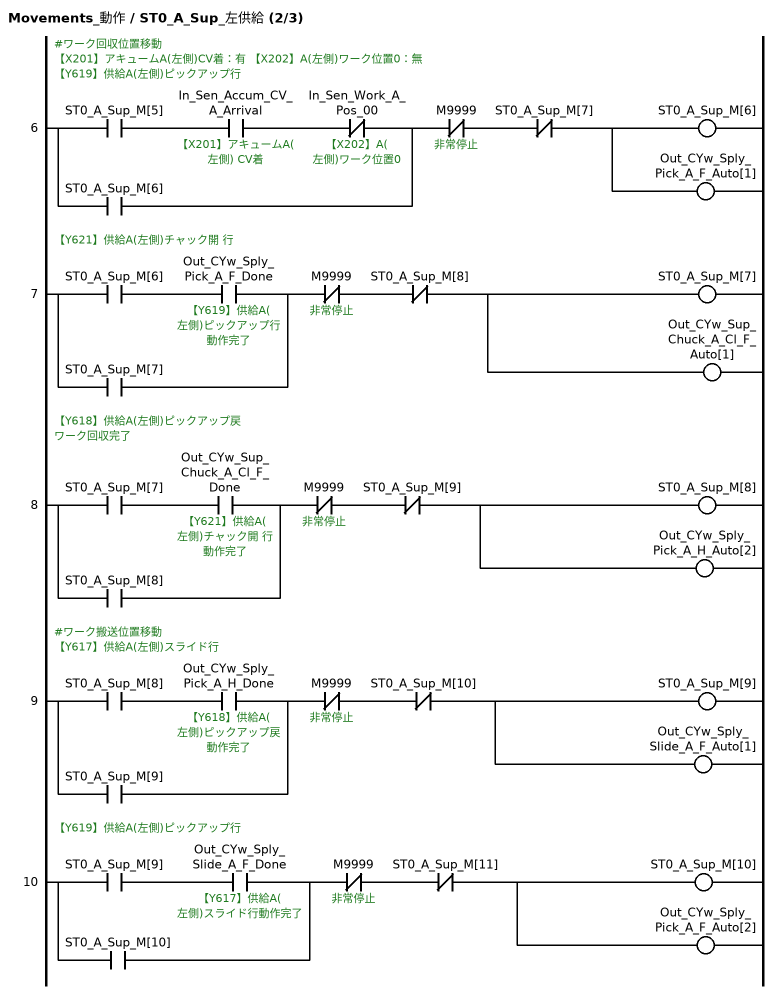
(* Rung 6: #ワーク回収位置移動 / 【X201】アキュームA(左側)CV着：有 【X202】A(左側)ワーク位置0：無 / 【Y619】供給A(左側)ピックアップ行 *)
_p20 := ((ST0_A_Sup_M[5] AND In_Sen_Accum_CV_A_Arrival AND NOT In_Sen_Work_A_Pos_00) OR ST0_A_Sup_M[6]) AND NOT M9999 AND NOT ST0_A_Sup_M[7];
ST0_A_Sup_M[6] := _p20;
Out_CYw_Sply_Pick_A_F_Auto[1] := _p20;
(* Rung 7: 【Y621】供給A(左側)チャック開 行 *)
_p21 := ((ST0_A_Sup_M[6] AND Out_CYw_Sply_Pick_A_F_Done) OR ST0_A_Sup_M[7]) AND NOT M9999 AND NOT ST0_A_Sup_M[8];
ST0_A_Sup_M[7] := _p21;
Out_CYw_Sup_Chuck_A_Cl_F_Auto[1] := _p21;
(* Rung 8: 【Y618】供給A(左側)ピックアップ戻 / ワーク回収完了 *)
_p22 := ((ST0_A_Sup_M[7] AND Out_CYw_Sup_Chuck_A_Cl_F_Done) OR ST0_A_Sup_M[8]) AND NOT M9999 AND NOT ST0_A_Sup_M[9];
ST0_A_Sup_M[8] := _p22;
Out_CYw_Sply_Pick_A_H_Auto[2] := _p22;
(* Rung 9: #ワーク搬送位置移動 / 【Y617】供給A(左側)スライド行 *)
_p23 := ((ST0_A_Sup_M[8] AND Out_CYw_Sply_Pick_A_H_Done) OR ST0_A_Sup_M[9]) AND NOT M9999 AND NOT ST0_A_Sup_M[10];
ST0_A_Sup_M[9] := _p23;
Out_CYw_Sply_Slide_A_F_Auto[1] := _p23;
(* Rung 10: 【Y619】供給A(左側)ピックアップ行 *)
_p24 := ((ST0_A_Sup_M[9] AND Out_CYw_Sply_Slide_A_F_Done) OR ST0_A_Sup_M[10]) AND NOT M9999 AND NOT ST0_A_Sup_M[11];
ST0_A_Sup_M[10] := _p24;
Out_CYw_Sply_Pick_A_F_Auto[2] := _p24;

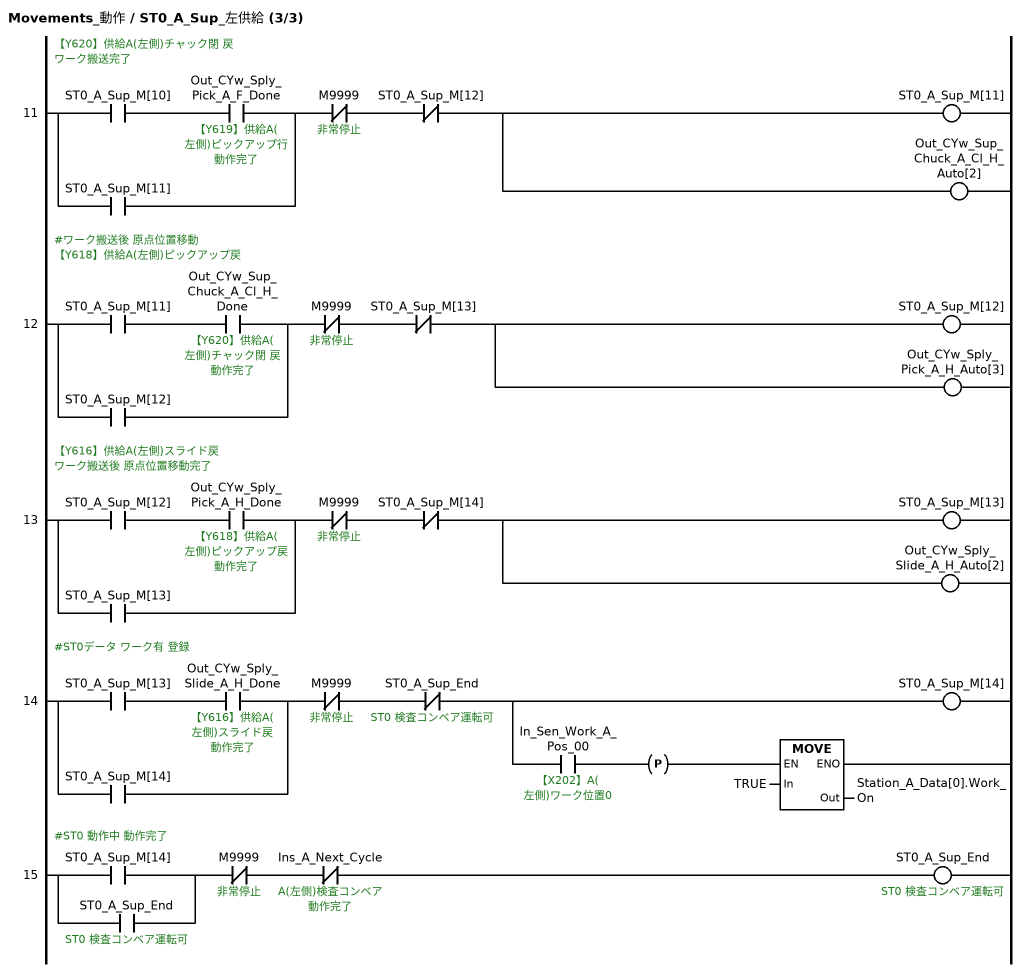
(* Rung 11: 【Y620】供給A(左側)チャック閉 戻 / ワーク搬送完了 *)
_p25 := ((ST0_A_Sup_M[10] AND Out_CYw_Sply_Pick_A_F_Done) OR ST0_A_Sup_M[11]) AND NOT M9999 AND NOT ST0_A_Sup_M[12];
ST0_A_Sup_M[11] := _p25;
Out_CYw_Sup_Chuck_A_Cl_H_Auto[2] := _p25;
(* Rung 12: #ワーク搬送後 原点位置移動 / 【Y618】供給A(左側)ピックアップ戻 *)
_p26 := ((ST0_A_Sup_M[11] AND Out_CYw_Sup_Chuck_A_Cl_H_Done) OR ST0_A_Sup_M[12]) AND NOT M9999 AND NOT ST0_A_Sup_M[13];
ST0_A_Sup_M[12] := _p26;
Out_CYw_Sply_Pick_A_H_Auto[3] := _p26;
(* Rung 13: 【Y616】供給A(左側)スライド戻 / ワーク搬送後 原点位置移動完了 *)
_p27 := ((ST0_A_Sup_M[12] AND Out_CYw_Sply_Pick_A_H_Done) OR ST0_A_Sup_M[13]) AND NOT M9999 AND NOT ST0_A_Sup_M[14];
ST0_A_Sup_M[13] := _p27;
Out_CYw_Sply_Slide_A_H_Auto[2] := _p27;
(* Rung 14: #ST0データ ワーク有 登録 *)
_p28 := ((ST0_A_Sup_M[13] AND Out_CYw_Sply_Slide_A_H_Done) OR ST0_A_Sup_M[14]) AND NOT M9999 AND NOT ST0_A_Sup_End;
ST0_A_Sup_M[14] := _p28;
_e29(CLK := _p28 AND In_Sen_Work_A_Pos_00);
IF _e29.Q THEN Station_A_Data[0].Work_On := TRUE; END_IF;
(* Rung 15: #ST0 動作中 動作完了 *)
ST0_A_Sup_End := (ST0_A_Sup_M[14] OR ST0_A_Sup_End) AND NOT M9999 AND NOT Ins_A_Next_Cycle;

(* Section ST1_A_Ca1_左Ca1検査: ladder, written here as Structured Text *)

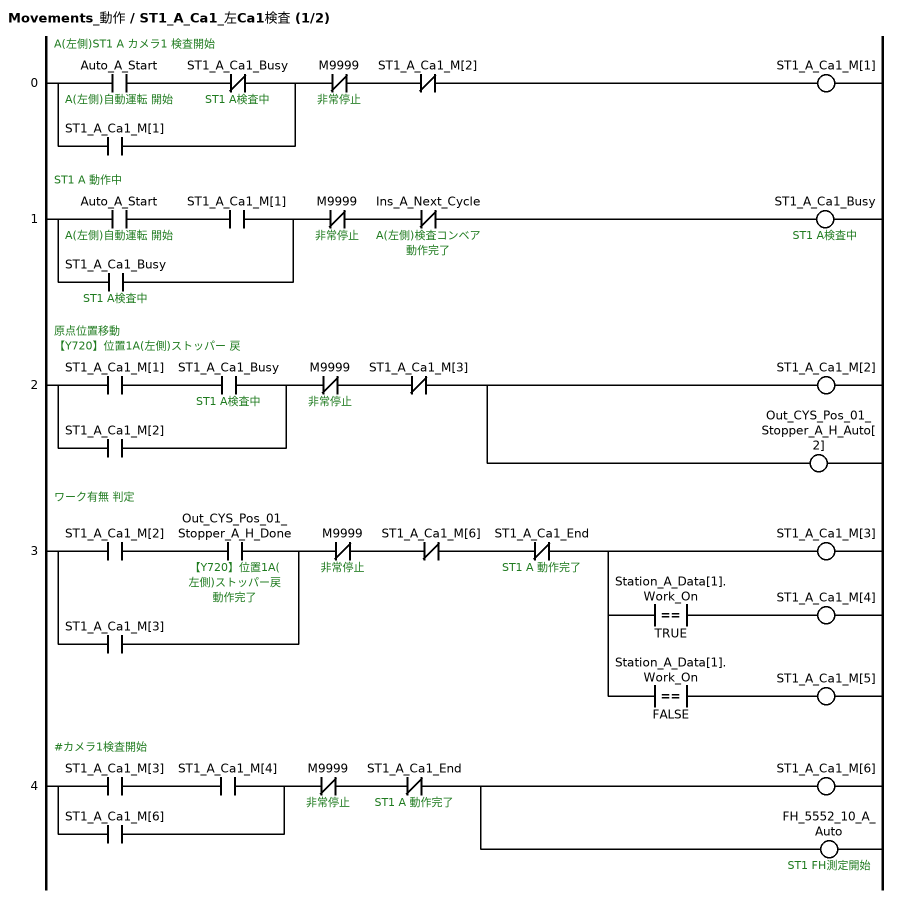
(* Rung 0: A(左側)ST1 A カメラ1 検査開始 *)
ST1_A_Ca1_M[1] := ((Auto_A_Start AND NOT ST1_A_Ca1_Busy) OR ST1_A_Ca1_M[1]) AND NOT M9999 AND NOT ST1_A_Ca1_M[2];
(* Rung 1: ST1 A 動作中 *)
ST1_A_Ca1_Busy := ((Auto_A_Start AND ST1_A_Ca1_M[1]) OR ST1_A_Ca1_Busy) AND NOT M9999 AND NOT Ins_A_Next_Cycle;
(* Rung 2: 原点位置移動 / 【Y720】位置1A(左側)ストッパー 戻 *)
_p30 := ((ST1_A_Ca1_M[1] AND ST1_A_Ca1_Busy) OR ST1_A_Ca1_M[2]) AND NOT M9999 AND NOT ST1_A_Ca1_M[3];
ST1_A_Ca1_M[2] := _p30;
Out_CYS_Pos_01_Stopper_A_H_Auto[2] := _p30;
(* Rung 3: ワーク有無 判定 *)
_p31 := ((ST1_A_Ca1_M[2] AND Out_CYS_Pos_01_Stopper_A_H_Done) OR ST1_A_Ca1_M[3]) AND NOT M9999 AND NOT ST1_A_Ca1_M[6] AND NOT ST1_A_Ca1_End;
ST1_A_Ca1_M[3] := _p31;
ST1_A_Ca1_M[4] := _p31 AND (Station_A_Data[1].Work_On = TRUE);
ST1_A_Ca1_M[5] := _p31 AND (Station_A_Data[1].Work_On = FALSE);
(* Rung 4: #カメラ1検査開始 *)
_p32 := ((ST1_A_Ca1_M[3] AND ST1_A_Ca1_M[4]) OR ST1_A_Ca1_M[6]) AND NOT M9999 AND NOT ST1_A_Ca1_End;
ST1_A_Ca1_M[6] := _p32;
FH_5552_10_A_Auto := _p32;

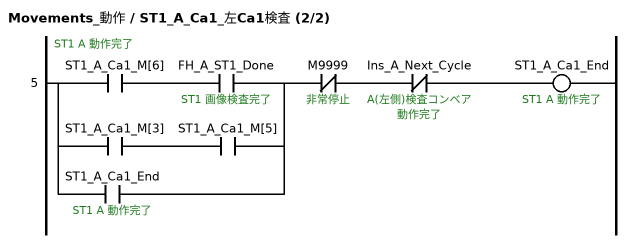
(* Rung 5: ST1 A 動作完了 *)
ST1_A_Ca1_End := ((ST1_A_Ca1_M[6] AND FH_A_ST1_Done) OR (ST1_A_Ca1_M[3] AND ST1_A_Ca1_M[5]) OR ST1_A_Ca1_End) AND NOT M9999 AND NOT Ins_A_Next_Cycle;

(* Section ST2_A_Hgt_左高さ検査: ladder, written here as Structured Text *)

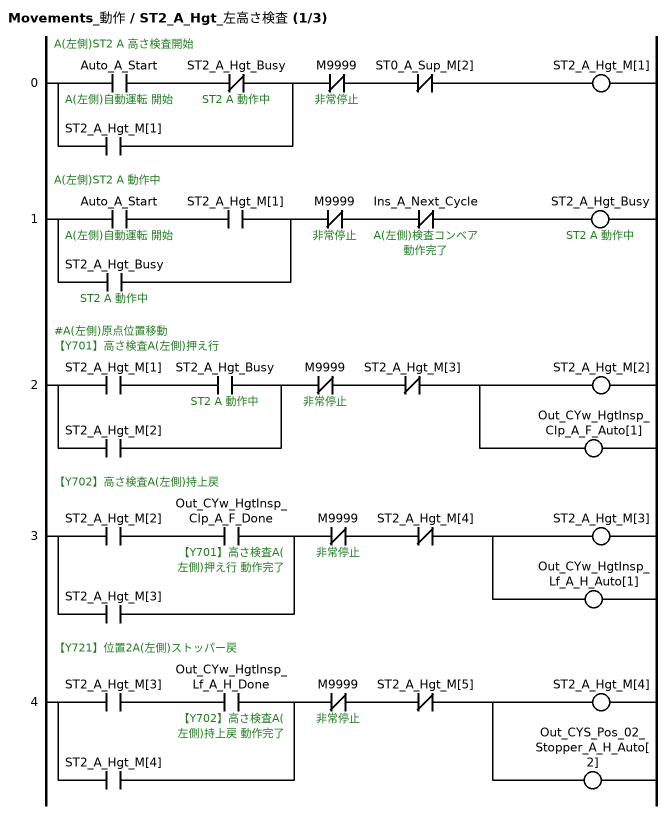
(* Rung 0: A(左側)ST2 A 高さ検査開始 *)
ST2_A_Hgt_M[1] := ((Auto_A_Start AND NOT ST2_A_Hgt_Busy) OR ST2_A_Hgt_M[1]) AND NOT M9999 AND NOT ST0_A_Sup_M[2];
(* Rung 1: A(左側)ST2 A 動作中 *)
ST2_A_Hgt_Busy := ((Auto_A_Start AND ST2_A_Hgt_M[1]) OR ST2_A_Hgt_Busy) AND NOT M9999 AND NOT Ins_A_Next_Cycle;
(* Rung 2: #A(左側)原点位置移動 / 【Y701】高さ検査A(左側)押え行 *)
_p33 := ((ST2_A_Hgt_M[1] AND ST2_A_Hgt_Busy) OR ST2_A_Hgt_M[2]) AND NOT M9999 AND NOT ST2_A_Hgt_M[3];
ST2_A_Hgt_M[2] := _p33;
Out_CYw_HgtInsp_Clp_A_F_Auto[1] := _p33;
(* Rung 3: 【Y702】高さ検査A(左側)持上戻 *)
_p34 := ((ST2_A_Hgt_M[2] AND Out_CYw_HgtInsp_Clp_A_F_Done) OR ST2_A_Hgt_M[3]) AND NOT M9999 AND NOT ST2_A_Hgt_M[4];
ST2_A_Hgt_M[3] := _p34;
Out_CYw_HgtInsp_Lf_A_H_Auto[1] := _p34;
(* Rung 4: 【Y721】位置2A(左側)ストッパー戻 *)
_p35 := ((ST2_A_Hgt_M[3] AND Out_CYw_HgtInsp_Lf_A_H_Done) OR ST2_A_Hgt_M[4]) AND NOT M9999 AND NOT ST2_A_Hgt_M[5];
ST2_A_Hgt_M[4] := _p35;
Out_CYS_Pos_02_Stopper_A_H_Auto[2] := _p35;

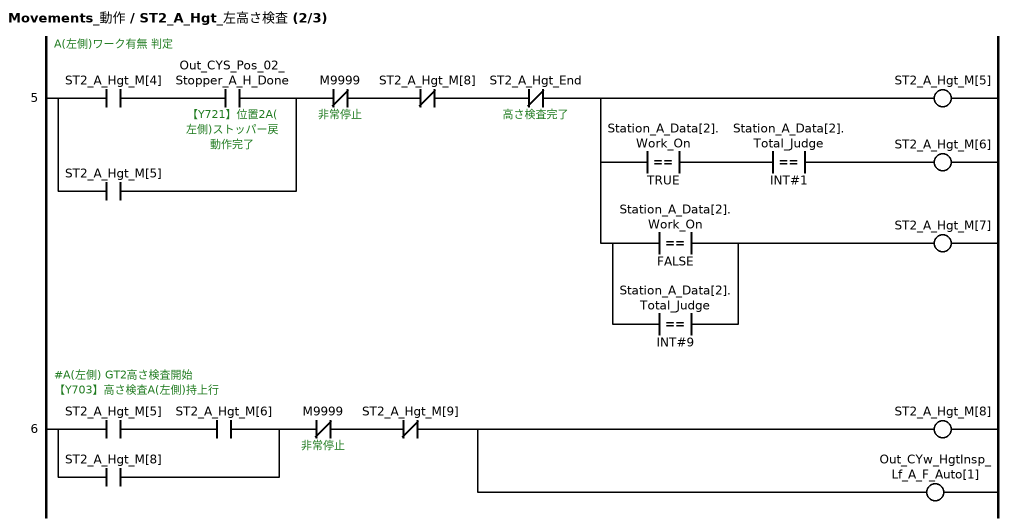
(* Rung 5: A(左側)ワーク有無 判定 *)
_p36 := ((ST2_A_Hgt_M[4] AND Out_CYS_Pos_02_Stopper_A_H_Done) OR ST2_A_Hgt_M[5]) AND NOT M9999 AND NOT ST2_A_Hgt_M[8] AND NOT ST2_A_Hgt_End;
ST2_A_Hgt_M[5] := _p36;
ST2_A_Hgt_M[6] := _p36 AND (Station_A_Data[2].Work_On = TRUE) AND (Station_A_Data[2].Total_Judge = INT#1);
ST2_A_Hgt_M[7] := _p36 AND ((Station_A_Data[2].Work_On = FALSE) OR (Station_A_Data[2].Total_Judge = INT#9));
(* Rung 6: #A(左側) GT2高さ検査開始 / 【Y703】高さ検査A(左側)持上行 *)
_p37 := ((ST2_A_Hgt_M[5] AND ST2_A_Hgt_M[6]) OR ST2_A_Hgt_M[8]) AND NOT M9999 AND NOT ST2_A_Hgt_M[9];
ST2_A_Hgt_M[8] := _p37;
Out_CYw_HgtInsp_Lf_A_F_Auto[1] := _p37;

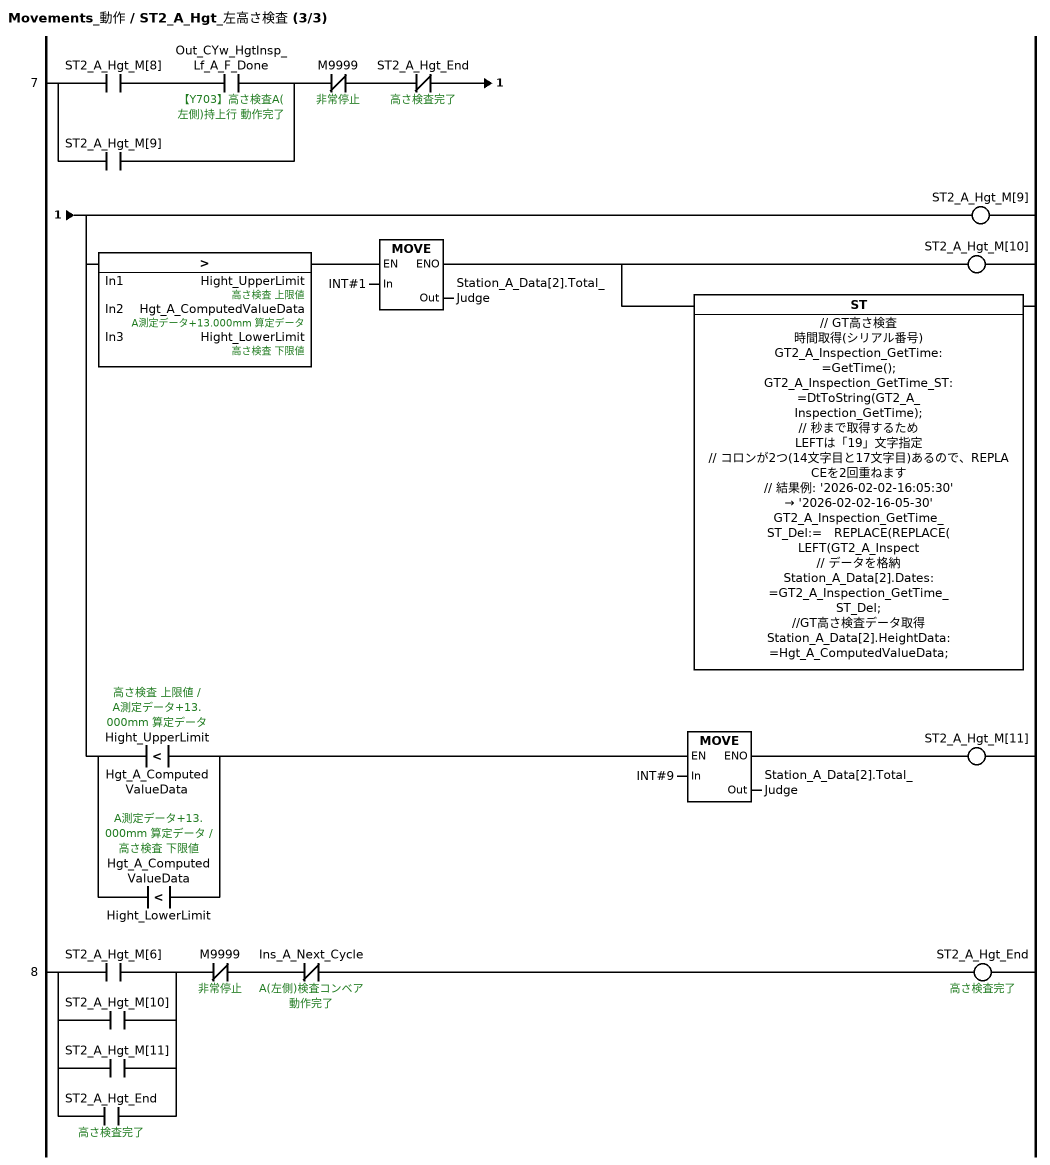
(* Rung 7 *)
_p38 := ((ST2_A_Hgt_M[8] AND Out_CYw_HgtInsp_Lf_A_F_Done) OR ST2_A_Hgt_M[9]) AND NOT M9999 AND NOT ST2_A_Hgt_End;
ST2_A_Hgt_M[9] := _p38;
IF _p38 AND GT(Hight_UpperLimit, Hgt_A_ComputedValueData, Hight_LowerLimit) THEN
    Station_A_Data[2].Total_Judge := INT#1;
END_IF;
_p39 := _p38 AND GT(Hight_UpperLimit, Hgt_A_ComputedValueData, Hight_LowerLimit);
ST2_A_Hgt_M[10] := _p39;
IF _p39 THEN
    // GT高さ検査 時間取得(シリアル番号)
    GT2_A_Inspection_GetTime:=GetTime();
    GT2_A_Inspection_GetTime_ST:=DtToString(GT2_A_Inspection_GetTime);
    // 秒まで取得するため LEFTは「19」文字指定
    // コロンが2つ(14文字目と17文字目)あるので、REPLACEを2回重ねます
    // 結果例: '2026-02-02-16:05:30' → '2026-02-02-16-05-30'
    GT2_A_Inspection_GetTime_ST_Del:=   REPLACE(REPLACE(LEFT(GT2_A_Inspection_GetTime_ST, UINT#19), STRING#'-', UINT#1, UINT#17), STRING#'-', UINT#1, UINT#14);
    // データを格納
    Station_A_Data[2].Dates:=GT2_A_Inspection_GetTime_ST_Del;
    //GT高さ検査データ取得
    Station_A_Data[2].HeightData:=Hgt_A_ComputedValueData;
END_IF;
IF _p38 AND ((Hight_UpperLimit < Hgt_A_ComputedValueData) OR (Hgt_A_ComputedValueData < Hight_LowerLimit)) THEN
    Station_A_Data[2].Total_Judge := INT#9;
END_IF;
ST2_A_Hgt_M[11] := _p38 AND ((Hight_UpperLimit < Hgt_A_ComputedValueData) OR (Hgt_A_ComputedValueData < Hight_LowerLimit));
(* Rung 8 *)
ST2_A_Hgt_End := (ST2_A_Hgt_M[6] OR ST2_A_Hgt_M[10] OR ST2_A_Hgt_M[11] OR ST2_A_Hgt_End) AND NOT M9999 AND NOT Ins_A_Next_Cycle;

(* Section ST3_A_Dis1_左NG1排出: ladder, written here as Structured Text *)

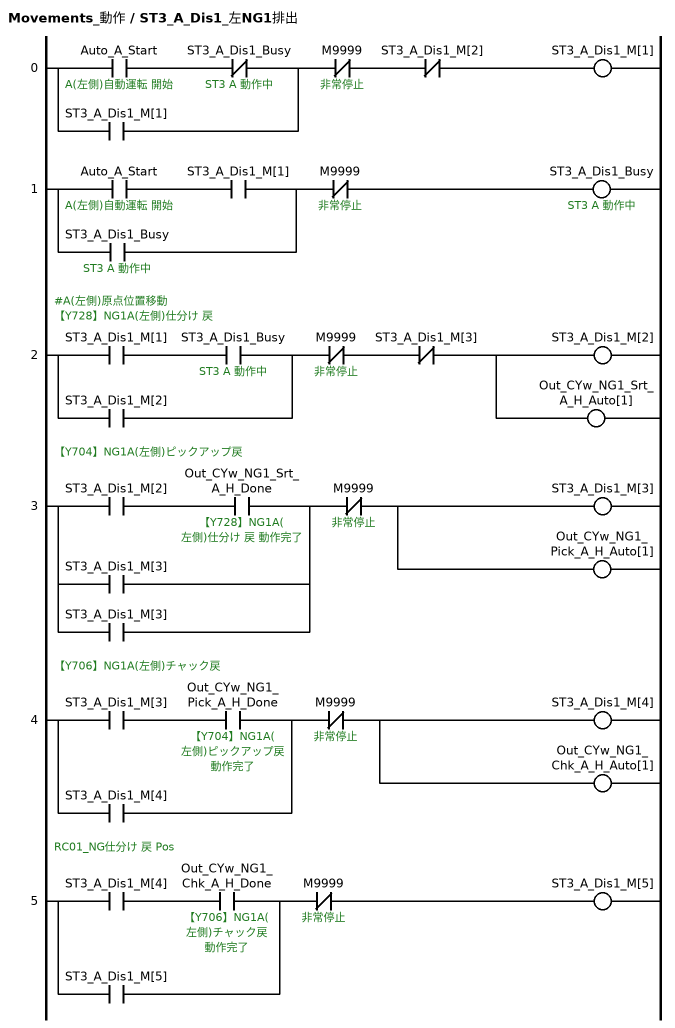
(* Rung 0 *)
ST3_A_Dis1_M[1] := ((Auto_A_Start AND NOT ST3_A_Dis1_Busy) OR ST3_A_Dis1_M[1]) AND NOT M9999 AND NOT ST3_A_Dis1_M[2];
(* Rung 1 *)
ST3_A_Dis1_Busy := ((Auto_A_Start AND ST3_A_Dis1_M[1]) OR ST3_A_Dis1_Busy) AND NOT M9999;
(* Rung 2: #A(左側)原点位置移動 / 【Y728】NG1A(左側)仕分け 戻 *)
_p40 := ((ST3_A_Dis1_M[1] AND ST3_A_Dis1_Busy) OR ST3_A_Dis1_M[2]) AND NOT M9999 AND NOT ST3_A_Dis1_M[3];
ST3_A_Dis1_M[2] := _p40;
Out_CYw_NG1_Srt_A_H_Auto[1] := _p40;
(* Rung 3: 【Y704】NG1A(左側)ピックアップ戻 *)
_p41 := ((ST3_A_Dis1_M[2] AND Out_CYw_NG1_Srt_A_H_Done) OR ST3_A_Dis1_M[3] OR ST3_A_Dis1_M[3]) AND NOT M9999;
ST3_A_Dis1_M[3] := _p41;
Out_CYw_NG1_Pick_A_H_Auto[1] := _p41;
(* Rung 4: 【Y706】NG1A(左側)チャック戻 *)
_p42 := ((ST3_A_Dis1_M[3] AND Out_CYw_NG1_Pick_A_H_Done) OR ST3_A_Dis1_M[4]) AND NOT M9999;
ST3_A_Dis1_M[4] := _p42;
Out_CYw_NG1_Chk_A_H_Auto[1] := _p42;
(* Rung 5: RC01_NG仕分け 戻 Pos *)
ST3_A_Dis1_M[5] := ((ST3_A_Dis1_M[4] AND Out_CYw_NG1_Chk_A_H_Done) OR ST3_A_Dis1_M[5]) AND NOT M9999;
END_PROGRAM

